(* IEC 61131-3 sources: plc-hackathon-2026/deliver/ME_v2_src, 24 files *)

(* ---- typeTeamAgg.st ---- *)
TYPE typeTeamAgg :
// Team energy [kWh] and cost [EUR] aggregate for one day, one month or the year.
// Names follow spec tables 12 (energies) and 4.3 (cost components). LREAL accumulators.
STRUCT
	E_fne : LREAL;                      // PV production after curtailment (FNE_P_act)
	E_fec : LREAL;                      // fixed consumption (FEC_P_fix remembered from k-1)
	E_bess_chg : LREAL;                 // battery charging, bus side
	E_bess_dch : LREAL;                 // battery discharging, bus side
	E_ev : LREAL;                       // all EV chargers, bus side
	E_ev_ch : ARRAY[0..3] OF LREAL;     // per EV charger, bus side
	E_import : LREAL;                   // grid import
	E_export : LREAL;                   // grid export
	P_peak : LREAL;                     // [kW] max 15-min import (monthly value; also kept per day for info)
	C_purchase : LREAL;                 // energy purchase = import * c_en
	C_revenue : LREAL;                  // export revenue = export * 0.9 * c_en
	C_grid : LREAL;                     // grid fee on import (VT/NT)
	C_peak : LREAL;                     // peak power cost (month/year only; 0 for days)
	C_total : LREAL;                    // purchase - revenue + grid (+ peak for month/year)
END_STRUCT
END_TYPE

(* ---- typeTeamAlarm.st ---- *)
TYPE typeTeamAlarm :
// One alarm/message history entry, stamped with SIMULATED time (no PLC clock).
STRUCT
	k : DINT;                           // simulation step when raised
	sStamp : STRING(20);                // simulated date/time "DD.MM.YYYY HH:MM"
	iCode : INT;                        // see Team_HMI alarm code list
	sText : STRING(80);                 // human readable message
END_STRUCT
END_TYPE

(* ---- Team_Cfg.st ---- *)
// Team_Cfg: team tuning constants (physics parameters are always read from SimParam).
VAR_GLOBAL CONSTANT
	N_STEPS : DINT := 35040;            // steps in the simulated year
	GRID_MARGIN_IMP : REAL := 1.0;      // [kW] safety margin below EGC_MAX_IMPORT for the predicted grid power
	GRID_MARGIN_EXP : REAL := 1.0;      // [kW] safety margin below EGC_MAX_EXPORT
	P_EPS : REAL := 0.001;              // [kW] below this a BESS setpoint is treated as zero
	// ---- forecast (FB_Forecast) ----
	FC_ALPHA_FEC : REAL := 0.5;         // EMA weight of the newest day for the load profile
	FC_ALPHA_PV : REAL := 0.3;          // EMA weight of the newest day for the PV profile
	FC_ALPHA_SIG : REAL := 0.3;         // EMA weight for the FEC deviation (sigma)
	FC_KSIG_TT : REAL := 1.0;           // two-tariff: pessimistic load = expected + FC_KSIG_TT * sigma
	FC_KSIG_DA : REAL := 0.0;           // day-ahead: same (arbitrage is worth more than the reserve)
	FC_CORR_W : INT := 4;               // intraday correction window [steps], 0 = off (max 16)
	FC_CORR_TAU : REAL := 16.0;         // fade-out of the intraday correction [steps]
	FC_CORR_FEC : BOOL := TRUE;         // apply intraday correction to FEC
	FC_CORR_PV : BOOL := TRUE;          // apply intraday correction to PV
	// ---- planner (FB_Planner) ----
	PLAN_H : INT := 96;                 // planning horizon [steps] (24 h)
	PLAN_DA_PUBLISHED : BOOL := TRUE;   // TRUE: day-ahead horizon limited to published prices (13:00 rule)
	PLAN_PEN : REAL := 20.0;            // [EUR/kW per step] penalty for planned import above the cap
	PLAN_TVF : REAL := 0.9;             // terminal value of stored energy = mean import price * PLAN_TVF
	PLAN_PVF : REAL := 0.6;             // PV share trusted when computing the peak cap
	PLAN_HI_TT : BOOL := TRUE;          // two-tariff: DP peak penalty uses the pessimistic net load
	PLAN_HI_DA : BOOL := FALSE;         // day-ahead: DP peak penalty uses the expected net load
	PLAN_TSPLIT : BOOL := FALSE;        // TRUE: free import level from the expected forecast (see FB_Planner)
	PLAN_CAPM : REAL := 1.02;           // safety factor on the computed peak cap
END_VAR

(* ---- Team_HMI.st ---- *)
// Team_HMI: everything the HMI needs that is not directly in SimIO/SimParam/SimCtrl.
// Written by FB_HmiUpdate (called from Team_Main). Only iSelDay / iSelMonth are written by the HMI.
// All times are SIMULATED time (derived from simOut.t_sim), never the PLC clock.
VAR_GLOBAL
	// ---- status / header (show on every screen) ----
	sDateTime : STRING(20);             // "DD.MM.YYYY HH:MM" start of current interval k
	k : DINT;                           // current step
	rProgressPct : REAL;                // 0..100 % of the year
	xTariffHigh : BOOL;                 // TRUE = VT (high tariff) in current interval
	sTariff : STRING(2);                // 'VT' / 'NT'
	sPriceMode : STRING(20);            // 'Dvotarifni (HEP)' / 'Dan-unaprijed'
	rPrice : REAL;                      // [EUR/kWh] energy price of the current interval
	rGridFee : REAL;                    // [EUR/kWh] grid fee of the current interval
	// ---- power flows: requested (simCmd, interval k) vs actual (*_act, interval k-1) [kW] ----
	rFneAvail : REAL;                   // available PV in interval k (before curtailment)
	rFneExpected : REAL;                // PV expected after our curtailment, interval k
	xCurtActive : BOOL;                 // curtailment enabled in interval k
	rCurtValue : REAL;                  // curtailment limit [kW]
	rFneAct : REAL;                     // actual PV, interval k-1
	rFec : REAL;                        // fixed consumption, interval k
	rFecPrev : REAL;                    // fixed consumption, interval k-1
	rBessReq : REAL;                    // requested battery power, + = discharge, - = charge
	rBessChgReq : REAL;                 // requested charge [kW] (0 if not charging)
	rBessDchReq : REAL;                 // requested discharge [kW]
	rBessAct : REAL;                    // actual battery power interval k-1, + = discharge
	rBessChgAct : REAL;
	rBessDchAct : REAL;
	aEvReq : ARRAY[0..3] OF REAL;       // requested EV power, interval k
	aEvAct : ARRAY[0..3] OF REAL;       // actual EV power, interval k-1
	rEvReqSum : REAL;
	rEvActSum : REAL;
	rGridPred : REAL;                   // predicted grid power interval k, + = import, - = export
	rImportAct : REAL;                  // measured import interval k-1
	rExportAct : REAL;                  // measured export interval k-1
	rGridPredErr : REAL;                // |prediction(k-1) - measurement(k-1)| [kW]
	rGridPredErrMax : REAL;             // max of the above since reset
	// ---- battery ----
	rSoc : REAL;                        // [%]
	rSocMin : REAL;                     // [%] safety limits (SimParam)
	rSocMax : REAL;
	sBessDir : STRING(12);              // 'PUNJENJE' / 'PRAZNJENJE' / 'MIROVANJE'
	// ---- EV chargers ----
	aEvConnected : ARRAY[0..3] OF BOOL;
	aEvDeparture : ARRAY[0..3] OF STRING(20);   // planned departure "DD.MM.YYYY HH:MM" ('' if not connected)
	aEvRemaining : ARRAY[0..3] OF REAL;         // [kWh] energy still required
	aEvDelivered : ARRAY[0..3] OF REAL;         // [kWh] delivered this session
	aEvStepsLeft : ARRAY[0..3] OF DINT;         // 15-min intervals until departure
	// ---- peak power ----
	rPeakMonth : REAL;                  // [kW] monthly import peak so far (current month)
	rPeakTarget : REAL;                 // [kW] import cap the controller currently aims for
	// ---- energy/cost tables: selection written by the HMI ----
	iSelDay : INT := 0;                 // 0..364 -> stSelDay
	iSelMonth : INT := 1;               // 1..12  -> stSelMonth, aSelMonthDays
	stSelDay : typeTeamAgg;
	stSelMonth : typeTeamAgg;
	aSelMonthDays : ARRAY[1..31] OF typeTeamAgg;   // days of the selected month (unused days = 0)
	iSelMonthDays : INT;                // number of days in the selected month
	// ---- 24 h trends: index 95 = newest interval (k-1), 0 = oldest ----
	aTrFne : ARRAY[0..95] OF REAL;      // PV actual [kW]
	aTrFec : ARRAY[0..95] OF REAL;      // fixed consumption [kW]
	aTrGrid : ARRAY[0..95] OF REAL;     // grid, + import / - export [kW]
	aTrBess : ARRAY[0..95] OF REAL;     // battery, + discharge / - charge [kW]
	aTrEv : ARRAY[0..95] OF REAL;       // EV total [kW]
	aTrSoc : ARRAY[0..95] OF REAL;      // SoC [%]
	aTrPrice : ARRAY[0..95] OF REAL;    // energy price [EUR/kWh]
	// ---- alarms ----
	xAlmImport : BOOL;                  // EGC_overload_import (previous step)
	xAlmExport : BOOL;                  // EGC_overload_export
	xAlmTripped : BOOL;                 // plant disconnected
	xAlmFinished : BOOL;                // year finished (message)
	xAlmEvUnmet : BOOL;                 // an EV left with undelivered energy (latched until reset)
	xAlmGuardEv : BOOL;                 // guard reduced EV charging to hold import limit (this step)
	xAlmGuardCurt : BOOL;               // guard curtailed PV to hold export limit (this step)
	xAlmGuardFail : BOOL;               // predicted import above limit even after all measures
	aAlarmHist : ARRAY[0..49] OF typeTeamAlarm;   // newest at index 0
	nAlarms : DINT;                     // number of messages since reset
	sLastAlarm : STRING(80);
	// ---- diagnostics ----
	nCalls : DINT;                      // Team_Main calls since PLC start
	nSteps : DINT;                      // new steps processed since reset
	nGuardEv : DINT;                    // steps with EV shedding
	nGuardCurt : DINT;                  // steps with export curtailment by the guard
	nGuardFail : DINT;                  // steps where the guard could not hold the import limit
	nBothEnables : DINT;                // must stay 0
	rEvUnmetSum : REAL;                 // [kWh] energy not delivered at departures (own estimate)
END_VAR

(* ---- Team_Log.st ---- *)
// Team_Log: daily and monthly energy/cost tables (spec 4.2/4.3). Index = simulated day / month of interval k-1.
VAR_GLOBAL
	aDay : ARRAY[0..364] OF typeTeamAgg;    // day_of_year 0..364 (C_peak = 0, C_total = purchase - revenue + grid)
	aMonth : ARRAY[1..12] OF typeTeamAgg;   // month 1..12 incl. peak power P_peak and C_peak
	stYear : typeTeamAgg;                   // yearly totals (copied to Team_Results)
END_VAR

(* ---- Team_Prices.st ---- *)
// Team_Prices: price lists (cjenici, spec 3.9/4.1) generated by tools/gen_prices.py from the organizer CSVs.
// Energy price only; grid fee and peak price come from SimParam. Not a simulator profile (FNE/FEC/EV are never embedded).
VAR_GLOBAL CONSTANT
	// Elektra two-tariff energy price [EUR/kWh] per calendar quarter (1 = Jan-Mar ... 4 = Oct-Dec)
	TT_NT : ARRAY[1..4] OF REAL := [0.09, 0.1051, 0.0934, 0.0949];
	TT_VT : ARRAY[1..4] OF REAL := [0.1531, 0.1786, 0.1588, 0.1613];
END_VAR
VAR_GLOBAL
	// Day-ahead energy price [EUR/kWh] per 15-min interval k = 0..35039 (ENTSO-E HR 2025, may be negative)
	aDA : ARRAY[0..35039] OF REAL := [
		4(0.1353348), 4(0.143694), 4(0.1349352), 4(0.1010124), 4(0.0687852), 4(0.1011852), 4(0.0974808), 4(0.0902556), 4(0.0399492), 4(0.0485892), 4(0.04158), 4(0.0430056),
		4(0.04347), 4(0.059886), 4(0.0664632), 4(0.0900288), 4(0.1161648), 4(0.1328832), 4(0.1382724), 4(0.1446984), 4(0.1406268), 4(0.1307124), 4(0.1310364), 4(0.0904176),
		4(0.0689904), 4(0.0865296), 4(0.0846936), 4(0.053136), 4(0.0614844), 4(0.0834732), 4(0.1200204), 4(0.1431324), 4(0.1405836), 4(0.1433268), 4(0.1391148), 4(0.1337364),
		4(0.1330668), 4(0.126144), 4(0.135), 4(0.1405188), 4(0.1650456), 4(0.1762452), 4(0.1695492), 4(0.1646028), 4(0.1414152), 4(0.134622), 4(0.1270188), 4(0.1095228),
		4(0.111996), 4(0.1023732), 4(0.0968436), 4(0.0945216), 4(0.0923832), 4(0.0993816), 4(0.1185516), 4(0.1469556), 4(0.1492452), 4(0.1461564), 4(0.1350216), 4(0.1219968),
		4(0.1201716), 4(0.118206), 4(0.124956), 4(0.1402596), 4(0.1587276), 4(0.1571508), 4(0.1572696), 4(0.1564488), 4(0.1478196), 4(0.1314684), 4(0.1361988), 4(0.1318572),
		4(0.1189296), 4(0.1130112), 4(0.1087344), 4(0.1065204), 4(0.1077732), 4(0.113454), 4(0.12096), 4(0.1352808), 4(0.1386612), 4(0.14121), 4(0.1407672), 4(0.1385532),
		4(0.1404324), 4(0.140238), 4(0.147312), 4(0.15309), 4(0.1819368), 4(0.1857924), 4(0.1848096), 4(0.1831572), 4(0.1590624), 4(0.151524), 4(0.1455192), 4(0.1259604),
		4(0.1211004), 4(0.107838), 4(0.1033668), 4(0.1013364), 4(0.1006992), 4(0.0971892), 4(0.0989064), 4(0.1068012), 4(0.105408), 4(0.1070172), 4(0.103194), 4(0.1084104),
		4(0.1057752), 4(0.1129248), 4(0.122094), 4(0.1337364), 4(0.1717308), 4(0.165024), 4(0.1562328), 4(0.1627236), 4(0.1535328), 4(0.1449144), 4(0.1105056), 4(0.0771984),
		4(0.1130004), 4(0.0960336), 4(0.0743256), 4(0.0708804), 4(0.070794), 4(0.0962172), 4(0.1229364), 4(0.1331748), 4(0.1334664), 4(0.1152576), 4(0.097956), 4(0.0780624),
		4(0.0841212), 4(0.10476), 4(0.1249668), 4(0.1229904), 4(0.1472904), 4(0.1600344), 4(0.1528524), 4(0.1521828), 4(0.1456272), 4(0.122364), 4(0.1168128), 4(0.0853416),
		4(0.0343116), 4(0.056538), 4(0.0510192), 4(0.0135), 4(0.0662688), 4(0.0844668), 4(0.1362636), 4(0.16443), 4(0.148014), 4(0.1423224), 4(0.1318248), 4(0.131274),
		4(0.1322676), 4(0.1404432), 4(0.1504656), 4(0.1588572), 4(0.1668384), 4(0.166806), 4(0.1628424), 4(0.1643328), 4(0.1532088), 4(0.1370196), 4(0.125064), 4(0.1204416),
		4(0.0901584), 4(0.0813672), 4(0.0789048), 4(0.0747036), 4(0.0923076), 4(0.11178), 4(0.1367388), 4(0.1635336), 4(0.1611252), 4(0.1341576), 4(0.1174068), 4(0.1103436),
		4(0.1120824), 4(0.1245996), 4(0.1353132), 4(0.1550556), 4(0.1646784), 4(0.165456), 4(0.1622916), 4(0.1614384), 4(0.1484352), 4(0.1356372), 4(0.1255716), 4(0.114588),
		4(0.1147284), 4(0.114588), 4(0.1119096), 4(0.1104408), 4(0.1152468), 4(0.1184868), 4(0.1342656), 4(0.1542132), 4(0.1678104), 4(0.1601208), 4(0.1514916), 4(0.1435644),
		4(0.1331532), 4(0.1284012), 4(0.1325484), 4(0.1425708), 4(0.1583496), 4(0.1566756), 4(0.16065), 4(0.1521612), 4(0.1421172), 4(0.1240056), 4(0.11151), 4(0.0968328),
		4(0.0941976), 4(0.0868104), 4(0.0826092), 4(0.0808164), 4(0.0767664), 4(0.1046088), 4(0.1354968), 4(0.165024), 4(0.1680264), 4(0.1522368), 4(0.1334556), 4(0.1226772),
		4(0.1160244), 4(0.1134108), 4(0.1188108), 4(0.1389852), 4(0.1609308), 4(0.1583604), 4(0.1590084), 4(0.1569024), 4(0.1457568), 4(0.1323108), 4(0.129492), 4(0.1226016),
		4(0.1179468), 4(0.1079676), 4(0.1042632), 4(0.1000296), 4(0.099144), 4(0.1006236), 4(0.1021788), 4(0.1209168), 4(0.12312), 4(0.1200744), 4(0.113454), 4(0.1078488),
		4(0.1046088), 4(0.100602), 4(0.1068768), 4(0.113994), 4(0.1448928), 4(0.1509732), 4(0.1472256), 4(0.148284), 4(0.1366848), 4(0.1265328), 4(0.11799), 4(0.1143612),
		4(0.1075896), 4(0.0961416), 4(0.0964548), 4(0.092178), 4(0.0918), 4(0.0919188), 4(0.0946836), 4(0.10989), 4(0.1258092), 4(0.1296756), 4(0.1271916), 4(0.1140588),
		4(0.1112292), 4(0.1075788), 4(0.1139616), 4(0.1299564), 4(0.1461024), 4(0.1542564), 4(0.1583928), 4(0.1557468), 4(0.1468152), 4(0.1380348), 4(0.1312956), 4(0.124092),
		4(0.1213812), 4(0.1134756), 4(0.1128168), 4(0.1083996), 4(0.108), 4(0.1190052), 4(0.1512108), 4(0.1927476), 4(0.2371032), 4(0.1868184), 4(0.15201), 4(0.1311444),
		4(0.1245456), 4(0.1297512), 4(0.1363284), 4(0.1529928), 4(0.1704564), 4(0.1678212), 4(0.16902), 4(0.1670976), 4(0.1538244), 4(0.1375164), 4(0.1288008), 4(0.1167588),
		4(0.1186812), 4(0.115344), 4(0.1107), 4(0.1092312), 4(0.1125036), 4(0.1180332), 4(0.1495908), 4(0.1742688), 4(0.2001672), 4(0.16416), 4(0.141156), 4(0.1340712),
		4(0.1289304), 4(0.1293084), 4(0.1439532), 4(0.1770552), 4(0.1979964), 4(0.2446632), 4(0.239652), 4(0.211572), 4(0.187164), 4(0.172746), 4(0.1610172), 4(0.1348812),
		4(0.127656), 4(0.1213488), 4(0.1200528), 4(0.1174932), 4(0.1255068), 4(0.1390392), 4(0.1600992), 4(0.2120148), 4(0.3359124), 4(0.338904), 4(0.3266568), 4(0.325566),
		4(0.31023), 4(0.306774), 4(0.3062448), 4(0.3319596), 4(0.326268), 4(0.368226), 4(0.320328), 4(0.265248), 4(0.1937088), 4(0.1670328), 4(0.1554768), 4(0.133812),
		4(0.136296), 4(0.131868), 4(0.1281636), 4(0.1259928), 4(0.1292652), 4(0.1392012), 4(0.1701216), 4(0.2121984), 4(0.2210544), 4(0.189), 4(0.164052), 4(0.1518912),
		4(0.1456488), 4(0.1492344), 4(0.1566), 4(0.1827144), 4(0.19683), 4(0.2082348), 4(0.1990656), 4(0.1943676), 4(0.172368), 4(0.1623996), 4(0.1519992), 4(0.1398276),
		4(0.1364364), 4(0.1331208), 4(0.1297836), 4(0.1277532), 4(0.1277964), 4(0.1346328), 4(0.152064), 4(0.1890108), 4(0.2247804), 4(0.1893672), 4(0.1700352), 4(0.1518696),
		4(0.1365552), 4(0.1339524), 4(0.1444284), 4(0.1637172), 4(0.1839888), 4(0.1930284), 4(0.1943136), 4(0.1881576), 4(0.1705428), 4(0.1566), 4(0.1511676), 4(0.1383588),
		4(0.1363392), 4(0.1309284), 4(0.1311336), 4(0.128412), 4(0.1263816), 4(0.1294164), 4(0.1325592), 4(0.1465776), 4(0.157626), 4(0.155628), 4(0.1445796), 4(0.1315224),
		4(0.1283796), 4(0.1242108), 4(0.129168), 4(0.149094), 4(0.1772712), 4(0.1826928), 4(0.1809756), 4(0.181278), 4(0.1686096), 4(0.1548936), 4(0.147312), 4(0.1397088),
		4(0.1403028), 4(0.1350108), 4(0.1336068), 4(0.1309392), 4(0.1297944), 4(0.1296), 4(0.1314252), 4(0.1340172), 4(0.1335636), 4(0.136188), 4(0.1366092), 4(0.1341252),
		4(0.12123), 4(0.1161108), 4(0.1261548), 4(0.1377324), 4(0.1627344), 4(0.1759428), 4(0.180522), 4(0.1794096), 4(0.1741608), 4(0.1651644), 4(0.145044), 4(0.133866),
		4(0.1322784), 4(0.1294056), 4(0.1259388), 4(0.1235628), 4(0.124686), 4(0.1404216), 4(0.1766232), 4(0.3070548), 4(0.4670028), 4(0.3149496), 4(0.2551932), 4(0.2076084),
		4(0.193266), 4(0.1851012), 4(0.2071332), 4(0.2981016), 4(0.446472), 4(0.6208812), 4(0.5111424), 4(0.3192156), 4(0.2376), 4(0.1836), 4(0.1718928), 4(0.1540944),
		4(0.1477764), 4(0.1417932), 4(0.134622), 4(0.1350972), 4(0.1429056), 4(0.16416), 4(0.207414), 4(0.3141612), 4(0.4177224), 4(0.2861676), 4(0.2540484), 4(0.2179224),
		4(0.2129004), 4(0.1951344), 4(0.2188512), 4(0.3057588), 4(0.245214), 4(0.3387744), 4(0.2779704), 4(0.2207844), 4(0.190728), 4(0.1687392), 4(0.153684), 4(0.144234),
		4(0.141588), 4(0.1360152), 4(0.1345896), 4(0.1350972), 4(0.1372464), 4(0.1506816), 4(0.20925), 4(0.3410964), 4(0.2672136), 4(0.2153628), 4(0.1933848), 4(0.1867752),
		4(0.1782), 4(0.1836), 4(0.1943136), 4(0.2137752), 4(0.2703888), 4(0.276102), 4(0.2261952), 4(0.222642), 4(0.2220156), 4(0.1710072), 4(0.1589436), 4(0.145854),
		4(0.1353888), 4(0.1299564), 4(0.119394), 4(0.1175796), 4(0.1227096), 4(0.1344708), 4(0.1809864), 4(0.2092608), 4(0.1881684), 4(0.1808568), 4(0.1625292), 4(0.1594728),
		4(0.1543104), 4(0.1588032), 4(0.1690416), 4(0.1919376), 4(0.2108916), 4(0.2148012), 4(0.2028672), 4(0.1957824), 4(0.2018628), 4(0.1633608), 4(0.1606176), 4(0.136188),
		4(0.127656), 4(0.1162512), 4(0.1107), 4(0.1093392), 4(0.1170288), 4(0.1424304), 4(0.17469), 4(0.1909872), 4(0.1764828), 4(0.1599048), 4(0.1535652), 4(0.1422576),
		4(0.1392444), 4(0.13662), 4(0.1417716), 4(0.161892), 4(0.1961064), 4(0.1983744), 4(0.1922616), 4(0.1883412), 4(0.1774872), 4(0.1666008), 4(0.1547208), 4(0.1429488),
		4(0.1203336), 4(0.1117476), 4(0.0980856), 4(0.094878), 4(0.0971136), 4(0.1055808), 4(0.1218564), 4(0.1337904), 4(0.1181628), 4(0.1153224), 4(0.1033776), 4(0.0975888),
		4(0.09396), 4(0.0924372), 4(0.1067256), 4(0.1288872), 4(0.1661148), 4(0.1701108), 4(0.1716444), 4(0.1709208), 4(0.162864), 4(0.155574), 4(0.1481004), 4(0.135),
		4(0.1419552), 4(0.1297404), 4(0.1272888), 4(0.1204524), 4(0.12096), 4(0.1231524), 4(0.1255176), 4(0.1334664), 4(0.1427112), 4(0.1400004), 4(0.1207656), 4(0.112752),
		4(0.1054188), 4(0.1028808), 4(0.1209168), 4(0.13095), 4(0.1467288), 4(0.1559088), 4(0.1424628), 4(0.1443312), 4(0.1348812), 4(0.1245888), 4(0.104004), 4(0.08397),
		4(0.0654696), 4(0.0605124), 4(0.0433404), 4(0.032022), 4(0.0490536), 4(0.118098), 4(0.1559088), 4(0.187002), 4(0.1719684), 4(0.1409616), 4(0.1084428), 4(0.1040148),
		4(0.0946944), 4(0.1125792), 4(0.1399464), 4(0.1582416), 4(0.1937628), 4(0.1899936), 4(0.1928124), 4(0.1906308), 4(0.170856), 4(0.1461024), 4(0.130626), 4(0.106056),
		4(0.106758), 4(0.0855684), 4(0.0941112), 4(0.0877068), 4(0.0877392), 4(0.122688), 4(0.1498608), 4(0.1502712), 4(0.1519992), 4(0.1354212), 4(0.141318), 4(0.1357344),
		4(0.1322892), 4(0.1372788), 4(0.1420632), 4(0.135162), 4(0.1540296), 4(0.1559304), 4(0.1593864), 4(0.1502928), 4(0.1499256), 4(0.1251612), 4(0.1250208), 4(0.1051704),
		4(0.105462), 4(0.097362), 4(0.0910332), 4(0.0914328), 4(0.0972), 4(0.1214676), 4(0.154656), 4(0.1773468), 4(0.1579068), 4(0.1480896), 4(0.1204308), 4(0.1014444),
		4(0.093204), 4(0.0935496), 4(0.1055484), 4(0.1400328), 4(0.1792692), 4(0.1827792), 4(0.1721088), 4(0.173502), 4(0.1609524), 4(0.1491912), 4(0.1330236), 4(0.1119204),
		4(0.110268), 4(0.1095228), 4(0.1069524), 4(0.1100844), 4(0.1098036), 4(0.1232496), 4(0.1569348), 4(0.1669788), 4(0.173124), 4(0.1639764), 4(0.1429704), 4(0.13311),
		4(0.1219428), 4(0.122364), 4(0.1403892), 4(0.1655748), 4(0.1736748), 4(0.1896696), 4(0.1858032), 4(0.1741824), 4(0.1635228), 4(0.145908), 4(0.1370952), 4(0.129816),
		4(0.1296), 4(0.1269), 4(0.1232064), 4(0.1236384), 4(0.1267164), 4(0.1316088), 4(0.1604556), 4(0.1728), 4(0.176796), 4(0.1672056), 4(0.140508), 4(0.136296),
		4(0.1296648), 4(0.1308852), 4(0.1296432), 4(0.1655964), 4(0.1810512), 4(0.1930716), 4(0.1992384), 4(0.1933092), 4(0.1756728), 4(0.164916), 4(0.1607472), 4(0.144126),
		4(0.1494828), 4(0.1409724), 4(0.135108), 4(0.1288332), 4(0.1295568), 4(0.1312308), 4(0.1374948), 4(0.1563192), 4(0.1657368), 4(0.1538352), 4(0.138672), 4(0.1296864),
		4(0.1191132), 4(0.111672), 4(0.122796), 4(0.1411344), 4(0.1683072), 4(0.1792368), 4(0.180036), 4(0.1760184), 4(0.169128), 4(0.1568592), 4(0.1530684), 4(0.1422792),
		4(0.1439208), 4(0.1370628), 4(0.1328292), 4(0.1303128), 4(0.1321272), 4(0.1332828), 4(0.1383372), 4(0.146772), 4(0.148284), 4(0.148716), 4(0.1404432), 4(0.1396764),
		4(0.1320192), 4(0.1208304), 4(0.1263168), 4(0.140562), 4(0.168156), 4(0.1802088), 4(0.185544), 4(0.187866), 4(0.17874), 4(0.1682316), 4(0.1603152), 4(0.1438992),
		4(0.1399032), 4(0.1367604), 4(0.1346976), 4(0.1296432), 4(0.1330992), 4(0.1379916), 4(0.1719144), 4(0.2245104), 4(0.2626884), 4(0.1922832), 4(0.161946), 4(0.1363176),
		4(0.1266516), 4(0.1249776), 4(0.1344276), 4(0.1597968), 4(0.1793664), 4(0.226962), 4(0.2167884), 4(0.217188), 4(0.1811592), 4(0.16524), 4(0.1557252), 4(0.1466748),
		4(0.142992), 4(0.1355832), 4(0.1330344), 4(0.1339092), 4(0.13311), 4(0.1378404), 4(0.1674432), 4(0.2056644), 4(0.2289492), 4(0.1763748), 4(0.1474524), 4(0.1369656),
		4(0.127602), 4(0.1222452), 4(0.1296972), 4(0.1542456), 4(0.181332), 4(0.189324), 4(0.189), 4(0.1863648), 4(0.1727352), 4(0.1464804), 4(0.1424412), 4(0.1347624),
		4(0.1260036), 4(0.1207548), 4(0.1198584), 4(0.1186056), 4(0.1248912), 4(0.1323648), 4(0.1636524), 4(0.1825092), 4(0.1952748), 4(0.1720764), 4(0.145476), 4(0.133704),
		4(0.127926), 4(0.1297512), 4(0.139158), 4(0.1556496), 4(0.1719252), 4(0.19116), 4(0.205092), 4(0.2048004), 4(0.1836), 4(0.1678536), 4(0.155196), 4(0.144774),
		4(0.1443636), 4(0.1403892), 4(0.13608), 4(0.135), 4(0.1350108), 4(0.1447524), 4(0.165996), 4(0.1944972), 4(0.2356128), 4(0.1930932), 4(0.1686204), 4(0.1617408),
		4(0.1561032), 4(0.1526148), 4(0.1520208), 4(0.1622808), 4(0.181656), 4(0.188244), 4(0.1913544), 4(0.1864512), 4(0.1768068), 4(0.159624), 4(0.1512108), 4(0.131706),
		4(0.136134), 4(0.121716), 4(0.1175256), 4(0.1134), 4(0.1185192), 4(0.1280772), 4(0.1678104), 4(0.1848744), 4(0.1782324), 4(0.1625076), 4(0.1456812), 4(0.1280556),
		4(0.1243512), 4(0.1240164), 4(0.12744), 4(0.1442556), 4(0.1857924), 4(0.1894644), 4(0.1884924), 4(0.1860624), 4(0.1818072), 4(0.1557576), 4(0.1285632), 4(0.1209816),
		4(0.09828), 4(0.0950184), 4(0.0937872), 4(0.09612), 4(0.0968652), 4(0.0982692), 4(0.1052028), 4(0.1174068), 4(0.1222128), 4(0.109134), 4(0.1035072), 4(0.0960336),
		4(0.0954828), 4(0.097686), 4(0.1025244), 4(0.12744), 4(0.16173), 4(0.1752948), 4(0.1733832), 4(0.1713852), 4(0.1661472), 4(0.16092), 4(0.1542564), 4(0.1449792),
		4(0.1458), 4(0.136404), 4(0.1319004), 4(0.128844), 4(0.1261656), 8(0.12636), 4(0.1441044), 4(0.1477116), 4(0.1321812), 4(0.1230876), 4(0.1191456), 4(0.1106028),
		4(0.1090368), 4(0.118692), 4(0.130032), 4(0.1627992), 4(0.1736856), 4(0.1889784), 4(0.1888164), 4(0.1786968), 4(0.1560816), 4(0.15444), 4(0.139482), 4(0.1297944),
		4(0.1247292), 4(0.1217916), 4(0.1173096), 4(0.1168992), 4(0.126576), 4(0.1724004), 4(0.1935684), 4(0.1958688), 4(0.1762344), 4(0.1672488), 4(0.1512108), 4(0.136512),
		4(0.132732), 4(0.142398), 4(0.179712), 4(0.2052972), 4(0.218322), 4(0.2210112), 4(0.2083752), 4(0.2056644), 4(0.1809), 4(0.1751544), 4(0.1435428), 4(0.1483812),
		4(0.1365768), 4(0.1335204), 4(0.1290384), 4(0.1365876), 4(0.1763856), 4(0.1951884), 4(0.2572236), 4(0.1924884), 4(0.15687), 4(0.13068), 4(0.1269432), 4(0.1278612),
		4(0.1289304), 4(0.1395684), 4(0.1727136), 4(0.200016), 4(0.2052), 4(0.2388312), 4(0.2170044), 4(0.1934064), 4(0.1859868), 4(0.1727892), 4(0.1431432), 4(0.1397952),
		4(0.1380996), 4(0.1369656), 4(0.1367172), 4(0.1390392), 4(0.1469772), 4(0.1866024), 4(0.1955232), 4(0.1944), 4(0.1889136), 4(0.1791612), 4(0.171234), 4(0.16119),
		4(0.1638144), 4(0.1802196), 4(0.1956852), 4(0.2190564), 4(0.3030804), 4(0.2873556), 4(0.240462), 4(0.2384316), 4(0.1923156), 4(0.1861812), 4(0.1728), 4(0.1722708),
		4(0.161298), 4(0.158868), 4(0.1538136), 4(0.1591596), 4(0.1767852), 4(0.2259684), 4(0.421524), 4(0.3348108), 4(0.2808108), 4(0.2247588), 4(0.2027268), 4(0.2015604),
		4(0.2252664), 4(0.2457648), 4(0.2673), 4(0.2891484), 4(0.2678184), 4(0.2236788), 4(0.2122416), 4(0.1927152), 4(0.1759536), 4(0.1653696), 4(0.1503036), 4(0.1514376),
		4(0.1460916), 4(0.141048), 4(0.1412748), 4(0.141858), 4(0.1520748), 4(0.1772712), 4(0.2337336), 4(0.2835216), 4(0.229284), 4(0.1935144), 4(0.1778976), 4(0.1623564),
		4(0.1625508), 4(0.1714824), 4(0.1871316), 4(0.2142396), 4(0.3135456), 4(0.3104244), 4(0.2420388), 4(0.198234), 4(0.1766232), 4(0.16524), 4(0.1512324), 4(0.1472688),
		4(0.1418796), 4(0.1303884), 4(0.1291356), 4(0.1295784), 4(0.1315872), 4(0.146718), 4(0.1623888), 4(0.1616328), 4(0.148068), 4(0.1345572), 4(0.1278288), 4(0.1213812),
		4(0.1188108), 4(0.126252), 4(0.1413936), 4(0.1687716), 4(0.1905552), 4(0.1925856), 4(0.1880064), 4(0.1818504), 4(0.165348), 4(0.1515672), 4(0.1441692), 4(0.1448388),
		4(0.139212), 4(0.1334556), 4(0.129492), 4(0.1291356), 4(0.1305612), 4(0.133758), 4(0.1448712), 4(0.153846), 4(0.152334), 4(0.1427652), 4(0.141696), 4(0.1389636),
		4(0.1375812), 4(0.14094), 4(0.1524744), 4(0.174852), 4(0.1890324), 4(0.191322), 4(0.1876932), 4(0.1830708), 4(0.1726272), 4(0.1613412), 4(0.1420308), 4(0.1431216),
		4(0.1307448), 4(0.1299672), 4(0.1365876), 4(0.1406052), 4(0.1550124), 4(0.1884924), 4(0.2253096), 4(0.2265732), 4(0.185004), 4(0.1508436), 4(0.1288764), 4(0.1232928),
		4(0.1176012), 4(0.13176), 4(0.1601748), 4(0.1869372), 4(0.238572), 4(0.2883816), 4(0.2338956), 4(0.1934928), 4(0.1759212), 4(0.169074), 4(0.15444), 4(0.146664),
		4(0.1429488), 4(0.1358748), 4(0.1331316), 4(0.1377216), 4(0.163998), 4(0.2263032), 4(0.3576096), 4(0.209304), 4(0.1750356), 4(0.154386), 4(0.1445148), 4(0.142398),
		4(0.1559736), 4(0.1631448), 4(0.1770876), 4(0.3453516), 4(0.2810268), 4(0.2770092), 4(0.2601612), 4(0.1939248), 4(0.1817316), 4(0.1740852), 4(0.1480032), 4(0.14121),
		4(0.1392768), 4(0.1372896), 4(0.136458), 4(0.1398168), 4(0.155088), 4(0.1828872), 4(0.218592), 4(0.190404), 4(0.165456), 4(0.123606), 4(0.1240056), 4(0.1162728),
		4(0.1160568), 4(0.126954), 4(0.1515888), 4(0.190944), 4(0.249534), 4(0.2520504), 4(0.2164968), 4(0.1938492), 4(0.1805868), 4(0.1764936), 4(0.1671192), 4(0.1350972),
		4(0.1303452), 4(0.1251936), 4(0.1203984), 4(0.1305396), 4(0.1563948), 4(0.2001456), 4(0.263412), 4(0.19062), 4(0.1302804), 4(0.1142748), 4(0.0986364), 4(0.1005588),
		4(0.1060236), 4(0.1154952), 4(0.153846), 4(0.1964844), 4(0.2781972), 4(0.3032856), 4(0.2709936), 4(0.187596), 4(0.176904), 4(0.1739556), 4(0.1439748), 4(0.1269432),
		4(0.1223964), 4(0.1204956), 4(0.1224288), 4(0.1231308), 4(0.1458), 4(0.1756512), 4(0.188244), 4(0.1582416), 4(0.1398276), 4(0.1123524), 4(0.0950508), 4(0.0867564),
		4(0.0860436), 4(0.107892), 4(0.1171476), 4(0.1718604), 4(0.2034612), 4(0.2067012), 4(0.2070792), 4(0.1797876), 4(0.1654884), 4(0.145422), 4(0.1260468), 4(0.13203),
		4(0.1259496), 4(0.1227312), 4(0.1168668), 4(0.1191024), 4(0.1260468), 4(0.151794), 4(0.1414152), 4(0.1065204), 4(0.0763344), 4(0.0634392), 4(0.0612036), 4(0.0569916),
		4(0.0606852), 4(0.0737316), 4(0.128358), 4(0.1802304), 4(0.2145528), 4(0.1995408), 4(0.2117664), 4(0.1919808), 4(0.1703268), 4(0.1657152), 4(0.1615464), 4(0.1378512),
		4(0.138294), 4(0.1283796), 4(0.1277748), 4(0.128736), 4(0.1349352), 4(0.1454112), 4(0.1423332), 4(0.1270296), 4(0.1109592), 4(0.0945432), 4(0.0962172), 4(0.0814752),
		4(0.080838), 4(0.1136808), 4(0.1515996), 4(0.20547), 4(0.2142504), 4(0.2108916), 4(0.2121984), 4(0.1816344), 4(0.1752408), 4(0.1579716), 4(0.1437696), 4(0.1412748),
		4(0.1266408), 4(0.1217808), 4(0.1202796), 4(0.12393), 4(0.1646784), 4(0.2244888), 4(0.2619324), 4(0.1898856), 4(0.17928), 4(0.1571292), 4(0.1439964), 4(0.1381104),
		4(0.1377216), 4(0.1576908), 4(0.2053944), 4(0.2542212), 4(0.3007044), 4(0.3385584), 4(0.314172), 4(0.2235384), 4(0.1914516), 4(0.1759428), 4(0.1442664), 4(0.154332),
		4(0.139428), 4(0.1344168), 4(0.1337688), 4(0.1378404), 4(0.1590192), 4(0.2322324), 4(0.2833596), 4(0.1877148), 4(0.1683828), 4(0.1544076), 4(0.139374), 4(0.1379268),
		4(0.140346), 4(0.1505088), 4(0.1666008), 4(0.2288196), 4(0.3069468), 4(0.3333636), 4(0.2880468), 4(0.2162916), 4(0.1727892), 4(0.1578528), 4(0.1416744), 4(0.1348488),
		4(0.1326132), 4(0.1286388), 4(0.1282284), 4(0.1286172), 4(0.1369332), 4(0.1886328), 4(0.2148444), 4(0.1917864), 4(0.1698516), 4(0.1571292), 4(0.1430892), 4(0.13122),
		4(0.1323864), 4(0.1405836), 4(0.1608552), 4(0.1918404), 4(0.2159892), 4(0.2162052), 4(0.1993896), 4(0.1851768), 4(0.1579716), 4(0.1453248), 4(0.129816), 4(0.1205928),
		4(0.1121148), 4(0.1109268), 8(0.1096308), 4(0.1193508), 4(0.158328), 4(0.1742148), 4(0.1794096), 4(0.1623456), 4(0.1463184), 4(0.1380024), 4(0.130626), 4(0.1261872),
		4(0.1297512), 4(0.1470096), 4(0.181764), 4(0.1843668), 4(0.1918836), 4(0.1853712), 4(0.1789992), 4(0.1529928), 4(0.1429056), 4(0.1239732), 4(0.1306044), 4(0.1193832),
		4(0.1181304), 4(0.1156464), 4(0.1216944), 4(0.13392), 4(0.1674648), 4(0.1978236), 4(0.1741608), 4(0.1593324), 4(0.1399248), 4(0.1272024), 4(0.1191888), 4(0.1188972),
		4(0.1216944), 4(0.1370952), 4(0.1721628), 4(0.2049408), 4(0.2110428), 4(0.2149308), 4(0.1967652), 4(0.1700352), 4(0.1497528), 4(0.134946), 4(0.1395468), 4(0.130464),
		4(0.1266948), 4(0.1222884), 4(0.1193616), 4(0.1248264), 4(0.1381212), 4(0.1493208), 4(0.1511892), 4(0.1508868), 4(0.138024), 4(0.12393), 4(0.1121904), 4(0.1080648),
		4(0.1125252), 4(0.1363068), 4(0.1677024), 4(0.21735), 4(0.2160972), 4(0.2048868), 4(0.173556), 4(0.1505412), 4(0.1351188), 4(0.1295136), 4(0.1363176), 4(0.1292436),
		4(0.1137132), 4(0.113724), 4(0.1215432), 4(0.1246428), 4(0.1444932), 4(0.1420956), 4(0.120906), 4(0.09612), 4(0.073764), 4(0.05292), 4(0.0297), 4(0.019008),
		4(0.0572184), 4(0.0780732), 4(0.1435644), 4(0.1693332), 4(0.176526), 4(0.1771632), 4(0.1706292), 4(0.1626372), 4(0.1358316), 4(0.1227204), 4(0.1238328), 4(0.1172664),
		4(0.115668), 4(0.1113588), 4(0.1151604), 4(0.1288332), 4(0.1513188), 4(0.17604), 4(0.1595484), 4(0.1176444), 4(0.0878364), 4(0.084618), 4(0.091476), 4(0.0626184),
		4(0.0921672), 4(0.1216296), 4(0.152766), 4(0.1925964), 4(0.2588436), 4(0.2024784), 4(0.1784916), 4(0.1745604), 4(0.1605204), 4(0.1555308), 4(0.1387368), 4(0.1302264),
		4(0.1188756), 4(0.1167696), 4(0.1265112), 4(0.1686852), 4(0.1939896), 4(0.1906956), 4(0.153306), 4(0.1248804), 4(0.103302), 4(0.1115964), 4(0.039798), 4(0.0315252),
		4(0.0721656), 4(0.1109484), 4(0.1677996), 4(0.2093148), 4(0.2734452), 4(0.215298), 4(0.1860192), 4(0.1675188), 4(0.1552824), 4(0.1442556), 4(0.1448064), 4(0.1312524),
		4(0.1238328), 4(0.118854), 4(0.1313712), 4(0.1473228), 4(0.18387), 4(0.163944), 4(0.1172124), 4(0.0805248), 4(0.0244836), 4(0.0119124), 4(0.0075924), 4(0.0011232),
		4(0.0041688), 4(0.0786888), 4(0.134892), 4(0.1743768), 4(0.228744), 4(0.1930392), 4(0.1734264), 4(0.1610604), 4(0.1397736), 4(0.1315116), 4(0.1128816), 4(0.1133676),
		4(0.1125792), 4(0.1146852), 4(0.1219968), 4(0.1468692), 4(0.1857276), 4(0.1662336), 4(0.11718), 4(0.086076), 4(0.0622944), 4(0.0057564), 4(0.0016632), 4(0.0007776),
		4(0.0142128), 4(0.0805788), 4(0.1324512), 4(0.2071116), 4(0.237006), 4(0.2223612), 4(0.1900692), 4(0.1577772), 4(0.1492776), 4(0.1302912), 4(0.1153116), 4(0.1140264),
		4(0.10854), 4(0.1099656), 4(0.114048), 4(0.1347624), 4(0.164322), 4(0.1642896), 4(0.1339956), 4(0.0899316), 4(0.071064), 4(0.0343548), 4(0.0138132), 4(0.0086508),
		4(0.0415476), 4(0.1037232), 4(0.1464804), 4(0.1729836), 4(0.2413584), 4(0.208764), 4(0.175068), 4(0.151524), 4(0.140994), 4(0.1352808), 4(0.1441908), 4(0.13662),
		4(0.1405512), 4(0.137808), 4(0.1404756), 4(0.1484568), 4(0.146016), 4(0.1347948), 4(0.1058832), 4(0.0783432), 4(0.019494), 4(0.00243), 4(0.000864), 4(4.32E-05),
		4(7.56E-05), 4(0.0650916), 4(0.1236708), 4(0.1769364), 4(0.2254716), 4(0.2034612), 4(0.166914), 4(0.154116), 4(0.1454112), 4(0.1249884), 4(0.1188108), 4(0.115452),
		4(0.1132056), 4(0.1155276), 4(0.1188864), 4(0.121716), 4(0.1188324), 4(0.106218), 4(0.0736344), 4(0.0316116), 4(0.010908), 4(0.0016416), 4(0.000702), 4(-0.0003456),
		4(0.0007884), 4(0.0187812), 4(0.1079352), 4(0.149796), 4(0.1598832), 4(0.158166), 4(0.148824), 4(0.1400328), 4(0.125334), 4(0.119502), 4(0.10692), 4(0.105948),
		4(0.1073304), 4(0.1075032), 4(0.107838), 4(0.1214136), 4(0.1614492), 4(0.1707372), 4(0.144612), 4(0.1070604), 4(0.0843588), 4(0.0798876), 4(0.0821016), 4(0.0835056),
		4(0.0917568), 4(0.1085508), 4(0.1429704), 4(0.1568592), 4(0.1869804), 4(0.171828), 4(0.1521828), 4(0.1384992), 4(0.1163376), 4(0.1065528), 4(0.114426), 4(0.1117476),
		4(0.1086804), 4(0.1099332), 4(0.1132272), 4(0.1220832), 4(0.1521828), 4(0.1583064), 4(0.1551744), 4(0.1403568), 4(0.1103544), 4(0.1058724), 4(0.1052568), 4(0.1080432),
		4(0.1128168), 4(0.1251504), 4(0.1503792), 4(0.1712016), 4(0.205632), 4(0.1912248), 4(0.1594512), 4(0.1449036), 4(0.1326996), 4(0.1161864), 4(0.1102356), 4(0.1087776),
		4(0.1059912), 4(0.1063044), 4(0.1118664), 4(0.122418), 4(0.1487052), 4(0.1657152), 4(0.1566972), 4(0.135), 4(0.110376), 4(0.1075248), 4(0.1059048), 4(0.1074924),
		4(0.1098576), 4(0.1288764), 4(0.1465776), 4(0.1611252), 4(0.205578), 4(0.1930068), 4(0.1576692), 4(0.142776), 4(0.1296), 4(0.1187028), 4(0.1152576), 4(0.0640764),
		4(0.0236844), 4(0.0324216), 4(0.0692064), 4(0.1137564), 4(0.1436292), 4(0.1567836), 4(0.141912), 4(0.1055592), 4(0.1039932), 4(0.0934092), 4(0.0904392), 4(0.0753192),
		4(0.094176), 4(0.11664), 4(0.1324296), 4(0.1532628), 4(0.179334), 4(0.1873476), 4(0.16092), 4(0.1465452), 4(0.1107216), 4(0.1079028), 4(0.1178172), 4(0.11448),
		4(0.114372), 4(0.1121364), 4(0.113724), 4(0.1232928), 4(0.1544832), 4(0.164646), 4(0.1372248), 4(0.1197936), 4(0.098928), 4(0.0945216), 4(0.0987228), 4(0.098604),
		4(0.1005372), 4(0.1195128), 4(0.1374084), 4(0.1529388), 4(0.1640088), 4(0.160002), 4(0.1404108), 4(0.1203012), 4(0.12312), 4(0.1135836), 4(0.121122), 4(0.1113912),
		4(0.10368), 4(0.097092), 4(0.093852), 4(0.097794), 4(0.1047708), 4(0.1073736), 4(0.0978804), 4(0.0824688), 4(0.0540432), 4(0.016038), 4(0.0560736), 4(0.05184),
		4(0.0588708), 4(0.0791316), 4(0.0940032), 4(0.1425492), 4(0.15444), 4(0.1435968), 4(0.1311768), 4(0.11718), 4(0.1134216), 4(0.10287), 4(0.0972108), 4(0.0926532),
		4(0.0859896), 4(0.0844344), 4(0.084888), 4(0.0869508), 4(0.0919512), 4(0.0886356), 4(0.084186), 4(0.0742608), 4(0.0340956), 4(0.0137268), 4(0.0090072), 4(0.0057564),
		4(0.0104112), 4(0.03348), 4(0.0786024), 4(0.1285416), 4(0.1432188), 4(0.1512), 4(0.1364364), 4(0.1175796), 4(0.1102248), 4(0.088614), 4(0.0892296), 4(0.0895212),
		4(0.0872208), 4(0.0873828), 4(0.092718), 4(0.111564), 4(0.1459944), 4(0.1650996), 4(0.1475496), 4(0.1150524), 4(0.0911736), 4(0.0838188), 4(0.0725976), 4(0.0486756),
		4(0.0543132), 4(0.0770472), 4(0.1122876), 4(0.1642572), 4(0.1824984), 4(0.1836), 4(0.15282), 4(0.1292544), 4(0.1171152), 4(0.10098), 4(0.099576), 4(0.0971892),
		4(0.1000404), 4(0.096876), 4(0.103248), 4(0.1221804), 4(0.1527228), 4(0.1476144), 4(0.0788184), 4(0.0556524), 4(0.033966), 4(0.0033156), 4(0.0044496), 4(0.0034992),
		4(0.0080676), 4(0.0745524), 4(0.1153116), 4(0.1616328), 4(0.18495), 4(0.178416), 4(0.1556388), 4(0.1349568), 4(0.1285092), 4(0.1130112), 4(0.1197396), 4(0.1151928),
		4(0.113292), 4(0.1126548), 4(0.1180764), 4(0.138024), 4(0.1770012), 4(0.1575828), 4(0.1099116), 4(0.0314172), 4(0.0230472), 4(0.0017064), 4(0.0002052), 4(0.001404),
		4(0.0042444), 4(0.07425), 4(0.1289088), 4(0.1772928), 4(0.2667708), 4(0.2296512), 4(0.1785348), 4(0.1571184), 4(0.1424952), 4(0.1250316), 4(0.1358532), 4(0.119772),
		4(0.1138968), 4(0.1154304), 4(0.1230444), 4(0.141642), 4(0.1664928), 4(0.1559628), 4(0.1072116), 4(0.087264), 4(0.0393336), 4(0.0036936), 4(0.0004644), 4(0.000702),
		4(0.0190728), 4(0.0910548), 4(0.1377324), 4(0.1914516), 4(0.2737044), 4(0.2508084), 4(0.1867536), 4(0.1605096), 4(0.1471608), 4(0.137484), 4(0.1430244), 4(0.132408),
		4(0.1289088), 4(0.1239192), 4(0.128898), 4(0.1521288), 4(0.1841832), 4(0.1653588), 4(0.1232388), 4(0.0808056), 4(0.0430488), 4(0.0079056), 4(0.00189), 4(0.0002376),
		4(0.0067608), 4(0.0624348), 4(0.1274616), 4(0.1607364), 4(0.2246508), 4(0.1900584), 4(0.1624212), 4(0.1486404), 4(0.132354), 4(0.1172556), 4(0.106812), 4(0.0965088),
		4(0.1034424), 4(0.1046304), 4(0.1058292), 4(0.1103976), 4(0.0961416), 4(0.076086), 4(0.0631044), 4(0.0527472), 4(0.023598), 4(0.0159948), 4(0.046926), 4(0.0540972),
		4(0.0613224), 4(0.0924372), 4(0.1254852), 4(0.1314252), 4(0.1388988), 4(0.1359504), 4(0.1250316), 4(0.0847152), 4(0.081108), 4(0.06696), 4(0.0401004), 4(0.03915),
		4(0.0478116), 4(0.0467424), 4(0.0470232), 4(0.0467316), 4(0.0483192), 4(0.041256), 4(0.0276156), 4(0.0231984), 4(0.0148824), 4(0.010368), 4(0.0145692), 4(0.0054108),
		4(0.0123768), 4(0.0467208), 4(0.097092), 4(0.1409076), 4(0.1566756), 4(0.1554228), 4(0.151632), 4(0.1417932), 4(0.1374084), 4(0.1233792), 4(0.1183032), 4(0.11637),
		4(0.1103112), 4(0.107298), 4(0.1109052), 4(0.1302696), 4(0.1545156), 4(0.1774008), 4(0.1754136), 4(0.1472364), 4(0.1205388), 4(0.1193184), 4(0.113616), 4(0.1166832),
		4(0.1260144), 4(0.1354752), 4(0.1469664), 4(0.1676052), 4(0.225018), 4(0.2084832), 4(0.1749708), 4(0.150984), 4(0.1370196), 4(0.1251072), 4(0.10989), 4(0.1109808),
		4(0.1094148), 4(0.1137564), 4(0.113076), 4(0.1185732), 4(0.1511568), 4(0.1553904), 4(0.1502604), 4(0.12474), 4(0.11718), 4(0.1110024), 4(0.1050516), 4(0.1064772),
		4(0.1191672), 4(0.1322028), 4(0.1511568), 4(0.15525), 4(0.1925208), 4(0.1871856), 4(0.160488), 4(0.1487268), 4(0.1365984), 4(0.110214), 4(0.1091016), 4(0.106596),
		4(0.1064016), 4(0.1079244), 4(0.1107216), 4(0.1205388), 4(0.1464264), 4(0.1543536), 4(0.1490616), 4(0.1211652), 4(0.1083348), 4(0.1047708), 4(0.1027296), 4(0.091908),
		4(0.1026864), 4(0.110538), 4(0.127116), 4(0.154818), 4(0.1812996), 4(0.1863648), 4(0.1700028), 4(0.142668), 4(0.1342008), 4(0.1196856), 4(0.1138104), 4(0.1077084),
		4(0.1057968), 4(0.1071468), 4(0.1059372), 4(0.1139292), 4(0.1418364), 4(0.15228), 4(0.13338), 4(0.0971136), 4(0.0874692), 4(0.0493992), 4(0.04212), 4(0.0297),
		4(0.0637956), 4(0.0911844), 4(0.1082484), 4(0.1454544), 4(0.1713312), 4(0.1830816), 4(0.1533384), 4(0.1351404), 4(0.12285), 4(0.109512), 4(0.099144), 4(0.08586),
		4(0.0853416), 4(0.0862488), 4(0.086778), 4(0.1185948), 4(0.141156), 4(0.131976), 4(0.1102464), 4(0.0834624), 4(0.073872), 4(0.0550908), 4(0.0735588), 4(0.081054),
		4(0.0810432), 4(0.112914), 4(0.1191132), 4(0.1475928), 4(0.1800792), 4(0.1791612), 4(0.1642248), 4(0.139266), 4(0.1315224), 4(0.1212516), 4(0.1260792), 4(0.1137672),
		4(0.1047384), 4(0.1047708), 4(0.1076652), 4(0.1040364), 4(0.0920052), 4(0.1079244), 4(0.102654), 4(0.0875772), 4(0.0980748), 4(0.101952), 4(0.0973728), 4(0.0860328),
		4(0.0907416), 4(0.09612), 4(0.1204956), 4(0.13689), 4(0.1678644), 4(0.1719684), 4(0.1418472), 4(0.1155708), 4(0.0931284), 4(0.0756324), 4(0.0499284), 4(0.0171504),
		4(0.0054972), 4(0.001296), 4(9.72E-05), 4(0.0011016), 4(0.0011772), 4(0.001728), 4(0.000108), 4(-0.0008856), 4(-0.0044712), 4(-0.016794), 4(-0.024732), 4(-0.0234252),
		4(-0.01161), 4(-0.0038664), 4(-0.002214), 4(0.0343872), 4(0.095202), 4(0.0986472), 4(0.09558), 4(0.0917568), 4(0.054864), 4(0.0783216), 4(0.07101), 4(0.0717876),
		4(0.0763452), 4(0.0797256), 4(0.1066068), 4(0.1601424), 4(0.204714), 4(0.1906092), 4(0.1490832), 4(0.1241892), 4(0.1147284), 4(0.1007532), 4(0.0931068), 4(0.0853848),
		4(0.0827388), 4(0.0965304), 4(0.121014), 4(0.1552932), 4(0.2376432), 4(0.208602), 4(0.1483272), 4(0.1257552), 4(0.1110024), 4(0.1108188), 4(0.104544), 4(0.1025028),
		4(0.1041228), 4(0.1015848), 4(0.1119852), 4(0.1436616), 4(0.1899504), 4(0.1721196), 4(0.119016), 4(0.0971784), 4(0.0837324), 4(0.0729216), 4(0.0497988), 4(0.0529308),
		4(0.063774), 4(0.0988956), 4(0.1104732), 4(0.150822), 4(0.1844424), 4(0.1531656), 4(0.1248264), 4(0.10611), 4(0.087804), 8(0.0763884), 4(0.0763236), 4(0.0782244),
		4(0.0793692), 4(0.094122), 4(0.1310364), 4(0.1680912), 4(0.1364364), 4(0.0936684), 4(0.0721872), 4(0.0539784), 4(0.0527688), 4(0.0516456), 4(0.0528228), 4(0.0762696),
		4(0.0892836), 4(0.1145448), 4(0.1249668), 4(0.163296), 4(0.1449576), 4(0.1180116), 4(0.0979236), 4(0.082134), 4(0.0786024), 4(0.082242), 4(0.0783216), 4(0.0791316),
		4(0.085266), 4(0.1108404), 4(0.1525068), 4(0.1803168), 4(0.143964), 4(0.0854388), 4(0.0449388), 4(0.0023436), 4(-5.4E-05), 4(-0.0026676), 4(7.56E-05), 4(0.0056268),
		4(0.0464508), 4(0.0988416), 4(0.15768), 4(0.2069928), 4(0.1957824), 4(0.155196), 4(0.1250748), 4(0.115398), 4(0.120636), 4(0.1153656), 4(0.1161432), 4(0.1162404),
		4(0.1199124), 4(0.1269432), 4(0.1723032), 4(0.2012256), 4(0.1536516), 4(0.1045656), 4(0.0711828), 4(0.0084456), 4(0.0), 4(-0.000864), 4(-0.000702), 4(0.0011124),
		4(0.0440208), 4(0.1187568), 4(0.144018), 4(0.1943892), 4(0.1816884), 4(0.1463508), 4(0.1414044), 4(0.120312), 4(0.1343952), 4(0.121824), 4(0.117882), 4(0.1172556),
		4(0.1168344), 4(0.1170072), 4(0.1300752), 4(0.1264248), 4(0.1114776), 4(0.0626724), 4(0.0007128), 4(-0.0008424), 4(-0.0193104), 4(-0.0406296), 4(-0.0391392), 4(-0.027378),
		4(0.0044712), 4(0.0357912), 4(0.0894132), 4(0.1547208), 4(0.1366092), 4(0.1053432), 4(0.0853092), 4(0.07425), 4(0.076086), 4(0.0674892), 4(0.06993), 4(0.0769716),
		4(0.0790452), 4(0.0877068), 4(0.086724), 4(0.088398), 4(0.0452952), 4(0.000108), 4(-0.0017064), 4(-0.0238572), 4(-0.053676), 4(-0.078732), 4(-0.0623376), 4(-0.0312228),
		4(-0.0057672), 4(0.0648432), 4(0.147474), 4(0.1614384), 4(0.1543968), 4(0.1360368), 4(0.1243404), 4(0.1108836), 4(0.0975888), 4(0.0961956), 4(0.0922104), 4(0.0947268),
		4(0.0965844), 4(0.1113912), 4(0.1432188), 4(0.1895832), 4(0.1559088), 4(0.1177956), 4(0.091692), 4(0.069714), 4(0.044496), 4(0.0462132), 4(0.0648108), 4(0.0874584),
		4(0.1036692), 4(0.1245888), 4(0.1679184), 4(0.1964952), 4(0.199206), 4(0.1556388), 4(0.1374732), 4(0.1198044), 4(0.1027512), 4(0.0974592), 4(0.0986472), 4(0.1008504),
		4(0.1032156), 4(0.1205712), 4(0.1641816), 4(0.193914), 4(0.1477116), 4(0.0986256), 4(0.0863892), 4(0.0829656), 4(0.0634176), 4(0.058482), 4(0.0728784), 4(0.0916488),
		4(0.1005912), 4(0.110322), 4(0.173988), 4(0.2445012), 4(0.2341332), 4(0.1611684), 4(0.134622), 4(0.119988), 4(0.1241676), 4(0.1159272), 4(0.1125792), 4(0.1121364),
		4(0.1148688), 4(0.1344708), 4(0.1790208), 4(0.1892376), 4(0.1422036), 4(0.1101384), 4(0.0935496), 4(0.0719064), 4(0.0168264), 4(0.0208332), 4(0.0560736), 4(0.080298),
		4(0.1092204), 4(0.118692), 4(0.1336284), 4(0.2242944), 4(0.2358504), 4(0.1809), 4(0.1442664), 4(0.1234116), 4(0.1139616), 4(0.1056348), 4(0.1038852), 4(0.103032),
		4(0.108972), 4(0.1207224), 4(0.1610712), 4(0.1946376), 4(0.1502064), 4(0.113184), 4(0.0890028), 4(0.0739584), 4(0.0424116), 4(0.0027648), 4(9.72E-05), 4(0.0023652),
		4(0.0735912), 4(0.0892836), 4(0.1238868), 4(0.1767744), 4(0.18414), 4(0.1397844), 4(0.1205496), 4(0.093258), 4(0.0891756), 4(0.085266), 4(0.0749844), 4(0.0763452),
		4(0.0837648), 4(0.0936144), 4(0.1195776), 4(0.1210788), 4(0.0954072), 4(0.0687636), 4(0.0160056), 4(0.0003456), 4(-0.0001944), 4(-0.0003996), 4(-0.0012204), 4(-1.08E-05),
		4(0.0644436), 4(0.1005372), 4(0.1495152), 4(0.2005128), 4(0.2052108), 4(0.1707912), 4(0.1496556), 4(0.1200096), 4(0.1212516), 4(0.1176876), 4(0.1135836), 4(0.111672),
		4(0.1126116), 4(0.1131084), 4(0.1209168), 4(0.1166508), 4(0.107244), 4(0.0751788), 4(0.0218052), 4(0.0), 4(-0.0082512), 4(-0.0096336), 4(-0.0296352), 4(-0.0058104),
		4(0.0024084), 4(0.0930852), 4(0.1310688), 4(0.1958904), 4(0.1957068), 4(0.1428516), 4(0.1317492), 4(0.1090692), 4(0.1047492), 4(0.0844236), 4(0.06723), 4(0.0808596),
		4(0.068904), 4(0.07047), 4(0.0669492), 4(0.02997), 4(0.0145044), 4(0.0091044), 4(0.0), 4(-2.16E-05), 4(-0.0039528), 4(-0.0203472), 4(-0.0274104), 4(-0.0107244),
		4(-1.08E-05), 4(0.067554), 4(0.1166076), 4(0.1562004), 4(0.1356588), 4(0.148338), 4(0.115992), 4(0.1072872), 4(0.1001376), 4(0.094446), 4(0.0936252), 4(0.0940464),
		4(0.0972324), 4(0.1147392), 4(0.134136), 4(0.1655532), 4(0.1559304), 4(0.1219968), 4(0.1114668), 4(0.1099224), 4(0.1146636), 4(0.0954828), 4(0.0881172), 4(0.0972108),
		4(0.1171152), 4(0.1199016), 4(0.1491372), 4(0.1905984), 4(0.1769904), 4(0.1226016), 4(0.1017792), 4(0.0915732), 4(0.0911844), 4(0.0888516), 4(0.082134), 4(0.0800496),
		4(0.0826848), 4(0.1007748), 4(0.1189296), 4(0.1303128), 4(0.1203444), 4(0.1157328), 4(0.1088316), 4(0.1033992), 4(0.110484), 4(0.1044684), 4(0.1045116), 4(0.1028592),
		4(0.113508), 4(0.1146852), 4(0.12258), 4(0.1606068), 4(0.166266), 4(0.1270404), 4(0.1207116), 4(0.1108404), 4(0.0989604), 4(0.0937116), 4(0.0941868), 4(0.0989712),
		4(0.1060128), 4(0.1160028), 4(0.1389204), 4(0.1464372), 4(0.1187352), 4(0.0677916), 4(0.0260604), 4(0.0118152), 4(0.006804), 4(0.0032724), 4(0.0025704), 4(0.0147204),
		4(0.0669168), 4(0.1053324), 4(0.1277748), 4(0.1716444), 4(0.175284), 4(0.1328184), 4(0.1192644), 4(0.1064772), 4(0.099576), 4(0.0939276), 4(0.0925668), 4(0.091908),
		4(0.093906), 4(0.101358), 4(0.1204632), 4(0.1335636), 4(0.1250856), 4(0.0778032), 4(0.0428112), 4(0.0188352), 4(0.0135324), 4(0.0105624), 4(0.0170424), 4(0.0813132),
		4(0.0984852), 4(0.1112832), 4(0.1260576), 4(0.1449144), 4(0.1362852), 4(0.122904), 4(0.106812), 4(0.1047492), 4(0.0972648), 4(0.0883116), 4(0.0846504), 4(0.0844128),
		4(0.0861948), 4(0.0853416), 4(0.0876312), 4(0.0921024), 4(0.0929556), 4(0.0878256), 4(0.092124), 4(0.0933336), 4(0.085482), 4(0.0714852), 4(0.069174), 4(0.073278),
		4(0.0888084), 4(0.104436), 4(0.1191024), 4(0.1419336), 4(0.1508112), 4(0.1315656), 4(0.122418), 4(0.1136808), 4(0.1031832), 4(0.0919836), 4(0.0969948), 4(0.0951048),
		4(0.0976968), 4(0.1049112), 4(0.1099656), 4(0.1059696), 4(0.09045), 4(0.0593676), 4(0.0165456), 4(0.0049032), 4(0.0), 4(-0.0026244), 4(-0.0063288), 4(-0.0007668),
		4(0.000216), 4(0.0784836), 4(0.1226556), 4(0.1489104), 4(0.181116), 4(0.1473984), 4(0.1261332), 4(0.1095876), 4(0.1113372), 4(0.1074492), 4(0.1029132), 4(0.1074924),
		4(0.1061208), 4(0.1018764), 4(0.1026432), 4(0.0850716), 4(0.0643032), 4(0.0005616), 4(-0.00108), 4(-0.0438264), 4(-0.1085184), 4(-0.1069632), 4(-0.0672084), 4(-0.0093204),
		4(0.0), 4(0.0681696), 4(0.1159164), 4(0.120852), 4(0.148608), 4(0.1387368), 4(0.1311444), 4(0.1202796), 4(0.115452), 4(0.1081512), 4(0.1023084), 4(0.1019736),
		4(0.1065636), 4(0.1056132), 4(0.1011636), 4(0.0946836), 4(0.0807948), 4(0.0301536), 4(-0.0018468), 4(-0.0013392), 4(-0.0304992), 4(-0.0383616), 4(-0.0051408), 4(0.0100548),
		4(0.0472284), 4(0.0835056), 4(0.1080324), 4(0.1305504), 4(0.1498932), 4(0.142668), 4(0.1325916), 4(0.1150308), 4(0.10503), 4(0.0969948), 4(0.095688), 4(0.092934),
		4(0.0926748), 4(0.1090368), 4(0.13473), 4(0.1637928), 4(0.1512756), 4(0.1119744), 4(0.0972108), 4(0.0858816), 4(0.0816156), 4(0.0716472), 4(0.0775332), 4(0.08559),
		4(0.0961524), 4(0.1151388), 4(0.166536), 4(0.25704), 4(0.2649024), 4(0.1657044), 4(0.134838), 4(0.1278936), 4(0.120042), 4(0.1111428), 4(0.1089396), 4(0.1093176),
		4(0.1144908), 4(0.1238868), 4(0.148446), 4(0.1554012), 4(0.1232496), 4(0.1085616), 4(0.092178), 4(0.0950508), 4(0.0863352), 4(0.0863136), 4(0.0951156), 4(0.1047924),
		4(0.1126332), 4(0.1224504), 4(0.1525176), 4(0.2163024), 4(0.233982), 4(0.1381968), 4(0.1173312), 4(0.1114992), 4(0.1053972), 4(0.0984636), 4(0.096984), 4(0.0951588),
		4(0.0964548), 4(0.104112), 4(0.12069), 4(0.129762), 4(0.1272348), 4(0.1106352), 4(0.1011204), 4(0.0885924), 4(0.08532), 4(0.081108), 4(0.0845316), 4(0.0884736),
		4(0.094878), 4(0.108486), 4(0.1284228), 4(0.140292), 4(0.170208), 4(0.1236384), 4(0.1150524), 4(0.100548), 4(0.1026432), 4(0.0913464), 4(0.0899424), 4(0.0921132),
		4(0.0935712), 4(0.1056348), 4(0.1142208), 4(0.1224612), 4(0.1139616), 4(0.089154), 4(0.0855684), 4(0.0797256), 4(0.0720036), 4(0.0555984), 4(0.0483516), 4(0.0726408),
		4(0.0891432), 4(0.0930528), 4(0.1091232), 4(0.1262304), 4(0.132894), 4(0.1184004), 4(0.1083996), 4(0.0994572), 4(0.1152684), 4(0.1028052), 4(0.1022544), 4(0.100332),
		4(0.0995868), 4(0.1011312), 4(0.1030644), 4(0.0941976), 4(0.0744228), 4(0.037206), 4(0.002754), 4(-1.08E-05), 4(-0.0003564), 4(-0.0021708), 4(-0.004806), 4(-0.0011556),
		4(0.0), 4(0.0334692), 4(0.086184), 4(0.1063584), 4(0.1207116), 4(0.102708), 4(0.0932472), 4(0.0797904), 4(0.075438), 4(0.0660312), 4(0.0624348), 4(0.0630396),
		4(0.0702432), 4(0.071982), 4(0.0714744), 4(0.0671436), 4(0.0379296), 4(4.32E-05), 4(-0.00324), 4(-0.0293004), 4(-0.0782676), 4(-0.1019088), 4(-0.0983664), 4(-0.048546),
		4(-0.0055836), 4(0.019818), 4(0.1018872), 4(0.1191996), 4(0.133866), 4(0.1172664), 4(0.10692), 4(0.101574), 4(0.1014768), 4(0.0955044), 4(0.0905364), 4(0.0940788),
		4(0.0999756), 4(0.1090908), 4(0.1507896), 4(0.1415772), 4(0.1030644), 4(0.0727596), 4(0.0104004), 4(-1.08E-05), 4(-0.0036072), 4(-0.006372), 4(-0.0066744), 4(-0.0016632),
		4(0.0024624), 4(0.0800388), 4(0.1211112), 4(0.1627776), 4(0.2053512), 4(0.13932), 4(0.1145448), 4(0.104922), 4(0.1003212), 4(0.096012), 4(0.0908172), 4(0.0884952),
		4(0.0898992), 4(0.1005372), 4(0.1155708), 4(0.1219212), 4(0.1014876), 4(0.0683964), 4(0.00405), 4(0.0), 4(-0.0008208), 4(-0.002052), 4(-0.0012096), 4(1.08E-05),
		4(0.0165672), 4(0.0854604), 4(0.109998), 4(0.1488564), 4(0.1870992), 4(0.1397088), 4(0.1188756), 4(0.1069848), 4(0.1026), 4(0.097308), 4(0.0969516), 4(0.0975132),
		4(0.10152), 4(0.1054404), 4(0.1240812), 4(0.1299672), 4(0.1004832), 4(0.0732132), 4(0.0076464), 4(0.0), 4(-0.00108), 4(-0.0067068), 4(-0.00324), 4(-2.16E-05),
		4(0.0225612), 4(0.0873072), 4(0.108972), 4(0.1333692), 4(0.1820232), 4(0.1380564), 4(0.1175148), 4(0.1079136), 4(0.1085184), 4(0.1022976), 4(0.100602), 4(0.100872),
		4(0.10098), 4(0.0932904), 4(0.0875772), 4(0.0758484), 4(0.0585252), 4(0.0), 4(-0.00324), 4(-0.043308), 4(-0.0840024), 4(-0.1321488), 4(-0.1249128), 4(-0.0539892),
		4(-0.0055836), 4(0.0390636), 4(0.1058724), 4(0.1395468), 4(0.1763748), 4(0.1295892), 4(0.1079352), 4(0.0932904), 4(0.0951588), 4(0.0777924), 4(0.0668196), 4(0.0670896),
		4(0.0719172), 4(0.0837972), 4(0.0954072), 4(0.0823392), 4(0.0659988), 4(0.0239544), 4(0.000918), 4(-1.08E-05), 4(-0.000864), 4(-0.00324), 4(-0.00432), 4(-8.64E-05),
		4(0.000324), 4(0.076356), 4(0.111726), 4(0.1352592), 4(0.1588464), 4(0.1337688), 4(0.118206), 4(0.1072008), 4(0.1083132), 4(0.1037448), 4(0.1019304), 4(0.0991224),
		4(0.0958284), 4(0.095742), 4(0.0939168), 4(0.088344), 4(0.072252), 4(0.0146124), 4(1.08E-05), 4(-1.08E-05), 4(-0.0012528), 4(-0.0032832), 4(-0.0029052), 4(-3.24E-05),
		4(0.0), 4(0.0320976), 4(0.0815724), 4(0.092772), 4(0.1169964), 4(0.1018224), 4(0.0896076), 4(0.080082), 4(0.0669924), 4(0.049896), 4(0.0354996), 4(0.0224964),
		4(0.0220212), 4(0.0168264), 4(0.0147096), 4(0.0084564), 4(0.0031644), 4(0.0), 8(-1.08E-05), 4(-2.16E-05), 4(-0.00216), 4(-0.0054108), 4(-0.0017172), 4(-1.08E-05),
		4(0.0115668), 4(0.0917568), 4(0.1081512), 4(0.117396), 4(0.112752), 4(0.107298), 4(0.0980316), 4(0.073062), 4(0.0782352), 4(0.0683316), 4(0.0703944), 4(0.0736344),
		4(0.0959688), 4(0.1133892), 4(0.1383912), 4(0.121554), 4(0.1057968), 4(0.0998136), 4(0.0791748), 4(0.0630828), 4(0.06129), 4(0.0630504), 4(0.0752544), 4(0.1072224),
		4(0.1063584), 4(0.1234548), 4(0.1529928), 4(0.2298996), 4(0.1341252), 4(0.114426), 4(0.1076328), 4(0.0901044), 4(0.083376), 4(0.0793152), 4(0.0782136), 4(0.0890352),
		4(0.1010232), 4(0.117504), 4(0.1349244), 4(0.121986), 4(0.106488), 4(0.0984636), 4(0.0834084), 4(0.0767772), 4(0.0748656), 4(0.082188), 4(0.09693), 4(0.10422),
		4(0.1187352), 4(0.1399032), 4(0.1995624), 4(0.1647864), 4(0.1384452), 4(0.1172664), 4(0.108108), 4(0.1052676), 4(0.0991224), 4(0.0969624), 4(0.0992304), 4(0.0996192),
		4(0.1077732), 4(0.1334124), 4(0.151308), 4(0.130464), 4(0.1252908), 4(0.1233036), 4(0.1053108), 4(0.0926424), 4(0.095472), 4(0.0964872), 4(0.1048356), 4(0.109242),
		4(0.11286), 4(0.124686), 4(0.1476684), 4(0.1641168), 4(0.1295892), 4(0.120636), 4(0.108486), 4(0.108594), 4(0.103842), 4(0.1037232), 4(0.1064232), 4(0.103356),
		4(0.1196856), 4(0.135378), 4(0.1460484), 4(0.1295892), 4(0.1150524), 4(0.1010556), 4(0.0880416), 4(0.0741312), 4(0.0734832), 4(0.080946), 4(0.0917028), 4(0.1069632),
		4(0.1270404), 4(0.1392876), 4(0.1683828), 4(0.2076624), 4(0.1483164), 4(0.1402164), 4(0.1265652), 4(0.1089288), 4(0.108918), 4(0.1056888), 4(0.1071036), 4(0.10746),
		4(0.1157328), 4(0.137268), 4(0.1338876), 4(0.0993276), 4(0.09261), 4(0.0594648), 4(0.0046332), 4(0.0041148), 4(0.0001836), 4(2.16E-05), 4(0.0539676), 4(0.0891108),
		4(0.1053324), 4(0.1233792), 4(0.1494936), 4(0.1941408), 4(0.1425492), 4(0.1244808), 4(0.1113912), 4(0.1144584), 4(0.1150632), 4(0.1104948), 4(0.1041984), 4(0.1083996),
		4(0.1083348), 4(0.1052352), 4(0.0992196), 4(0.0747576), 4(0.0101952), 4(0.0001188), 4(-0.0266004), 4(-0.064206), 4(-0.109242), 4(-0.1218996), 4(-0.0501552), 4(-0.0003672),
		4(0.048924), 4(0.115236), 4(0.1368576), 4(0.2568348), 4(0.1327212), 4(0.1220832), 4(0.1079136), 4(0.1080648), 4(0.1071144), 4(0.1053216), 4(0.1077192), 4(0.1077732),
		4(0.1077624), 4(0.0990792), 4(0.0740232), 4(0.0053568), 4(-0.000108), 4(-0.0128304), 4(-0.031752), 4(-0.053622), 4(-0.1621728), 4(-0.1631232), 4(-0.1230984), 4(-0.0197532),
		4(0.0024084), 4(0.1368144), 4(0.1777356), 4(0.2075004), 4(0.1311444), 4(0.1164564), 4(0.0999108), 4(0.0973836), 4(0.0920268), 4(0.0915192), 4(0.0922104), 4(0.0959904),
		4(0.1181736), 4(0.183114), 4(0.18117), 4(0.1382508), 4(0.1005912), 4(0.0831924), 4(0.0682452), 4(0.08856), 4(0.0952776), 4(0.1076976), 4(0.089262), 4(0.100386),
		4(0.1452492), 4(0.1892592), 4(0.2874204), 4(0.398142), 4(0.1982556), 4(0.1593756), 4(0.1203984), 4(0.1186812), 4(0.1068012), 4(0.1048248), 4(0.1049328), 4(0.1081728),
		4(0.1320624), 4(0.148176), 4(0.1388016), 4(0.1085832), 4(0.0890784), 4(0.040014), 4(0.01296), 4(0.0476172), 4(0.0699948), 4(0.0722196), 4(0.0861624), 4(0.1033236),
		4(0.102492), 4(0.1289088), 4(0.206118), 4(0.3784752), 4(0.1723788), 4(0.133326), 4(0.1205496), 4(0.1241244), 4(0.1132056), 4(0.112914), 4(0.11232), 4(0.1106676),
		4(0.11826), 4(0.1400868), 4(0.131814), 4(0.1078812), 4(0.0788292), 4(0.0158652), 4(0.0215028), 4(0.0409536), 4(0.042174), 4(0.0464184), 4(0.053028), 4(0.080568),
		4(0.108), 4(0.1353888), 4(0.2057724), 4(0.3596508), 4(0.149526), 4(0.1296864), 4(0.1213272), 4(0.1189188), 4(0.1101924), 4(0.1071144), 4(0.109026), 4(0.1114668),
		4(0.1188216), 4(0.1345248), 4(0.1406052), 4(0.1073304), 4(0.074952), 4(0.0139752), 4(0.0087156), 4(0.0107244), 4(0.0185112), 4(0.0243), 4(0.0544644), 4(0.0997812),
		4(0.1133352), 4(0.127548), 4(0.1606176), 4(0.1883736), 4(0.1441152), 4(0.1249776), 4(0.1201068), 4(0.1119852), 4(0.0981396), 4(0.0953856), 4(0.0943596), 4(0.0985392),
		4(0.1052676), 4(0.1185624), 4(0.125874), 4(0.11988), 4(0.1070604), 4(0.0822744), 4(0.0500256), 4(0.0670464), 4(0.0664308), 4(0.0704916), 4(0.0389556), 4(0.0719712),
		4(0.0899964), 4(0.1389744), 4(0.1404972), 4(0.1750788), 4(0.1504548), 4(0.1267164), 4(0.1187244), 4(0.1025028), 4(0.1025676), 4(0.0971136), 4(0.0976104), 4(0.0991008),
		4(0.1047384), 4(0.1007856), 4(0.0982584), 4(0.0659556), 4(0.0012312), 4(3.24E-05), 4(0.0022896), 4(-0.0045684), 4(-0.0105624), 4(-0.0120852), 4(-0.004212), 4(0.0168696),
		4(0.103248), 4(0.1315008), 4(0.1367496), 4(0.2086992), 4(0.168588), 4(0.1741176), 4(0.149526), 4(0.1169748), 4(0.111294), 4(0.108216), 4(0.10692), 4(0.1079784),
		4(0.1076112), 4(0.1000404), 4(0.09558), 4(0.0674784), 4(0.0087372), 4(0.0), 4(-0.000216), 4(-0.00216), 4(-0.0079596), 4(-0.0162), 4(-0.0096876), 4(-0.0001944),
		4(0.0266004), 4(0.1076976), 4(0.1350864), 4(0.1609092), 4(0.1439424), 4(0.1304532), 4(0.1149876), 4(0.1225692), 4(0.1158084), 4(0.108216), 4(0.1047708), 4(0.1207008),
		4(0.1344384), 4(0.1598184), 4(0.1454976), 4(0.134082), 4(0.1046628), 4(0.0786996), 4(0.0315252), 4(0.0137916), 4(0.0054), 4(0.00864), 4(0.031644), 4(0.0960444),
		4(0.1199988), 4(0.1412748), 4(0.1701648), 4(0.2475684), 4(0.165942), 4(0.153036), 4(0.133164), 4(0.1355076), 4(0.1200204), 4(0.1187892), 4(0.125226), 4(0.1433052),
		4(0.1516968), 4(0.1575072), 4(0.1465776), 4(0.1102248), 4(0.1443636), 4(0.0680832), 4(0.01728), 4(0.0474336), 4(0.0505008), 4(0.0750492), 4(0.1015524), 4(0.1183032),
		4(0.125226), 4(0.1600668), 4(0.2360664), 4(0.3586572), 4(0.2145528), 4(0.1586304), 4(0.1271052), 4(0.126846), 4(0.1122768), 4(0.10854), 4(0.108), 4(0.1068984),
		4(0.11259), 4(0.135864), 4(0.14904), 8(0.1380024), 4(0.1104948), 4(0.1079136), 4(0.1441044), 4(0.0809352), 4(0.0972864), 4(0.08856), 4(0.10638), 4(0.164808),
		4(0.1511136), 4(0.1728), 4(0.244026), 4(0.1728), 4(0.127386), 4(0.1714716), 4(0.1155492), 4(0.1046412), 4(0.099252), 4(0.1009584), 4(0.100494), 4(0.107784),
		4(0.1307772), 4(0.1335528), 4(0.1153332), 4(0.0972648), 4(0.0782136), 4(0.0742284), 4(0.0745416), 4(0.0848016), 4(0.0877176), 4(0.1006236), 4(0.1068768), 4(0.1139616),
		4(0.1231416), 4(0.1410264), 4(0.2009556), 4(0.1498176), 4(0.1325592), 4(0.1225476), 4(0.1203012), 4(0.1095876), 4(0.1022436), 4(0.1019952), 4(0.1123956), 4(0.1309932),
		4(0.1546668), 4(0.1647864), 4(0.14688), 4(0.1138968), 4(0.1063476), 4(0.0952236), 4(0.0704808), 4(0.0646488), 4(0.0784728), 4(0.0910872), 4(0.10611), 4(0.1036152),
		4(0.1372248), 4(0.1579608), 4(0.2321676), 4(0.1640844), 4(0.1405836), 4(0.1221264), 4(0.1219212), 4(0.1096848), 4(0.102546), 4(0.0975564), 4(0.0960444), 4(0.09612),
		4(0.09963), 4(0.0857736), 4(0.0697572), 4(0.0132408), 4(0.0001188), 4(0.0020412), 4(0.0028512), 4(0.0034668), 4(0.0050436), 4(0.0023328), 4(0.0112752), 4(0.061884),
		4(0.1006236), 4(0.131598), 4(0.1714932), 4(0.143316), 4(0.1268136), 4(0.1065204), 4(0.0853956), 4(0.055566), 4(0.0240732), 4(0.0094068), 4(0.0050652), 4(0.0044928),
		4(0.001404), 4(0.0014364), 4(0.0006048), 4(0.0006156), 4(-2.16E-05), 4(-0.0010908), 4(0.0), 4(-0.000108), 4(-0.0054432), 4(-0.0015552), 4(0.0001728), 4(0.0081972),
		4(0.0522072), 4(0.1140372), 4(0.1248048), 4(0.1272996), 4(0.1148148), 4(0.1052568), 4(0.1039284), 4(0.0939384), 4(0.0904176), 4(0.0894132), 4(0.0949104), 4(0.1055052),
		4(0.1440396), 4(0.1637388), 4(0.1495368), 4(0.1128168), 4(0.0786132), 4(0.0399708), 4(0.0249804), 4(0.0192564), 4(0.0132084), 4(0.0109296), 4(0.0421308), 4(0.1064772),
		4(0.1375056), 4(0.1655856), 4(0.2446308), 4(0.1834272), 4(0.1646568), 4(0.125064), 4(0.112266), 4(0.0988308), 4(0.0900828), 4(0.0875016), 4(0.091152), 4(0.0979236),
		4(0.1111968), 4(0.0986148), 4(0.0764532), 4(0.0566352), 4(0.0049356), 4(0.0037908), 4(0.0001944), 4(0.0019872), 4(0.0054), 4(0.0240948), 4(0.0672516), 4(0.101304),
		4(0.125766), 4(0.1537272), 4(0.2341008), 4(0.1538784), 4(0.125172), 4(0.1048248), 4(0.0974484), 4(0.0846288), 4(0.0822312), 4(0.0766584), 4(0.0804708), 4(0.0921564),
		4(0.1108836), 4(0.111996), 4(0.107892), 4(0.1027944), 4(0.0878904), 4(0.083808), 4(0.075654), 4(0.0714528), 4(0.0676836), 4(0.065826), 4(0.086562), 4(0.1224504),
		4(0.1397196), 4(0.1499148), 4(0.1804572), 4(0.1550016), 4(0.1392552), 4(0.128466), 4(0.1038852), 4(0.0990792), 4(0.0972756), 4(0.0968544), 4(0.0965628), 4(0.0972648),
		4(0.1080324), 4(0.0871992), 4(0.088236), 4(0.065232), 4(0.018792), 4(0.001458), 4(-5.4E-05), 4(0.0184464), 4(0.01674), 4(0.0305748), 4(0.0394632), 4(0.0908496),
		4(0.0944568), 4(0.1191996), 4(0.1864188), 4(0.1461024), 4(0.1067256), 4(0.0862488), 4(0.0728892), 4(0.0557496), 4(0.0441288), 4(0.036666), 4(0.0403812), 4(0.0619704),
		4(0.0924588), 4(0.0738504), 4(0.0572508), 4(0.0314604), 4(0.001836), 4(0.0002052), 4(0.0040392), 4(0.0006912), 4(0.0002484), 4(0.0001296), 4(0.000162), 4(0.0238248),
		4(0.0842832), 4(0.1412532), 4(0.1762776), 4(0.1549584), 4(0.1406052), 4(0.1169856), 4(0.11556), 4(0.1095876), 4(0.1095012), 4(0.1109592), 4(0.112158), 4(0.1099332),
		4(0.096876), 4(0.0852444), 4(0.0590544), 4(0.00108), 4(-2.16E-05), 4(-0.00108), 4(-0.0033156), 4(-0.0142236), 4(-0.00837), 4(-0.00324), 4(-4.32E-05), 4(0.0477468),
		4(0.0958176), 4(0.141696), 4(0.2635524), 4(0.1943244), 4(0.1402812), 4(0.1119204), 4(0.1022652), 4(0.0918756), 4(0.0811512), 4(0.0760104), 4(0.0733212), 4(0.0671976),
		4(0.0372708), 4(0.01404), 4(0.002592), 4(-1.08E-05), 4(-0.000648), 4(-0.0022788), 4(-0.0059184), 4(-0.0139644), 4(-0.0220428), 4(-0.0168588), 4(-0.00648), 4(0.0103896),
		4(0.0524988), 4(0.1278072), 4(0.1284984), 4(0.1213596), 4(0.1189944), 4(0.1043388), 4(0.0950508), 4(0.0870048), 4(0.0853524), 4(0.0898452), 4(0.0964656), 4(0.1171584),
		4(0.1232496), 4(0.1143072), 4(0.1108188), 4(0.0956772), 4(0.0651564), 4(0.0358668), 4(0.0216), 4(0.0138024), 4(0.01188), 4(0.02133), 4(0.0661176), 4(0.1079568),
		4(0.1765908), 4(0.3469392), 4(0.4860864), 4(0.26784), 4(0.1620108), 4(0.1377432), 4(0.1282284), 4(0.1261008), 4(0.1164672), 4(0.1145556), 4(0.1159704), 4(0.1350216),
		4(0.1554444), 4(0.137538), 4(0.0964656), 4(0.062802), 4(0.006156), 4(0.0056592), 4(0.0068904), 4(0.0050652), 4(0.0030132), 4(0.010098), 4(0.044658), 4(0.0909468),
		4(0.1353456), 4(0.1728324), 4(0.256392), 4(0.1592244), 4(0.1248588), 4(0.126306), 4(0.1097388), 4(0.09288), 4(0.0863676), 4(0.0856224), 4(0.0912492), 4(0.1063908),
		4(0.1080216), 4(0.120366), 4(0.1102572), 4(0.0616032), 4(0.019764), 4(0.0150876), 4(0.0100656), 4(0.0104652), 4(0.0204768), 4(0.0584928), 4(0.11124), 4(0.1388988),
		4(0.182358), 4(0.235872), 4(0.3683772), 4(0.2498796), 4(0.1628424), 4(0.1323864), 4(0.141534), 4(0.124794), 4(0.113724), 4(0.1114776), 4(0.1157868), 4(0.1220724),
		4(0.1202364), 4(0.1400976), 4(0.1223748), 4(0.0857844), 4(0.0725976), 4(0.0539244), 4(0.0222696), 4(0.0136944), 4(0.0097308), 4(0.0267516), 4(0.091962), 4(0.1187028),
		4(0.1723896), 4(0.2221668), 4(0.3450708), 4(0.141912), 4(0.12339), 4(0.119394), 4(0.1108836), 4(0.1109916), 4(0.1019844), 4(0.099252), 4(0.0910764), 4(0.104922),
		4(0.1252152), 4(0.1134), 4(0.0784296), 4(0.0095904), 4(4.32E-05), 4(0.0035208), 4(0.0230364), 4(0.0484488), 4(0.043362), 4(0.0673812), 4(0.1042308), 4(0.1218456),
		4(0.1533492), 4(0.1487052), 4(0.2392416), 4(0.1461996), 4(0.13554), 4(0.1167156), 4(0.1227744), 4(0.1135512), 4(0.1086696), 4(0.1050192), 4(0.0993384), 4(0.0978264),
		4(0.0852444), 4(0.0829872), 4(0.0763884), 4(0.0613116), 4(0.031536), 4(0.0101952), 4(0.0012852), 4(-1.08E-05), 8(-2.16E-05), 4(0.0051084), 4(0.0542808), 4(0.1124064),
		4(0.220914), 4(0.1984716), 4(0.1426248), 4(0.1268676), 4(0.1132596), 4(0.105192), 4(0.0964656), 4(0.0910764), 4(0.0871668), 4(0.0844668), 4(0.0704808), 4(0.0487296),
		4(0.0044496), 4(0.0), 4(-0.00054), 4(-0.00216), 4(-0.003888), 4(-0.0186732), 4(-0.0281772), 4(-0.0354132), 4(-0.0223452), 4(0.007182), 4(0.094122), 4(0.1315116),
		4(0.1775628), 4(0.2268324), 4(0.1461024), 4(0.1164024), 4(0.0955692), 4(0.0949968), 4(0.0844344), 4(0.057294), 4(0.0558144), 4(0.059508), 4(0.07074), 4(0.1152576),
		4(0.1198692), 4(0.0993816), 4(0.0310608), 4(0.0198072), 4(0.0327024), 4(0.032778), 4(0.0394524), 4(0.0001728), 4(0.0155196), 4(0.0060696), 4(0.1347192), 4(0.1499472),
		4(0.1755108), 4(0.264762), 4(0.185814), 4(0.1346004), 4(0.1173852), 4(0.0981612), 4(0.0895968), 4(0.0771876), 4(0.0673596), 4(0.061506), 4(0.0814428), 4(0.0904932),
		4(0.092556), 4(0.0938628), 4(0.0725544), 4(0.0251964), 4(0.0030456), 4(0.002916), 4(0.0042876), 4(0.0351864), 4(0.0820152), 4(0.111078), 4(0.1142208), 4(0.1436292),
		4(0.236682), 4(0.2784888), 4(0.1508976), 4(0.1117476), 4(0.1179252), 4(0.0867456), 4(0.0793476), 4(0.0732564), 4(0.0795744), 4(0.079434), 4(0.10476), 4(0.1211544),
		4(0.1116828), 4(0.086832), 4(0.0623484), 4(0.020898), 4(0.0018684), 4(0.0072144), 4(0.0162864), 4(0.0223992), 4(0.0470772), 4(0.1081836), 4(0.1273428), 4(0.1238004),
		4(0.1679508), 4(0.2366928), 4(0.1964196), 4(0.1338552), 4(0.114696), 4(0.1250316), 4(0.096714), 4(0.0909792), 4(0.0917676), 4(0.0962496), 4(0.105678), 4(0.1190268),
		4(0.1024488), 4(0.0828792), 4(0.0399924), 4(1.08E-05), 4(0.0067068), 4(0.0241488), 4(0.0286416), 4(0.0509436), 4(0.05751), 4(0.0763236), 4(0.1107108), 4(0.1377756),
		4(0.194562), 4(0.2354076), 4(0.1548612), 4(0.1331532), 4(0.119394), 4(0.1273752), 4(0.1156788), 4(0.1081512), 4(0.104112), 4(0.101466), 4(0.1098468), 4(0.1141776),
		4(0.0954396), 4(0.0818856), 4(0.0436536), 4(0.006642), 4(0.0026244), 4(0.0062316), 4(0.0070956), 4(0.0139212), 4(0.0508464), 4(0.082674), 4(0.1157976), 4(0.0856224),
		4(0.1397736), 4(0.1737072), 4(0.14742), 4(0.129708), 4(0.1228176), 4(0.1137348), 4(0.0952992), 4(0.0897264), 4(0.0863136), 4(0.076896), 4(0.0692496), 4(0.0551772),
		4(0.0243864), 4(0.0093744), 4(0.0), 4(-0.0018792), 4(-0.0094608), 4(-0.0035964), 4(-0.007074), 4(-0.023436), 4(-0.0066204), 4(-9.72E-05), 4(0.0122904), 4(0.1031184),
		4(0.1500768), 4(0.1819152), 4(0.1509516), 4(0.143262), 4(0.1263708), 4(0.0990792), 4(0.0934848), 4(0.0919296), 4(0.093906), 4(0.096768), 4(0.0973404), 4(0.0855144),
		4(0.0631476), 4(0.011124), 4(0.0008208), 4(0.0), 4(-2.16E-05), 4(-0.0012744), 4(-0.0060264), 4(-0.0054), 4(-0.00216), 4(0.0), 4(0.0708264), 4(0.1212408),
		4(0.1461132), 4(0.1623132), 4(0.150606), 4(0.1439424), 4(0.1298484), 4(0.112482), 4(0.0996192), 4(0.0937872), 4(0.0932688), 4(0.0895968), 4(0.118638), 4(0.1185516),
		4(0.1324404), 4(0.111618), 4(0.087426), 4(0.0643032), 4(0.0597996), 4(0.0489996), 4(0.0471204), 4(0.0472716), 4(0.0797364), 4(0.1164132), 4(0.12339), 4(0.1369548),
		4(0.1420308), 4(0.2038392), 4(0.2098332), 4(0.1419444), 4(0.1309608), 4(0.1126008), 4(0.103464), 4(0.1013472), 4(0.1011096), 4(0.1019304), 4(0.1105704), 4(0.1262628),
		4(0.113832), 4(0.1038312), 4(0.0719172), 4(0.0064152), 4(0.0144828), 4(0.019224), 4(0.0210384), 4(0.034128), 4(0.0487728), 4(0.0869076), 4(0.1121256), 4(0.1290276),
		4(0.1652076), 4(0.2544156), 4(0.25002), 4(0.146988), 4(0.1266516), 4(0.1217916), 4(0.114696), 4(0.1093716), 4(0.1025244), 4(0.1039284), 4(0.1101168), 4(0.1198368),
		4(0.1233036), 4(0.1179684), 4(0.0779004), 4(0.0237708), 4(0.0012636), 4(0.004698), 4(0.0074628), 4(0.0149688), 4(0.0956556), 4(0.1121472), 4(0.1222668), 4(0.1513296),
		4(0.1998756), 4(0.2920428), 4(0.1903176), 4(0.1462968), 4(0.1251072), 4(0.1233144), 4(0.1181412), 4(0.111024), 4(0.1086048), 4(0.1050192), 4(0.1081512), 4(0.105408),
		4(0.0920376), 4(0.0803088), 4(0.0111888), 4(0.001728), 4(0.0064908), 4(0.0041688), 4(0.0290196), 4(0.034722), 4(0.0723168), 4(0.0699192), 4(0.1370628), 4(0.1520316),
		4(0.15984), 4(0.1751004), 4(0.1606608), 4(0.1512972), 4(0.1363068), 4(0.1316196), 4(0.117234), 4(0.118638), 4(0.116046), 4(0.1123308), 4(0.1180332), 4(0.1292112),
		4(0.1247184), 4(0.1100736), 4(0.0665928), 4(0.01674), 4(0.0040068), 4(0.0014472), 4(0.0025704), 4(0.0004968), 4(0.0084888), 4(0.07857), 4(0.1214892), 4(0.1335852),
		4(0.1467396), 4(0.2140452), 4(0.1911816), 4(0.148014), 4(0.1310904), 4(0.1293516), 4(0.1193184), 4(0.116802), 4(0.115668), 4(0.1170612), 4(0.1123848), 4(0.1087344),
		4(0.0979992), 4(0.0820044), 4(0.025272), 4(0.000216), 4(-5.4E-05), 4(9.72E-05), 4(-0.0121608), 4(-0.0070632), 4(-6.48E-05), 4(0.000216), 4(0.0830628), 4(0.1289628),
		4(0.1418148), 4(0.1637928), 4(0.1766556), 4(0.1519128), 4(0.1360584), 4(0.11799), 4(0.1090044), 4(0.1035828), 4(0.1008072), 4(0.098496), 4(0.0948348), 4(0.0805464),
		4(0.0285552), 4(0.0), 4(-9.72E-05), 4(-0.0119988), 4(-0.0366984), 4(-0.0538812), 4(-0.0822096), 4(-0.068418), 4(-0.03105), 4(-0.0011556), 4(0.028026), 4(0.1011096),
		4(0.1409292), 4(0.1519992), 4(0.1468584), 4(0.1372896), 4(0.1097604), 4(0.0923292), 4(0.0985932), 4(0.08721), 4(0.0870912), 4(0.1015416), 4(0.122742), 4(0.1363176),
		4(0.1230552), 4(0.0982044), 4(0.0436968), 4(0.0270756), 4(0.0405972), 4(0.0665928), 4(0.0669276), 4(0.0775872), 4(0.1097172), 4(0.14148), 4(0.15012), 4(0.2063232),
		4(0.2017872), 4(0.17307), 4(0.1608336), 4(0.133272), 4(0.1248696), 4(0.1080756), 4(0.1046628), 4(0.1011096), 4(0.0991656), 4(0.0924588), 4(0.1161756), 4(0.1274508),
		4(0.1290276), 4(0.100278), 4(0.0648108), 4(0.0324432), 4(0.0243432), 4(0.0190512), 4(0.0177336), 4(0.0194508), 4(0.0532116), 4(0.08721), 4(0.1349352), 4(0.155628),
		4(0.191376), 4(0.1916568), 4(0.184464), 4(0.1894968), 4(0.154332), 4(0.133164), 4(0.1138212), 4(0.1153872), 4(0.1079892), 4(0.1228284), 4(0.1260036), 4(0.1202256),
		4(0.1207548), 4(0.1074924), 4(0.0803736), 4(0.0287064), 4(0.0168156), 4(0.0170856), 4(0.0137376), 4(0.0324756), 4(0.0447876), 4(0.1053), 4(0.1256904), 4(0.1491048),
		4(0.2041848), 4(0.2267568), 4(0.2653668), 4(0.1892376), 4(0.1403244), 4(0.129546), 4(0.1185408), 4(0.1140372), 4(0.113238), 4(0.1132056), 4(0.121284), 4(0.1272456),
		4(0.1306476), 4(0.1153332), 4(0.1050732), 4(0.0949968), 4(0.087372), 4(0.0764208), 4(0.0724464), 4(0.0726192), 4(0.1070064), 4(0.1196532), 4(0.1327968), 4(0.1564812),
		4(0.2280852), 4(0.231768), 4(0.1820448), 4(0.1643328), 4(0.1386288), 4(0.127926), 4(0.1314576), 4(0.1225908), 4(0.1213596), 4(0.1183896), 4(0.1196532), 4(0.1212192),
		4(0.122256), 4(0.116316), 4(0.098766), 4(0.0856008), 4(0.072846), 4(0.059346), 4(0.0697896), 4(0.0748548), 4(0.0992412), 4(0.1045116), 4(0.1250748), 4(0.1391904),
		4(0.1592784), 4(0.1797444), 4(0.1571508), 4(0.1402704), 4(0.1227636), 4(0.107622), 4(0.097524), 4(0.0896076), 4(0.0851256), 4(0.0768636), 4(0.083106), 4(0.0826524),
		4(0.0644976), 4(0.030024), 4(0.0025272), 4(1.08E-05), 4(0.000162), 4(0.0002484), 4(-1.08E-05), 4(0.007776), 4(5.4E-05), 4(0.0324864), 4(0.1048464), 4(0.1136808),
		4(0.1214784), 4(0.1394928), 4(0.138888), 4(0.1296108), 4(0.11178), 4(0.1026756), 4(0.0965736), 4(0.0968328), 4(0.0937656), 4(0.0920052), 4(0.092124), 4(0.0932472),
		4(0.0725868), 4(0.0477144), 4(0.0023976), 4(0.0), 4(-0.0001296), 4(-0.004752), 4(-0.0142884), 4(-0.007236), 4(-0.0008424), 4(0.00162), 4(0.0497124), 4(0.0990252),
		4(0.1103112), 4(0.1209384), 4(0.1275156), 4(0.1228284), 4(0.10908), 4(0.1066284), 4(0.0961524), 4(0.0918324), 4(0.0908604), 4(0.0929664), 4(0.1032264), 4(0.1212948),
		4(0.1202472), 4(0.1114884), 4(0.1036908), 4(0.0807732), 4(0.0590436), 4(0.0407052), 4(0.0968868), 4(0.1061748), 4(0.11691), 4(0.1244592), 4(0.1278504), 4(0.1276776),
		4(0.1932552), 4(0.2946888), 4(0.2458188), 4(0.16956), 4(0.132462), 4(0.1201824), 4(0.109458), 4(0.096228), 4(0.0955476), 4(0.0972108), 4(0.1119096), 4(0.1241676),
		4(0.1273104), 4(0.1150416), 4(0.1123092), 4(0.098874), 4(0.0896292), 4(0.0532872), 4(0.0516132), 4(0.0717444), 4(0.084564), 4(0.098064), 4(0.1242108), 4(0.164214),
		4(0.3122388), 4(0.4338144), 4(0.388584), 4(0.2623536), 4(0.1559952), 4(0.1288332), 4(0.1110024), 4(0.0999432), 4(0.0994464), 4(0.0976212), 4(0.1071144), 4(0.1231308),
		4(0.1185516), 4(0.1128816), 4(0.0977184), 4(0.0837648), 4(0.0732888), 4(0.050328), 4(0.0368496), 4(0.057996), 4(0.0777708), 4(0.0928368), 4(0.1289304), 4(0.198234),
		4(0.4699296), 4(0.4789368), 4(0.21816), 4(0.148122), 4(0.122148), 4(0.1028808), 4(0.0955908), 4(0.08532), 4(0.0852444), 4(0.0873504), 4(0.0986472), 4(0.1117044),
		4(0.1153872), 4(0.113292), 4(0.097686), 4(0.0810648), 4(0.061938), 4(0.0455328), 4(0.0431892), 4(0.0624672), 4(0.0844776), 4(0.1244808), 4(0.1308096), 4(0.1752084),
		4(0.2456892), 4(0.3086964), 4(0.1867212), 4(0.1485432), 4(0.1245564), 4(0.138186), 4(0.1172556), 4(0.1213056), 4(0.1042956), 4(0.1119096), 4(0.123336), 4(0.1305288),
		4(0.124578), 4(0.108), 4(0.098442), 4(0.0756108), 4(0.1065096), 4(0.1281528), 4(0.1286388), 4(0.1359828), 4(0.1321704), 4(0.179982), 4(0.1339956), 4(0.16038),
		4(0.1565028), 4(0.1752732), 4(0.1635012), 4(0.1387584), 4(0.1272348), 4(0.1133676), 4(0.1060452), 4(0.102924), 4(0.0987984), 4(0.0963684), 4(0.092124), 4(0.0866376),
		4(0.0490752), 4(0.0192888), 4(0.0036072), 4(0.0), 4(-8.64E-05), 4(-0.0011772), 4(0.0134352), 4(-0.0001944), 4(0.01593), 4(0.1086156), 4(0.1355724), 4(0.1884384),
		4(0.2259144), 4(0.2191968), 4(0.194346), 4(0.1416744), 4(0.1329588), 4(0.1122444), 4(0.105408), 4(0.0995544), 4(0.0977076), 4(0.0972756), 4(0.094446), 4(0.079866),
		4(0.0787212), 4(0.0717768), 4(0.0364176), 4(0.021546), 4(0.016308), 4(0.0138996), 4(0.008532), 4(0.0115236), 4(0.0597672), 4(0.0795636), 4(0.1052568), 4(0.1294488),
		4(0.1887192), 4(0.2116368), 4(0.1651104), 4(0.1423548), 4(0.1216728), 4(0.1251072), 4(0.1106568), 4(0.1060992), 4(0.1022112), 4(0.1041984), 4(0.115398), 4(0.1387908),
		4(0.1447308), 4(0.1512864), 4(0.1352376), 4(0.1192968), 4(0.1111644), 4(0.0945324), 4(0.0956124), 4(0.09369), 4(0.0995652), 4(0.12123), 4(0.128574), 4(0.1542132),
		4(0.1693008), 4(0.18414), 4(0.1525824), 4(0.1401192), 4(0.1097064), 4(0.1121904), 4(0.0989388), 4(0.09423), 4(0.092934), 4(0.0933768), 4(0.09693), 4(0.1155384),
		4(0.1243836), 4(0.1200204), 4(0.0915084), 4(0.092826), 4(0.0928044), 4(0.0939708), 4(0.0866592), 4(0.0844344), 4(0.0944352), 4(0.1188432), 4(0.1055268), 4(0.1377324),
		4(0.1460916), 4(0.1474524), 4(0.1412208), 4(0.1289844), 4(0.1089504), 4(0.1065312), 4(0.0933984), 4(0.0898668), 4(0.0884088), 4(0.0888084), 4(0.1027512), 4(0.1169964),
		4(0.1215108), 4(0.1180332), 4(0.1012284), 4(0.083376), 4(0.0748872), 4(0.0638064), 4(0.04563), 4(0.0364284), 4(0.0563652), 4(0.0715716), 4(0.0873504), 4(0.1155816),
		4(0.1312416), 4(0.1470204), 4(0.1511892), 4(0.133056), 4(0.1130112), 4(0.1089828), 4(0.1033884), 4(0.096228), 4(0.0925344), 4(0.094284), 4(0.1059912), 4(0.1124928),
		4(0.1032264), 4(0.1032048), 4(0.0900288), 4(0.0736344), 4(0.064908), 4(0.0485352), 8(0.0414828), 4(0.0599076), 4(0.0819072), 4(0.0999), 4(0.11745), 4(0.1283688),
		4(0.1516104), 4(0.1534032), 4(0.1318248), 4(0.1157976), 4(0.1107864), 4(0.1042092), 4(0.0983448), 4(0.0939816), 4(0.0947268), 4(0.1011852), 4(0.1112616), 4(0.109944),
		4(0.1046736), 4(0.0960012), 4(0.0843588), 4(0.0724896), 4(0.0641736), 4(0.042822), 4(0.0346032), 4(0.077652), 4(0.1113696), 4(0.134028), 4(0.159894), 4(0.167292),
		4(0.1526472), 4(0.13824), 4(0.1301184), 4(0.1221372), 4(0.1221696), 4(0.1123092), 4(0.110484), 4(0.1019844), 4(0.0973404), 4(0.0948888), 4(0.0898668), 4(0.0926316),
		4(0.0873936), 4(0.0626076), 4(0.0196452), 4(0.00324), 4(0.0002376), 8(0.0), 4(0.0002376), 4(0.0390312), 4(0.1000836), 4(0.1085832), 4(0.115506), 4(0.1379808),
		4(0.1350756), 4(0.1348812), 4(0.1282392), 4(0.1221156), 4(0.1147932), 4(0.112374), 4(0.1097604), 4(0.1064124), 4(0.1026216), 4(0.097308), 4(0.0930636), 4(0.0784512),
		4(0.0241596), 4(0.0046224), 4(5.4E-05), 16(0.0), 4(0.0023436), 4(0.0706428), 4(0.1156032), 4(0.12042), 4(0.1377432), 4(0.1392444), 4(0.1370952), 4(0.1259496),
		4(0.1212948), 4(0.1081188), 4(0.100278), 4(0.0963144), 4(0.0985284), 4(0.1117044), 4(0.1222776), 4(0.1216296), 4(0.1069092), 4(0.0902016), 4(0.0821448), 4(0.0802116),
		4(0.079218), 4(0.0714852), 4(0.0639576), 4(0.0804708), 4(0.120906), 4(0.129384), 4(0.1402596), 4(0.1705644), 4(0.2698272), 4(0.2057832), 4(0.1403028), 4(0.128034),
		4(0.1134), 4(0.1056564), 4(0.096444), 4(0.0920484), 4(0.0905256), 4(0.0976536), 4(0.1151604), 4(0.11934), 4(0.1141452), 4(0.0955476), 4(0.0771336), 4(0.0666144),
		4(0.0662364), 4(0.0532764), 4(0.0603612), 4(0.093204), 4(0.119556), 4(0.1280124), 4(0.1289952), 4(0.169776), 4(0.1799928), 4(0.1607256), 4(0.1293732), 4(0.115344),
		4(0.1033776), 4(0.0960768), 4(0.0887868), 4(0.0847044), 4(0.0849312), 4(0.0909144), 4(0.1100844), 4(0.1174068), 4(0.1167264), 4(0.1069848), 4(0.0921564), 4(0.0912924),
		4(0.092772), 4(0.0919188), 4(0.0991764), 4(0.1137888), 4(0.117558), 4(0.1215324), 4(0.1491048), 4(0.1629288), 4(0.1708128), 4(0.1590732), 4(0.1402164), 4(0.1337256),
		4(0.1199448), 4(0.108594), 4(0.0995544), 4(0.0976104), 4(0.0983124), 4(0.102762), 4(0.127008), 4(0.1325484), 4(0.1143936), 4(0.100548), 4(0.0918), 4(0.0832356),
		4(0.0757836), 4(0.06777), 4(0.0670788), 4(0.0744012), 4(0.115884), 4(0.1212192), 4(0.1259604), 4(0.1470312), 4(0.1611036), 4(0.1453032), 4(0.1350756), 4(0.1233144),
		4(0.1162404), 4(0.1071036), 4(0.1037988), 4(0.1025352), 4(0.1034856), 4(0.113346), 4(0.1238328), 4(0.1238652), 4(0.118044), 4(0.1041984), 4(0.0887868), 4(0.0885384),
		4(0.0864), 4(0.0788616), 4(0.076896), 4(0.0784944), 4(0.1206792), 4(0.1259928), 4(0.1369656), 4(0.1487808), 4(0.167238), 4(0.1630476), 4(0.1398816), 4(0.1346112),
		4(0.1253448), 4(0.1143612), 4(0.1140804), 4(0.1131948), 4(0.1085076), 4(0.1195128), 4(0.0999216), 4(0.0894132), 4(0.08181), 4(0.0543996), 4(0.0108), 4(0.000702),
		4(0.0), 4(-1.08E-05), 4(0.0), 4(0.011556), 4(0.083268), 4(0.1204308), 4(0.152766), 4(0.1486836), 4(0.1716012), 4(0.1554984), 4(0.1422252), 4(0.139104),
		4(0.1324512), 4(0.1087452), 4(0.1015524), 4(0.1168884), 4(0.1063044), 4(0.1143936), 4(0.102762), 4(0.0783), 4(0.0729), 4(0.0387288), 4(0.007992), 4(0.0020196),
		4(0.0), 4(-1.08E-05), 4(0.0), 4(0.008856), 4(0.0770904), 4(0.1126224), 4(0.1337688), 4(0.1530252), 4(0.1504224), 4(0.1490724), 4(0.1397196), 4(0.1353024),
		4(0.1188756), 4(0.0903852), 4(0.0857304), 4(0.084996), 4(0.1062936), 4(0.116694), 4(0.129114), 4(0.128466), 4(0.1157328), 4(0.100062), 4(0.0910872), 4(0.0889272),
		4(0.0922104), 4(0.093582), 4(0.0813132), 4(0.083484), 4(0.1195776), 4(0.123012), 4(0.1785456), 4(0.2618892), 4(0.1650672), 4(0.1500228), 4(0.1317492), 4(0.123336),
		4(0.1198476), 4(0.111888), 4(0.1070928), 4(0.1060776), 4(0.1067688), 4(0.1103868), 4(0.121014), 4(0.118854), 4(0.108108), 4(0.1104516), 4(0.0917028), 4(0.0775008),
		4(0.0584064), 4(0.0771336), 4(0.0931176), 4(0.1044576), 4(0.115884), 4(0.1167048), 4(0.1890108), 4(0.2402892), 4(0.1754892), 4(0.1508436), 4(0.1356264), 4(0.1235196),
		4(0.1188864), 4(0.118962), 4(0.1160244), 4(0.11286), 4(0.1170936), 4(0.1198908), 4(0.123552), 4(0.1251396), 4(0.10422), 4(0.0911412), 4(0.092394), 4(0.1002996),
		4(0.1063584), 4(0.1061424), 4(0.1061856), 4(0.08883), 4(0.1239192), 4(0.1787616), 4(0.2854656), 4(0.398628), 4(0.4804272), 4(0.1721088), 4(0.1566324), 4(0.13878),
		4(0.1209708), 4(0.1177308), 4(0.113346), 4(0.112212), 4(0.1119528), 4(0.1116936), 4(0.119124), 4(0.1251504), 4(0.1225152), 4(0.1044036), 4(0.0979668), 4(0.0928476),
		4(0.0901044), 4(0.1005696), 4(0.1140372), 4(0.1066932), 4(0.1181844), 4(0.125766), 4(0.2029968), 4(0.3079404), 4(0.2915676), 4(0.2006208), 4(0.1465668), 4(0.12204),
		4(0.1231092), 4(0.1187892), 4(0.115398), 4(0.1139832), 4(0.1163052), 4(0.1242648), 4(0.129438), 4(0.124146), 4(0.1254744), 4(0.1117584), 4(0.112806), 4(0.1030644),
		4(0.1017252), 4(0.1113588), 4(0.1166184), 4(0.1194372), 4(0.140724), 4(0.1522584), 4(0.3404592), 4(0.510408), 4(0.5089608), 4(0.2201256), 4(0.151308), 4(0.1296756),
		4(0.1241568), 4(0.1185084), 4(0.1193508), 4(0.116154), 4(0.11556), 4(0.1164564), 4(0.1171044), 4(0.1135944), 4(0.0973944), 4(0.096444), 4(0.0903096), 4(0.0855468),
		4(0.0751356), 4(0.0724896), 4(0.0754812), 4(0.0893484), 4(0.1319868), 4(0.1819368), 4(0.1296324), 4(0.1445256), 4(0.165132), 4(0.1652076), 4(0.131166), 4(0.1181304),
		4(0.1073088), 4(0.1025244), 4(0.0995436), 4(0.0939276), 4(0.0988632), 4(0.0997812), 4(0.0945), 4(0.0898452), 4(0.0815832), 4(0.0830952), 4(0.0853848), 4(0.0782352),
		4(0.0503928), 4(0.0162432), 4(0.009558), 4(0.0216756), 4(0.0634284), 4(0.0904176), 4(0.1181304), 4(0.1282284), 4(0.1380564), 4(0.1473768), 4(0.1389744), 4(0.1187892),
		4(0.1032048), 4(0.090288), 4(0.0862056), 4(0.0877284), 4(0.0891108), 4(0.09369), 4(0.1125792), 4(0.1263816), 4(0.1265112), 4(0.1220076), 4(0.1134864), 4(0.105462),
		4(0.096606), 4(0.0935928), 4(0.0874152), 4(0.0934956), 4(0.106758), 4(0.1110672), 4(0.1481436), 4(0.1478628), 4(0.1523232), 4(0.1424304), 4(0.1201284), 4(0.1055052),
		4(0.1123308), 4(0.1009692), 4(0.0942408), 4(0.0937548), 4(0.096768), 4(0.1102464), 4(0.1139184), 4(0.1168452), 4(0.1014984), 4(0.0914004), 4(0.077652), 4(0.0622944),
		4(0.0343548), 4(0.0290736), 4(0.0639468), 4(0.0737748), 4(0.0968976), 4(0.106758), 4(0.1316952), 4(0.1355076), 4(0.1717524), 4(0.1509408), 4(0.1256688), 4(0.1129896),
		4(0.1054944), 4(0.101088), 4(0.0940896), 4(0.0945756), 4(0.0971568), 4(0.1081944), 4(0.1146204), 4(0.1203336), 4(0.0942408), 4(0.0735804), 4(0.0575424), 4(0.0437076),
		4(0.0267732), 4(0.0191052), 4(0.011556), 4(0.0307476), 4(0.086454), 4(0.1083456), 4(0.147744), 4(0.2216052), 4(0.1869264), 4(0.1528416), 4(0.126414), 4(0.1158192),
		4(0.1119312), 4(0.1084428), 4(0.083808), 4(0.0798552), 4(0.084456), 4(0.1081944), 4(0.1160028), 4(0.109944), 4(0.1012932), 4(0.088344), 4(0.0800496), 4(0.079704),
		4(0.0688932), 4(0.0549288), 4(0.0422064), 4(0.0672408), 4(0.0867024), 4(0.1121256), 4(0.1342548), 4(0.1381212), 4(0.1514484), 4(0.1485972), 4(0.1384668), 4(0.110916),
		4(0.1135404), 4(0.1060776), 4(0.0983124), 4(0.0939924), 4(0.0995436), 4(0.1082808), 4(0.11367), 4(0.1179036), 4(0.11394), 4(0.0974052), 4(0.0724572), 4(0.0712368),
		4(0.073116), 4(0.0709884), 4(0.056214), 4(0.0570132), 4(0.0814752), 4(0.0968868), 4(0.1303668), 4(0.144666), 4(0.165672), 4(0.1641816), 4(0.1395144), 4(0.1199556),
		4(0.122526), 4(0.1066392), 4(0.103032), 4(0.096822), 4(0.09585), 4(0.09558), 4(0.0940572), 4(0.089046), 4(0.0775224), 4(0.0549288), 4(0.0320544), 4(0.0061344),
		4(0.003186), 12(0.0), 4(0.0061776), 4(0.0699948), 4(0.1038852), 4(0.1246104), 4(0.1494612), 4(0.1344276), 4(0.1197288), 4(0.1017684), 4(0.095526), 4(0.083862),
		4(0.0759456), 4(0.0758808), 4(0.0736128), 4(0.06723), 4(0.0518076), 4(0.0283716), 4(0.0066528), 4(0.0), 4(-0.0010908), 4(-0.002268), 4(-0.00324), 4(-0.010692),
		4(-0.0108864), 4(-0.0053784), 4(-0.0009612), 4(0.0394956), 4(0.0933336), 4(0.1022976), 4(0.1315332), 4(0.1193832), 4(0.1134864), 4(0.0918972), 4(0.0896184), 4(0.0756756),
		4(0.0755676), 4(0.0747576), 4(0.0777924), 4(0.0994896), 4(0.1007964), 4(0.1092528), 4(0.1029132), 4(0.0925344), 4(0.072036), 4(0.053244), 4(0.0158112), 4(0.004374),
		4(0.0007128), 4(0.0428328), 4(0.0724248), 4(0.1031508), 4(0.128088), 4(0.1614816), 4(0.1781676), 4(0.1270404), 4(0.1074816), 4(0.0851796), 4(0.061452), 4(0.0173016),
		4(0.0335556), 4(0.0270432), 4(0.0647676), 4(0.0875988), 4(0.1043928), 4(0.1010232), 4(0.0789588), 4(0.0040932), 4(0.0), 4(-0.0019656), 4(-0.0053676), 4(0.0193104),
		4(-0.01296), 4(0.0035208), 4(0.0650376), 4(0.1025028), 4(0.1197072), 4(0.158976), 4(0.1924884), 4(0.1321704), 4(0.1163592), 4(0.0919944), 4(0.08235), 4(0.064584),
		4(0.0724356), 4(0.0751032), 4(0.0722196), 4(0.0885708), 4(0.1032264), 4(0.105138), 4(0.09072), 4(0.0300564), 4(2.16E-05), 4(0.0023436), 4(0.0112536), 4(0.0130032),
		4(0.0072576), 4(0.0324432), 4(0.0902232), 4(0.0826092), 4(0.110862), 4(0.14283), 4(0.1920996), 4(0.1685556), 4(0.1188), 4(0.1092312), 4(0.1051596), 4(0.1038312),
		4(0.0972972), 4(0.0937008), 4(0.0947052), 4(0.0947484), 4(0.1088856), 4(0.1022544), 4(0.0511704), 4(0.0184032), 4(-0.0021276), 4(0.0), 4(-0.0001836), 4(-0.0034992),
		8(2.16E-05), 4(0.0560196), 4(0.0812052), 4(0.119826), 4(0.1540512), 4(0.19008), 4(0.1396332), 4(0.1188), 4(0.1093824), 4(0.101466), 4(0.097254), 4(0.092988),
		4(0.0895428), 4(0.087534), 4(0.098604), 4(0.105732), 4(0.10341), 4(0.0797364), 4(0.0515268), 4(0.008964), 4(0.0071172), 4(0.0), 4(-1.08E-05), 8(0.0),
		4(0.0113292), 4(0.1089072), 4(0.1307232), 4(0.2210112), 4(0.2701836), 4(0.1662768), 4(0.1353348), 4(0.117126), 4(0.1107756), 4(0.1098576), 4(0.1093176), 4(0.106056),
		4(0.1058724), 4(0.1059696), 4(0.1053864), 4(0.0925344), 4(0.0733644), 4(0.0165672), 4(-2.16E-05), 4(-0.00108), 4(-0.0112428), 4(-0.0178308), 4(-0.0161028), 4(-0.0029376),
		4(0.0001404), 4(0.1256688), 4(0.1277856), 4(0.147744), 4(0.1759428), 4(0.1368576), 4(0.121932), 4(0.1026), 4(0.0914004), 4(0.089478), 4(0.0891324), 4(0.0834624),
		4(0.086292), 4(0.089424), 4(0.087588), 4(0.075006), 4(0.0285768), 4(-1.08E-05), 4(-0.0037908), 4(-0.016848), 4(-0.040986), 4(-0.065124), 4(-0.053622), 4(-0.0213408),
		4(-0.000216), 4(0.0612792), 4(0.0978912), 4(0.1306692), 4(0.1625292), 4(0.1290276), 4(0.1151172), 4(0.1057968), 4(0.1071684), 4(0.098442), 4(0.0938196), 4(0.091152),
		4(0.0998136), 4(0.11178), 4(0.1383372), 4(0.1235952), 4(0.088992), 4(0.0359748), 4(0.003942), 4(0.0027432), 12(0.0), 4(0.00972), 4(0.0638496), 4(0.1064124),
		4(0.1511892), 4(0.2255148), 4(0.2634228), 4(0.151578), 4(0.1175796), 4(0.10368), 4(0.10044), 4(0.0968436), 4(0.0922428), 4(0.0915516), 4(0.0927288), 4(0.1013688),
		4(0.1112076), 4(0.1062072), 4(0.1012068), 4(0.06966), 4(0.016686), 4(0.0142344), 4(0.0090504), 4(0.00324), 4(0.005562), 4(0.037854), 4(0.0789264), 4(0.1226988),
		4(0.1589544), 4(0.2915352), 4(0.3295404), 4(0.1598076), 4(0.1236708), 4(0.106056), 4(0.1043928), 4(0.0972), 4(0.0938412), 4(0.0914868), 4(0.0940356), 4(0.0992844),
		4(0.1173312), 4(0.1118016), 4(0.0965628), 4(0.0675972), 4(-0.0010476), 4(0.0051948), 4(0.0072792), 4(0.0105516), 4(0.044496), 4(0.076572), 4(0.091044), 4(0.1043712),
		4(0.1423548), 4(0.2827332), 4(0.3024756), 4(0.1629936), 4(0.1330668), 4(0.1147716), 4(0.105948), 4(0.09936), 4(0.095526), 4(0.0944892), 4(0.0948996), 4(0.1036908),
		4(0.114372), 4(0.1140804), 4(0.102222), 4(0.091692), 4(0.0690768), 4(0.0608688), 4(0.0477468), 4(0.0395712), 4(0.059292), 4(0.0749844), 4(0.0853092), 4(0.1082484),
		4(0.1595268), 4(0.2783052), 4(0.302832), 4(0.1678968), 4(0.131436), 4(0.114426), 4(0.1070496), 4(0.1056888), 4(0.0997812), 4(0.0950724), 4(0.09747), 4(0.1012932),
		4(0.1066392), 4(0.1069632), 4(0.1008936), 4(0.076302), 4(0.0271944), 4(0.00324), 4(8.64E-05), 8(0.0), 4(0.0018684), 4(0.0396684), 4(0.0890028), 4(0.112968),
		4(0.1316412), 4(0.1474308), 4(0.1201176), 4(0.114156), 4(0.1033668), 4(0.101574), 4(0.0963468), 4(0.0948024), 4(0.0887652), 4(0.086832), 4(0.0897912), 4(0.0926424),
		4(0.0928044), 4(0.0834084), 4(0.0707292), 4(0.0261468), 4(0.004104), 4(0.0001836), 8(-1.08E-05), 4(0.0), 4(0.0336312), 4(0.0784512), 4(0.1110888), 4(0.1409832),
		4(0.1503576), 4(0.1296864), 4(0.1070172), 4(0.0968328), 4(0.0962496), 4(0.0894672), 4(0.0898884), 4(0.088344), 4(0.0886572), 4(0.0896832), 4(0.0897588), 4(0.0794124),
		4(0.0700272), 4(0.0251208), 4(0.0085104), 4(0.000486), 4(7.56E-05), 4(-0.0006912), 4(-0.0008532), 4(0.000702), 4(0.0162972), 4(0.070848), 4(0.102168), 4(0.1183464),
		4(0.1214784), 4(0.1188432), 4(0.1131624), 4(0.1099656), 4(0.0972864), 4(0.0915408), 4(0.0894888), 4(0.087264), 4(0.0926532), 4(0.1038636), 4(0.1221048), 4(0.1274508),
		4(0.1095984), 4(0.0944784), 4(0.0745632), 4(0.0496044), 4(0.0216432), 4(0.0153684), 4(0.0198072), 4(0.0589248), 4(0.078408), 4(0.1063152), 4(0.1248372), 4(0.1927476),
		4(0.2221668), 4(0.1348596), 4(0.115074), 4(0.10692), 4(0.1082484), 4(0.1004724), 4(0.0934956), 4(0.0911412), 4(0.094662), 4(0.107838), 4(0.11718), 4(0.116748),
		4(0.105894), 4(0.0956556), 4(0.0752112), 4(0.0466884), 4(0.0322704), 4(0.0410184), 4(0.0458892), 4(0.062154), 4(0.0813456), 4(0.1165104), 4(0.1353024), 4(0.1965816),
		4(0.1798848), 4(0.12447), 4(0.112752), 4(0.1057968), 4(0.1039068), 4(0.09855), 4(0.0925776), 4(0.0904824), 4(0.0944244), 4(0.1039284), 4(0.1170288), 4(0.1152144),
		4(0.1107756), 4(0.0854712), 4(0.0685584), 4(0.0496908), 4(0.0509112), 4(0.0378), 4(0.0441936), 4(0.0734832), 4(0.0816264), 4(0.108918), 4(0.1242432), 4(0.1416852),
		4(0.141588), 4(0.1269756), 4(0.1184868), 4(0.10854), 4(0.1003428), 4(0.0889596), 4(0.0889812), 4(0.0913248), 4(0.0920376), 4(0.1071468), 4(0.1159488), 4(0.116586),
		4(0.1103868), 4(0.1104948), 4(0.0993924), 4(0.0908712), 4(0.081594), 4(0.0765936), 4(0.0845424), 4(0.0920916), 4(0.1040688), 4(0.1174392), 4(0.1227852), 4(0.139212),
		4(0.1449468), 4(0.1272888), 4(0.1077516), 4(0.0973404), 4(0.0931824), 4(0.084294), 4(0.080514), 4(0.0785376), 4(0.0771336), 4(0.0883224), 4(0.1097928), 4(0.1111752),
		4(0.0999864), 4(0.0854604), 4(0.0674352), 4(0.0444852), 4(0.0181548), 4(0.0063828), 4(0.002376), 4(0.0068796), 4(0.0500148), 4(0.0769608), 4(0.0993816), 4(0.1111752),
		4(0.1211436), 4(0.1157868), 4(0.1110996), 4(0.1019196), 4(0.1029564), 4(0.0964656), 4(0.0937764), 4(0.09099), 4(0.0910008), 4(0.0914868), 4(0.0932148), 4(0.0936576),
		4(0.0893916), 4(0.0561708), 4(0.0136512), 4(0.003618), 4(0.0014904), 4(0.0001296), 4(0.0004752), 4(0.0038016), 4(0.0161028), 4(0.0949212), 4(0.11961), 4(0.1299672),
		4(0.1430676), 4(0.1295676), 4(0.1200528), 4(0.1143612), 4(0.10854), 4(0.1027188), 4(0.101088), 4(0.0984528), 4(0.0972756), 4(0.0975348), 4(0.0972), 4(0.0913896),
		4(0.0492804), 4(0.0023112), 4(-1.08E-05), 4(-7.56E-05), 4(-0.0021384), 4(-0.008046), 4(-0.007992), 4(-0.000108), 4(0.0), 4(0.0745524), 4(0.111132), 4(0.1190052),
		4(0.1265544), 4(0.1234656), 4(0.1161), 4(0.1085616), 4(0.1029024), 4(0.0939924), 4(0.0890676), 4(0.0857736), 4(0.0867456), 4(0.107298), 4(0.12069), 4(0.1304856),
		4(0.116316), 4(0.0993276), 4(0.0734616), 4(0.0378216), 4(0.0108), 4(0.0064044), 4(0.0073224), 4(0.027216), 4(0.0745092), 4(0.0971784), 4(0.1213812), 4(0.1643868),
		4(0.2321028), 4(0.1470636), 4(0.1242432), 4(0.113562), 4(0.112644), 4(0.1100736), 4(0.1075032), 4(0.1061424), 4(0.1086696), 4(0.1091124), 4(0.1281636), 4(0.12933),
		4(0.1141884), 4(0.0972), 4(0.0625104), 4(0.050706), 4(0.0335988), 4(0.0283824), 4(0.041094), 4(0.0801792), 4(0.0985392), 4(0.1215756), 4(0.1410696), 4(0.1973484),
		4(0.1938816), 4(0.1351944), 4(0.1184976), 4(0.1075464), 4(0.1070928), 4(0.09747), 4(0.0937332), 4(0.0956988), 4(0.0993708), 4(0.1079136), 4(0.1183896), 4(0.1245996),
		4(0.1227312), 4(0.1097604), 4(0.0743688), 4(0.0643356), 4(0.0582552), 4(0.0422172), 4(0.0506736), 4(0.0843372), 4(0.0943704), 4(0.116424), 4(0.1400436), 4(0.2202228),
		4(0.2212164), 4(0.136296), 4(0.1227204), 4(0.1118556), 4(0.104922), 4(0.0995112), 4(0.0951588), 4(0.095796), 4(0.1001052), 4(0.1042956), 4(0.1260036), 4(0.1299456),
		4(0.1062612), 4(0.029592), 4(0.0138672), 4(0.0003348), 4(0.0001404), 4(0.0001188), 4(0.0174528), 4(0.041256), 4(0.0967572), 4(0.1228392), 4(0.1542024), 4(0.17901),
		4(0.1546992), 4(0.1292976), 4(0.1138644), 4(0.098226), 4(0.0921564), 4(0.0942408), 4(0.093906), 4(0.0953208), 4(0.0980748), 4(0.107244), 4(0.1150092), 4(0.1181088),
		4(0.1187568), 4(0.1012824), 4(0.0864108), 4(0.0636984), 4(0.0523152), 4(0.0518508), 4(0.06426), 4(0.0898452), 4(0.1021896), 4(0.1253232), 4(0.1316736), 4(0.1583172),
		4(0.1521504), 4(0.1255824), 4(0.1086804), 4(0.0977076), 4(0.1025028), 4(0.0968328), 4(0.0924264), 4(0.0880308), 4(0.0945756), 4(0.1008936), 4(0.0983664), 4(0.100008),
		4(0.0945648), 4(0.08991), 4(0.041742), 4(0.0056484), 12(0.0), 4(0.0103356), 4(0.06912), 4(0.1111428), 4(0.1403244), 4(0.1409292), 4(0.1352808), 4(0.120528),
		4(0.1060776), 4(0.0908604), 4(0.0856764), 4(0.0759348), 4(0.0680832), 4(0.0641412), 4(0.0608688), 4(0.0760752), 4(0.0766476), 4(0.0724464), 4(0.0240948), 4(0.0058212),
		4(1.08E-05), 4(-1.08E-05), 4(-0.000108), 4(-0.0010584), 4(-0.000648), 4(0.0), 4(0.030024), 4(0.0945432), 4(0.1216944), 4(0.1385316), 4(0.1365552), 4(0.1198692),
		4(0.1080108), 4(0.09585), 4(0.0969516), 4(0.0968112), 4(0.0954072), 4(0.0943488), 4(0.0963144), 4(0.1070496), 4(0.1234008), 4(0.128142), 4(0.1157544), 4(0.1080432),
		4(0.0664956), 4(0.0680292), 4(0.0436752), 4(0.0244944), 4(0.041256), 4(0.0772308), 4(0.0893484), 4(0.1196316), 4(0.1857816), 4(0.2346516), 4(0.212058), 4(0.136728),
		4(0.1164672), 4(0.1057212), 4(0.0926316), 4(0.0898236), 4(0.0930096), 4(0.0931068), 4(0.0956664), 4(0.1035288), 4(0.1270404), 4(0.1475064), 4(0.1280124), 4(0.0709884),
		4(0.0660312), 4(0.062964), 4(0.066798), 4(0.0583308), 4(0.0742932), 4(0.079974), 4(0.1011096), 4(0.1198476), 4(0.178308), 4(0.2984796), 4(0.2524068), 4(0.1359072),
		4(0.1167048), 4(0.1117692), 4(0.1128816), 4(0.0878148), 4(0.0844236), 4(0.0785268), 4(0.0828684), 4(0.0997812), 4(0.1169856), 4(0.1197612), 4(0.1093716), 4(0.0844128),
		4(0.0385668), 4(0.0088884), 4(0.0064908), 4(0.0067608), 4(0.012582), 4(0.080136), 4(0.1025676), 4(0.129438), 4(0.1508436), 4(0.1916244), 4(0.1670868), 4(0.1346652),
		4(0.1231308), 4(0.1146096), 4(0.1114992), 4(0.1050732), 4(0.1006668), 4(0.09288), 4(0.087102), 4(0.1057536), 4(0.125334), 4(0.1277748), 4(0.1141668), 4(0.0795636),
		4(0.0416664), 4(0.0062532), 4(0.003456), 4(0.0034128), 4(0.0332316), 4(0.0673596), 4(0.0984312), 4(0.127278), 4(0.1856952), 4(0.3272724), 4(0.2477304), 4(0.1391688),
		4(0.121014), 4(0.1136052), 4(0.1053864), 4(0.0918216), 4(0.0890136), 8(0.087588), 4(0.1003644), 4(0.1224828), 4(0.1366524), 4(0.1304424), 4(0.1102464), 4(0.0993816),
		4(0.097416), 4(0.0900504), 4(0.082728), 4(0.0814104), 4(0.0889812), 4(0.1041768), 4(0.1378512), 4(0.1486188), 4(0.1789128), 4(0.1654668), 4(0.1353564), 4(0.1314684),
		4(0.1117476), 4(0.1114668), 4(0.1121472), 4(0.1123308), 4(0.1119636), 4(0.1110024), 4(0.1117908), 4(0.100494), 4(0.0984312), 4(0.108162), 4(0.09099), 4(0.0130788),
		4(0.0), 4(-2.16E-05), 4(-0.0009288), 4(-0.0010692), 4(-1.08E-05), 4(0.0502416), 4(0.113994), 4(0.1474416), 4(0.1770012), 4(0.1669356), 4(0.1444716), 4(0.1326672),
		4(0.0921456), 4(0.0880632), 4(0.0820908), 4(0.0779868), 4(0.0805032), 4(0.0799632), 4(0.0797256), 4(0.078192), 4(0.0539892), 4(0.0), 4(-9.72E-05), 4(-0.00432),
		4(-0.0216972), 4(-0.0432216), 4(-0.057672), 4(-0.0437616), 4(-0.0214056), 4(-0.0013176), 4(0.0628344), 4(0.1138752), 4(0.155412), 4(0.1439532), 4(0.1284336), 4(0.1154304),
		4(0.101034), 4(0.0932148), 4(0.0950832), 4(0.0944892), 4(0.0954504), 4(0.0971676), 4(0.1091448), 4(0.1326996), 4(0.152874), 4(0.1329696), 4(0.1096416), 4(0.09261),
		4(0.0804168), 4(0.0693144), 4(0.0674784), 4(0.0777924), 4(0.0887004), 4(0.112428), 4(0.1440828), 4(0.220644), 4(0.4345812), 4(0.324864), 4(0.1563516), 4(0.1446228),
		4(0.1303344), 4(0.1172556), 4(0.1099872), 4(0.109728), 4(0.10962), 4(0.109674), 4(0.1178388), 4(0.1933632), 4(0.2904876), 4(0.1942488), 4(0.130086), 4(0.1123956),
		4(0.10449), 4(0.0924588), 4(0.0926532), 4(0.0978048), 4(0.1064448), 4(0.118476), 4(0.1529172), 4(0.2284632), 4(0.4141368), 4(0.2348568), 4(0.1481004), 4(0.1352484),
		4(0.1256364), 4(0.1052892), 4(0.0994032), 4(0.0979128), 4(0.0980424), 4(0.0970704), 4(0.1056024), 4(0.1359828), 4(0.2188404), 4(0.1539), 4(0.1290384), 4(0.125712),
		4(0.1230768), 4(0.1085184), 4(0.1033776), 4(0.11043), 4(0.1105056), 4(0.126468), 4(0.1398816), 4(0.1782432), 4(0.2774736), 4(0.1759644), 4(0.1263384), 4(0.1052028),
		4(0.0919728), 4(0.0889164), 4(0.0832464), 4(0.0747468), 4(0.0768636), 4(0.0815292), 4(0.1068768), 4(0.135432), 4(0.146124), 4(0.1241352), 4(0.11853), 4(0.0859248),
		4(0.088668), 4(0.0951804), 4(0.0963576), 4(0.0906876), 4(0.1092528), 4(0.1655532), 4(0.161352), 4(0.1674648), 4(0.2125224), 4(0.1584576), 4(0.1357452), 4(0.128142),
		4(0.1159164), 4(0.08721), 4(0.0774792), 4(0.0737208), 4(0.0738612), 4(0.076464), 4(0.1169208), 4(0.1486944), 4(0.1574748), 4(0.139698), 4(0.1020816), 4(0.0672192),
		4(0.0574668), 4(0.047304), 4(0.0592164), 4(0.0684396), 4(0.0917784), 4(0.1134), 4(0.1579392), 4(0.1558548), 4(0.2587356), 4(0.1702728), 4(0.1234872), 4(0.1149768),
		4(0.1011096), 4(0.096012), 4(0.080298), 4(0.072252), 4(0.074034), 4(0.0797472), 4(0.08343), 4(0.0946296), 4(0.0837432), 4(0.0709776), 4(0.0609444), 4(0.0148608),
		4(0.0025596), 12(0.0), 4(1.08E-05), 4(0.0906228), 4(0.1221156), 4(0.130572), 4(0.1434996), 4(0.1292112), 4(0.1107), 4(0.1089072), 4(0.0983988), 4(0.0882792),
		4(0.0777168), 4(0.0787212), 4(0.0838944), 4(0.090018), 4(0.0977508), 4(0.0976428), 4(0.1017792), 4(0.096876), 4(0.0805788), 4(0.0567108), 4(0.01809), 4(0.0064044),
		4(0.0), 4(-1.08E-05), 4(0.0), 4(0.0218484), 4(0.09477), 4(0.1365012), 4(0.1884924), 4(0.1353348), 4(0.0953532), 4(0.0811836), 4(0.034344), 4(0.0627372),
		4(0.0462888), 4(0.051678), 4(0.0491184), 4(0.0495288), 4(0.0818532), 4(0.1369224), 4(0.153846), 4(0.1176336), 4(0.068094), 4(0.0139752), 4(0.0094608), 4(0.0073548),
		4(0.0079596), 4(0.0097416), 4(0.0347652), 4(0.100494), 4(0.1305612), 4(0.1646028), 4(0.2120364), 4(0.1541376), 4(0.1421928), 4(0.1278396), 4(0.1211652), 4(0.1188),
		4(0.1095552), 4(0.0971892), 4(0.0976968), 4(0.0990792), 4(0.1087992), 4(0.1271916), 4(0.1418364), 4(0.1350108), 4(0.0979668), 4(0.1011852), 4(0.0575208), 4(0.088074),
		4(0.07857), 4(0.060588), 4(0.099576), 4(0.1183572), 4(0.1818828), 4(0.1750572), 4(0.2438856), 4(0.1561032), 4(0.1332504), 4(0.1225908), 4(0.0931716), 4(0.0876096),
		4(0.0686448), 4(0.05508), 4(0.0507816), 4(0.0610956), 4(0.0904392), 4(0.1231416), 4(0.1347192), 4(0.1216296), 4(0.1008936), 4(0.073818), 4(0.0471528), 4(0.0137268),
		4(0.0096768), 4(0.0134784), 4(0.0524124), 4(0.09369), 4(0.1133892), 4(0.1575504), 4(0.2139372), 4(0.1597536), 4(0.114804), 4(0.10638), 4(0.080514), 4(0.062748),
		4(0.0543888), 4(0.0425304), 4(0.043038), 4(0.0548208), 4(0.0846072), 4(0.1183032), 4(0.1257876), 4(0.100386), 4(0.0878364), 4(0.0657396), 4(0.005886), 4(0.0001944),
		8(0.0), 4(0.0005184), 4(0.0727812), 4(0.1296648), 4(0.158274), 4(0.2404404), 4(0.1616112), 4(0.1188), 4(0.1122552), 4(0.095256), 4(0.0800172), 4(0.0774684),
		4(0.0767124), 4(0.076248), 4(0.0762048), 4(0.0984204), 4(0.1245888), 4(0.1485324), 4(0.118476), 4(0.089802), 4(0.0535464), 4(0.0134352), 4(0.0010692), 8(0.0),
		4(0.0129276), 4(0.086292), 4(0.1228284), 4(0.2646648), 4(0.4275612), 4(0.1723896), 4(0.1162404), 4(0.1088856), 4(0.0867132), 4(0.1031508), 4(0.0917568), 4(0.0873288),
		4(0.08721), 4(0.0871344), 4(0.0936792), 4(0.102762), 4(0.1012608), 4(0.0878688), 4(0.0269028), 4(-6.48E-05), 4(-0.0009936), 4(-0.0082512), 4(-0.0099144), 4(-0.0044388),
		4(0.000216), 4(0.035316), 4(0.1202148), 4(0.1439532), 4(0.1590408), 4(0.1135296), 4(0.091098), 4(0.0837972), 4(0.0549828), 4(0.0308124), 4(0.0162972), 4(0.0076788),
		4(0.00675), 4(0.0060156), 4(0.0162216), 4(0.0047628), 4(0.0056484), 4(0.0036396), 4(0.000162), 4(0.0002808), 4(-0.0107244), 4(-0.0153684), 4(-0.0153144), 4(-0.003294),
		4(-5.4E-05), 4(0.0102276), 4(0.1020168), 4(0.1085724), 4(0.1221048), 4(0.122526), 4(0.1062612), 4(0.1080432), 4(0.0909792), 4(0.0825984), 4(0.078786), 4(0.0760968),
		4(0.0744444), 4(0.0742932), 4(0.0893808), 4(0.1210032), 4(0.1334664), 4(0.1137996), 4(0.0994896), 4(0.070254), 4(0.0389232), 4(0.052812), 4(0.0392148), 4(0.0638172),
		4(0.0730836), 4(0.0939168), 4(0.1230552), 4(0.1426464), 4(0.2384208), 4(0.146934), 4(0.1176444), 4(0.1114452), 4(0.0988524), 4(0.0848556), 4(0.0842832), 4(0.0831168),
		4(0.08289), 4(0.0864432), 4(0.1043496), 4(0.1272888), 4(0.1743984), 4(0.1552824), 4(0.1128708), 4(0.0788076), 4(0.0907848), 4(0.0831924), 4(0.080676), 4(0.0836676),
		4(0.1017036), 4(0.1199016), 4(0.147096), 4(0.2131812), 4(0.3071952), 4(0.1736964), 4(0.124254), 4(0.117558), 4(0.10125), 4(0.0936252), 4(0.083754), 4(0.0831384),
		4(0.0755568), 4(0.0933012), 4(0.1062828), 4(0.1361556), 4(0.1363824), 4(0.1237248), 4(0.1157868), 4(0.118692), 4(0.1044792), 4(0.0871236), 4(0.0786024), 4(0.0952776),
		4(0.1093932), 4(0.1175148), 4(0.139698), 4(0.1697328), 4(0.2123172), 4(0.1445796), 4(0.1106892), 4(0.0973728), 4(0.0833652), 4(0.0777816), 4(0.076626), 4(0.0708804),
		4(0.06912), 4(0.0704484), 4(0.0855684), 4(0.1162404), 4(0.1383048), 4(0.1346976), 4(0.1101168), 4(0.1086372), 4(0.108972), 4(0.1170612), 4(0.094338), 4(0.095472),
		4(0.1007748), 4(0.112536), 4(0.1278612), 4(0.1292328), 4(0.1483272), 4(0.1333908), 4(0.1194804), 4(0.1092204), 4(0.0875772), 4(0.0847584), 4(0.0812808), 4(0.0790344),
		4(0.0791532), 4(0.081594), 4(0.0895644), 4(0.1201392), 4(0.130626), 4(0.135756), 4(0.1283256), 4(0.1155708), 4(0.1126116), 4(0.110214), 4(0.1050624), 4(0.1039176),
		4(0.1070604), 4(0.111456), 4(0.1222776), 4(0.131976), 4(0.142506), 4(0.1291788), 4(0.1147068), 4(0.104652), 4(0.097092), 4(0.0918864), 4(0.0918648), 4(0.091854),
		4(0.091962), 4(0.0957852), 4(0.1001052), 4(0.0948024), 4(0.1089936), 4(0.1145664), 4(0.1060236), 4(0.1005588), 4(0.0880848), 4(0.0704592), 4(0.0411804), 4(0.056052),
		4(0.0906984), 4(0.108108), 4(0.116964), 4(0.1370628), 4(0.1540728), 4(0.1331964), 4(0.1216836), 4(0.1145556), 4(0.1095336), 4(0.1089504), 4(0.106596), 4(0.0993492),
		4(0.099468), 4(0.0983664), 4(0.099144), 4(0.101574), 4(0.107082), 4(0.1004724), 4(0.0990144), 4(0.0934092), 4(0.0413208), 4(0.0184788), 4(0.0092124), 4(0.01404),
		4(0.0682128), 4(0.1161432), 4(0.140724), 4(0.1449468), 4(0.1676916), 4(0.1495368), 4(0.1350216), 4(0.1247616), 4(0.1067796), 4(0.1024812), 4(0.1003752), 4(0.0995868),
		4(0.1000728), 4(0.0999756), 4(0.1110348), 4(0.1501524), 4(0.2378484), 4(0.170154), 4(0.1240596), 4(0.0999324), 4(0.0954072), 4(0.0886464), 4(0.0872316), 4(0.0953532),
		4(0.0993276), 4(0.1150416), 4(0.1596996), 4(0.336852), 4(0.4232628), 4(0.181818), 4(0.1384884), 4(0.1234764), 4(0.112536), 4(0.1080972), 4(0.10179), 4(0.10368),
		4(0.1070604), 4(0.1053108), 4(0.1181196), 4(0.1588572), 4(0.2841588), 4(0.2259684), 4(0.1509408), 4(0.1291896), 4(0.1101168), 4(0.1014012), 4(0.100656), 4(0.1039176),
		4(0.111186), 4(0.169668), 4(0.2632932), 4(0.3780648), 4(0.3876876), 4(0.1838376), 4(0.1418148), 4(0.1209276), 4(0.1133244), 0.1176984, 0.1049004, 0.1022004,
		0.1020168, 0.0994572, 0.098496, 0.0972864, 0.0966492, 0.1020168, 0.1018656, 0.1025136, 0.102708, 2(0.1000296), 0.1016172, 0.104544,
		0.0976752, 0.0990036, 0.0951048, 0.1050408, 0.09747, 0.1049328, 0.1107864, 0.1254096, 0.1078596, 0.1275264, 0.1438884, 0.160542,
		0.1744524, 0.1942812, 0.1903932, 0.1838268, 0.2056968, 0.1525716, 0.1267488, 0.10287, 0.1481868, 0.1134108, 0.101034, 0.087642,
		0.1117476, 0.103032, 0.0897372, 0.0739368, 0.1107864, 0.1032588, 0.0964224, 0.0984096, 0.1004724, 0.0957204, 0.095256, 0.0957204,
		0.0962928, 0.099846, 0.1029672, 0.1054944, 0.0981936, 0.1029888, 0.1093608, 0.1115856, 0.1092204, 0.1101924, 0.1172988, 0.1233252,
		0.1030644, 0.1108404, 0.1180116, 0.141588, 0.0972108, 0.128628, 0.1557252, 0.2078136, 0.1522476, 0.2071764, 0.286524, 0.3740796,
		0.3946968, 0.3669516, 0.3216564, 0.2560356, 0.2248668, 0.1646892, 0.1406484, 0.118098, 0.1419012, 0.13122, 0.111402, 0.1049976,
		0.119016, 0.1114992, 0.103194, 0.0972432, 0.1028376, 0.1007532, 0.0987336, 0.0940248, 0.107838, 0.1001808, 0.0955152, 0.0980532,
		0.1042416, 0.1008612, 0.0935388, 0.0902556, 0.0940896, 0.0946836, 0.0973296, 0.1021788, 0.1022652, 2(0.1022004), 0.102114, 0.1012068,
		0.1042092, 0.104436, 0.1044684, 0.096444, 0.0999972, 0.1069848, 0.1239948, 0.1036692, 0.1272564, 0.143046, 0.17955, 0.1791936,
		0.207252, 0.200556, 0.1771092, 0.1978668, 0.1599156, 0.1201176, 0.0903528, 0.1381752, 0.1273644, 0.108162, 0.0947052, 0.1228284,
		0.1167804, 0.1018548, 0.0940356, 0.1076328, 0.0988092, 0.0917568, 0.087912, 0.0979884, 0.0909144, 0.0873288, 0.0871668, 0.0857088,
		0.0867456, 0.0921996, 0.0960768, 0.0901692, 0.099036, 0.0997164, 0.1002132, 0.089856, 0.0997704, 0.1118232, 0.124362, 0.1047492,
		0.1313172, 0.1454436, 0.1568592, 0.1152036, 0.129654, 0.1487376, 0.1744308, 0.1295136, 0.1557252, 0.1912032, 0.2399112, 0.2334312,
		0.2184084, 0.1760724, 0.1458972, 0.1684584, 0.1434996, 0.1309068, 0.1161432, 0.1353564, 0.1268676, 0.1066716, 0.0984312, 0.1247184,
		0.1180008, 0.106704, 0.0996516, 0.1130112, 0.1004508, 0.0868428, 0.0863568, 0.0998892, 0.0899532, 0.0836028, 0.0741744, 0.0889272,
		0.0825012, 0.0749628, 0.0645192, 0.0826848, 0.0809136, 0.0779544, 0.0773172, 0.069984, 0.0884088, 0.0915192, 0.0865404, 0.0818208,
		0.082458, 0.0914544, 0.0942732, 0.0842724, 0.088884, 0.1003968, 0.1227852, 0.1029132, 0.1215972, 0.1445256, 0.160542, 0.1543536,
		0.1549692, 0.1495044, 0.140562, 0.1559412, 0.1398384, 0.1335636, 0.1174716, 0.1315548, 0.1192536, 0.1061316, 0.094068, 0.1159272,
		0.105678, 0.0879552, 0.0579636, 0.058806, 0.0549288, 0.0512676, 0.0431676, 0.0487728, 0.0444096, 0.0401868, 0.0350676, 0.0293652,
		0.0250776, 0.0278964, 0.0329616, 0.0209844, 0.030402, 0.0673704, 0.0730836, 0.0356076, 0.0785268, 0.0981396, 0.1111104, 0.0897804,
		0.095742, 0.1120824, 0.1355508, 0.0998028, 0.113832, 0.1480356, 0.1649916, 0.1248156, 0.1364688, 0.1570428, 0.16551, 0.1535652,
		0.153792, 0.1444284, 0.1402596, 0.1580148, 0.1400328, 0.1317168, 0.1256688, 0.138996, 0.133218, 0.1250856, 0.1080324, 0.1381212,
		0.1300644, 0.1134108, 0.1031616, 0.1231632, 0.1115964, 0.0996192, 0.0915516, 0.1191672, 0.1138104, 0.1026972, 0.0926208, 0.1060992,
		0.1004076, 0.0922968, 0.0871344, 0.0970812, 0.09288, 0.0907848, 0.090342, 0.089046, 0.089694, 0.0903744, 0.0909792, 0.0925236,
		0.092664, 0.0946512, 0.0992844, 0.096714, 0.1025568, 0.109026, 0.1239192, 0.1080972, 0.1201392, 0.1225044, 0.1286064, 0.1474632,
		0.1445472, 0.1453572, 0.1209276, 0.1454976, 0.1221912, 0.1184004, 0.1068444, 0.1182384, 0.1087776, 0.0995328, 0.062964, 0.1067904,
		0.0810216, 0.0158328, 0.0022572, 0.00243, 0.0010368, 0.0003348, 0.0001404, 0.0007452, 0.0001836, 7.56E-05, 8.64E-05, 0.002106,
		0.002052, 0.0019656, 0.0031428, 0.0056808, 0.0111564, 0.023706, 0.058806, 0.0173556, 0.0504144, 0.0758808, 0.11475, 0.0453276,
		0.089802, 0.1099764, 0.1335744, 0.09099, 0.1438128, 0.1691496, 0.173124, 0.1792152, 0.20061, 0.2262492, 0.24354, 0.164808,
		0.1630692, 0.1615572, 0.1581336, 0.2051352, 0.1921536, 0.175122, 0.1358532, 0.1642896, 0.1350972, 0.1303236, 0.1138428, 0.1456596,
		0.135432, 0.114966, 0.100278, 0.1303884, 0.1167696, 0.1017576, 0.0870048, 0.0873072, 0.085698, 0.056214, 0.0130572, 0.0275724,
		0.0482652, 0.020682, 0.0133164, 0.0782568, 0.0822312, 0.07155, 0.0712044, 0.0605772, 0.0687096, 0.0687204, 0.0787428, 0.0830088,
		0.0852012, 0.0864432, 0.0920484, 0.085698, 0.0869616, 0.087156, 0.09504, 0.0814104, 0.0918972, 0.0919188, 0.0891216, 0.0947052,
		0.09504, 0.0848448, 0.051408, 0.0820368, 0.0129708, 0.0100656, 0.0061344, 0.047466, 0.0721224, 0.0904716, 0.079542, 0.0154332,
		0.0368064, 0.045576, 0.054, 0.0182736, 0.0179712, 0.0139428, 0.008046, 0.0323352, 0.0155628, 0.0118152, 0.0072684, 0.0070416,
		0.0055512, 0.0030996, 0.0020736, 2(1.08E-05), 0.00054, 0.0010584, -2.16E-05, 0.0031752, 0.0106704, 0.0306504, 0.005022, 0.0426168,
		0.1134, 0.1351188, 0.066258, 0.086562, 0.1340388, 0.1532196, 0.1172016, 0.1268136, 0.139158, 0.1457568, 0.1442556, 0.142614,
		0.143586, 0.1440072, 0.1479168, 0.1447848, 0.138456, 0.0887328, 0.1392012, 0.1258632, 0.1051488, 0.085806, 0.1379484, 0.109566,
		0.1019844, 0.0797904, 0.1045656, 0.094878, 0.0814752, 0.0646488, 0.101844, 0.0893268, 0.077652, 0.0772308, 0.0826092, 0.0796392,
		0.0766368, 0.0702864, 0.0717444, 0.0638064, 0.0589464, 0.0523692, 0.0580716, 0.057888, 0.0622404, 0.06642, 0.0612684, 0.0675216,
		0.0721764, 0.0819612, 0.068688, 0.0839052, 0.1074924, 0.1369872, 0.1094688, 0.1496124, 0.170478, 0.1855872, 0.2101896, 0.214272,
		0.1971864, 0.1863432, 0.216108, 0.1817856, 0.167724, 0.1485756, 0.1620108, 0.1439856, 0.1333152, 0.1198476, 0.124038, 0.1167696,
		0.1086156, 0.1027188, 0.1122768, 0.1064664, 0.0966492, 0.0923832, 0.0929016, 0.1012824, 0.1008072, 0.110052, 0.1221696, 0.1114776,
		0.1168452, 0.1200096, 0.1030752, 0.1081944, 0.1187892, 0.12528, 0.1076868, 0.1193508, 0.131382, 0.1385316, 0.123768, 0.1342872,
		0.171774, 0.2146932, 0.1349136, 0.14418, 0.1804032, 0.21708, 0.1469124, 0.1782, 0.241002, 0.2900448, 0.2545668, 0.246996,
		0.227772, 0.1727892, 0.20736, 0.1773468, 0.1520532, 0.1370304, 0.1412316, 0.1366524, 0.1278396, 0.1242972, 0.152226, 0.1258848,
		0.124416, 0.1183896, 0.1213164, 0.116316, 0.112644, 0.1110888, 0.1139508, 0.110808, 0.1088856, 0.1051812, 0.108, 0.1030968,
		0.1000944, 0.0972324, 0.0993168, 0.099198, 0.0977076, 0.099198, 0.0961416, 0.0972, 0.0981288, 0.1018764, 0.0958392, 0.098334,
		0.1049328, 0.1130868, 0.0959796, 0.102492, 0.1086372, 0.1176444, 0.1149228, 0.1321056, 0.1440072, 0.1679508, 0.1555848, 0.2138616,
		0.279018, 0.2931876, 0.3108024, 0.2996568, 0.2890188, 0.2544264, 0.3050136, 0.2530656, 0.173664, 0.1415772, 0.1963872, 0.1652724,
		0.1403028, 0.1213488, 0.1681668, 0.1559088, 0.1369656, 0.12879, 0.140508, 0.1251288, 0.121176, 0.1211112, 0.1295136, 0.1218888,
		0.1211436, 0.1180008, 0.1196424, 0.1218564, 0.1231092, 0.1248696, 0.117342, 0.122364, 0.1344168, 0.1501092, 0.1199016, 0.1273644,
		0.1460916, 0.1683288, 0.1221696, 0.136998, 0.1654668, 0.2201148, 0.1523772, 0.163242, 0.2310228, 0.3013524, 0.25839, 0.2321568,
		0.1981152, 0.1952748, 0.1926396, 0.1716012, 0.1414908, 0.12636, 0.1589976, 0.1393308, 0.1218132, 0.112266, 0.125658, 0.1208196,
		0.114588, 0.1029996, 0.1164456, 0.1063044, 0.1010556, 0.0973188, 0.1098792, 0.098712, 0.0987876, 0.096336, 0.099198, 0.0961956,
		0.0943164, 0.09234, 0.0963468, 0.0951912, 0.0939492, 0.092772, 0.0941328, 0.0959364, 0.0939384, 0.0946728, 0.0925128, 0.0973296,
		0.101682, 0.1035612, 0.0939384, 0.1007424, 0.11367, 0.1232388, 0.1004292, 0.1191672, 0.1309932, 0.146988, 0.1476684, 0.1657908,
		0.1802736, 0.1835352, 0.217782, 0.1872936, 0.1625832, 0.1442556, 0.1807272, 0.1469016, 0.1255716, 0.1117584, 0.1502604, 0.1312416,
		0.1169748, 0.112212, 0.1354428, 0.115074, 0.1085832, 0.0982044, 0.1040364, 0.0999216, 0.0974052, 0.09747, 0.0998568, 0.0995868,
		0.0992952, 0.0970596, 0.0946944, 0.0974808, 0.1004076, 0.1104948, 0.099522, 0.10476, 0.113724, 0.1265112, 0.107514, 0.1182168,
		0.1465992, 0.1692576, 0.1158624, 0.1330452, 0.1709424, 0.235386, 0.1479384, 0.1552284, 0.2146932, 0.2691036, 0.2403972, 0.2150712,
		0.1948968, 0.189, 0.1846692, 0.1639224, 0.1478196, 0.1389528, 0.1428732, 0.1340388, 0.1221156, 0.1126332, 0.1278072, 0.12717,
		0.1152252, 0.1057644, 0.1206684, 0.1077732, 0.1031184, 0.0972, 0.1190484, 0.1080108, 0.098442, 0.096714, 0.099522, 0.1025028,
		0.1009584, 0.1023084, 0.1050516, 0.1009584, 0.1010016, 0.1018656, 0.1033128, 0.0998136, 0.0999972, 0.1006668, 0.0969408, 0.0994896,
		0.1040364, 0.11583, 0.1007208, 0.1063584, 0.1207008, 0.1420956, 0.1145664, 0.1428408, 0.1495692, 0.1659528, 0.1585764, 0.1677348,
		0.1683828, 0.162756, 0.1843344, 0.1641276, 0.1540188, 0.1390824, 0.1798956, 0.1488024, 0.135756, 0.1183896, 0.1442664, 0.1255608,
		0.111726, 0.101736, 0.1150416, 0.1125468, 0.1019628, 0.0992952, 0.1083564, 0.1022652, 0.1014012, 0.100926, 0.1057536, 0.1067688,
		0.1066284, 0.0821448, 0.0839916, 0.0986688, 0.1053756, 0.112644, 0.1015308, 0.1092528, 0.112752, 0.1208088, 0.1164996, 0.1352592,
		0.1494288, 0.1777248, 0.1274292, 0.1482624, 0.1693656, 0.1868184, 0.1503144, 0.1552608, 0.16875, 0.19575, 0.1671732, 0.1787184,
		0.1742148, 0.1660176, 0.1751868, 0.162594, 0.1450872, 0.1403784, 0.158436, 0.1559952, 0.1545588, 0.1380456, 0.1558656, 0.1495368,
		0.1354212, 0.126144, 0.13986, 0.135702, 0.1142964, 0.1052892, 0.1086912, 0.0990576, 0.0948348, 0.090936, 0.0996948, 0.0937548,
		0.0918648, 0.0906876, 0.090234, 0.0888408, 0.0879552, 0.0875988, 0.0889056, 0.088938, 0.0891324, 0.0894672, 0.0898128, 0.0916812,
		0.0917676, 0.1003428, 0.096498, 0.1212732, 0.137592, 0.1551204, 0.1330884, 0.1578096, 0.1804356, 0.194238, 0.1716336, 0.176418,
		0.178632, 0.1515024, 0.17847, 0.1448172, 0.118152, 0.1036908, 0.1553364, 0.1227744, 0.1044684, 0.08478, 0.1356804, 0.1012824,
		0.091314, 0.0770148, 0.1039608, 0.088236, 0.0862488, 0.0846072, 0.0949428, 0.0879228, 0.08154, 0.0731592, 0.0853092, 0.0915732,
		0.0908172, 0.0816912, 0.0713664, 0.092772, 0.0985068, 0.1113912, 0.0898992, 0.0984528, 0.1055052, 0.118368, 0.091638, 0.112266,
		0.1420632, 0.175986, 0.1311228, 0.1598724, 0.1924128, 0.2146284, 0.175554, 0.1929204, 0.2121228, 0.2276748, 0.2036988, 0.2043468,
		0.2052216, 0.1920672, 0.1988172, 0.1789668, 0.156114, 0.1493856, 0.1576368, 0.1538136, 0.144288, 0.1259064, 0.143856, 0.1364148,
		0.1187136, 0.1115748, 0.118206, 0.1091016, 0.1087776, 0.1002564, 0.1209816, 0.1074816, 0.0951264, 0.0921024, 0.1004616, 0.0966816,
		0.094392, 0.0941436, 0.095202, 0.0957204, 0.0963468, 0.0954288, 0.0942948, 0.0921348, 0.0929988, 0.0906228, 0.0917028, 0.0910008,
		0.0898884, 0.0911952, 0.089532, 0.092772, 0.0926424, 0.095472, 0.0948996, 0.0960876, 0.098496, 0.1004616, 0.1044468, 0.1026648,
		2(0.1054296), 0.1122768, 0.1115424, 0.1094796, 0.1011096, 0.1236708, 0.1123308, 0.1000512, 0.0823284, 0.1158516, 0.1001376, 0.0823068,
		0.0836784, 0.0931284, 0.0804924, 0.0573588, 0.0527148, 0.0621324, 0.0572508, 0.0494208, 0.045306, 0.0402624, 0.037422, 0.0341496,
		0.0380808, 0.0306072, 0.0364284, 0.0407808, 0.0587304, 0.0588924, 0.0848988, 0.1020708, 0.0965412, 0.0752544, 0.0930096, 0.1109592,
		0.128898, 0.0982368, 0.114912, 0.1438668, 0.1677996, 0.1429812, 0.1402272, 0.1559304, 0.1629396, 0.1479276, 0.1554228, 0.1460376,
		0.1311768, 0.1612008, 0.1406592, 0.1174068, 0.1103976, 0.1386504, 0.125172, 0.126306, 0.1071576, 0.1377108, 0.1225908, 0.1096956,
		0.1006128, 0.1135728, 0.1033452, 0.1006344, 0.094068, 0.1177092, 0.1142856, 0.0965304, 0.0889488, 0.1131084, 0.1061532, 0.0946944,
		0.0944028, 0.1068444, 0.097092, 0.094068, 0.0957528, 0.1000728, 0.0961092, 0.0962388, 0.0904284, 0.08667, 0.0928476, 0.1034208,
		0.1039284, 0.0943056, 0.0897696, 0.1039824, 0.1038744, 0.0946512, 0.0964872, 0.0998136, 0.0979668, 0.108486, 0.093258, 0.0947592,
		0.0932688, 0.1124064, 0.0958392, 0.0936576, 0.0830196, 0.1132596, 0.096552, 0.0786672, 0.0875448, 0.1037772, 0.090342, 0.0670788,
		0.0670032, 0.0719388, 0.068418, 0.0680076, 0.0682776, 0.060102, 0.0511704, 0.0289764, 0.0211896, 0.0478872, 0.0465048, 0.044658,
		0.052218, 0.0666036, 0.0691848, 0.0793584, 0.0885384, 0.0872748, 0.0895428, 0.1049004, 0.1134324, 0.0901044, 0.103464, 0.1142532,
		0.1247616, 0.1050516, 0.1236276, 0.1505196, 0.1755432, 0.1378944, 0.1412424, 0.1545696, 0.1874556, 0.1624752, 0.157032, 0.1658772,
		0.1534248, 0.1587276, 0.1593648, 0.152874, 0.14472, 0.1428516, 0.143856, 0.1181088, 0.11205, 0.1350324, 0.1256256, 0.1124388,
		0.1051812, 0.1123092, 0.103626, 0.10098, 0.0935928, 0.1153116, 0.1029024, 0.1017792, 0.1015956, 0.100656, 0.0987768, 0.1027512,
		0.1026648, 0.1029024, 0.102762, 0.1008288, 0.102492, 0.1025784, 0.1025244, 0.1031292, 0.1091016, 0.109512, 0.10638, 0.1095876,
		0.1158948, 0.1068768, 0.1123848, 0.1123524, 0.1326024, 0.1200744, 0.1541484, 0.1843776, 0.2134404, 0.2228688, 0.251694, 0.266436,
		0.2562408, 0.2592, 0.2351484, 0.1857384, 0.146556, 0.2076948, 0.159624, 0.1434996, 0.1146852, 0.1568916, 0.147204, 0.1315656,
		0.1199124, 0.14499, 0.1240164, 0.1148688, 0.1090152, 0.1148364, 0.1059372, 0.1018224, 0.0972, 0.1055052, 0.1024812, 0.0998028,
		0.0961632, 0.0921672, 0.0989712, 0.1121472, 0.1188864, 0.1031616, 0.109296, 0.1219212, 0.1388124, 0.1242648, 0.1552068, 0.2089476,
		0.2519532, 0.156168, 0.1972944, 0.2636388, 0.3315816, 0.238626, 0.3011904, 0.4206708, 0.4431888, 0.4450248, 0.4063176, 0.3306636,
		0.2485512, 0.359046, 0.3067848, 0.2208384, 0.1744956, 0.2306232, 0.1998756, 0.1768716, 0.1600344, 0.1737612, 0.1503792, 0.1287036,
		0.1215972, 0.1379268, 0.1338768, 0.1222668, 0.1155276, 0.1241244, 0.1258524, 0.1171692, 0.111834, 0.1161756, 0.1142532, 0.1127844,
		0.1110024, 0.113238, 0.1099764, 0.1088856, 0.1073952, 0.1107648, 0.110484, 0.1097388, 0.1117044, 0.1090152, 0.1113696, 0.1119096,
		0.118746, 0.1129356, 0.1209384, 0.1232712, 0.1403676, 0.1263492, 0.15687, 0.2153088, 0.2551392, 0.2749788, 0.284364, 0.2625264,
		0.2026296, 0.2487888, 0.2413476, 0.1803492, 0.1519884, 0.2302776, 0.1645596, 0.1429272, 0.1314684, 0.1834272, 0.1397952, 0.1232496,
		0.115182, 0.1510596, 0.1358424, 0.130086, 0.1199772, 0.1267812, 0.1253232, 0.120528, 0.112428, 0.119124, 0.117342, 0.1197504,
		0.1185408, 0.1069848, 0.1231848, 0.1352808, 0.15363, 0.1226556, 0.131382, 0.1485648, 0.1860408, 0.1202148, 0.1371492, 0.209142,
		0.3695652, 0.137322, 0.218916, 0.3211272, 0.418716, 0.3239244, 0.3852252, 0.5113584, 0.5596128, 0.5441256, 0.5013684, 0.4402188,
		0.3578796, 0.38421, 0.296622, 0.2267784, 0.171288, 0.267948, 0.2181492, 0.1980936, 0.169344, 0.182898, 0.1560492, 0.138132,
		0.132678, 0.1464804, 0.1368468, 0.12609, 0.122418, 0.13959, 0.1257876, 0.1299996, 0.1289736, 0.1329264, 0.1272024, 0.123336,
		0.1226016, 0.1228608, 0.1231956, 0.1200636, 0.1179684, 0.1186272, 0.1175472, 0.11691, 0.1170072, 0.1170936, 0.119178, 0.122148,
		0.1272564, 0.12312, 0.129438, 0.1349784, 0.1702944, 0.1234332, 0.1439424, 0.2346192, 0.2706696, 0.3183516, 0.3557412, 0.3398328,
		0.3171852, 0.3654288, 0.3168828, 0.2636928, 0.2101248, 0.262224, 0.20493, 0.1511136, 0.1410804, 0.1845504, 0.1481976, 0.1390392,
		0.118962, 0.1658988, 0.1475496, 0.131868, 0.1246428, 0.14553, 0.1418256, 0.1321164, 0.1246212, 0.1346868, 0.132138, 0.1277424,
		0.124686, 0.1229364, 0.1260684, 0.140346, 0.1529496, 0.1240056, 0.1245456, 0.1476684, 0.1839348, 0.124632, 0.1525176, 0.2266812,
		0.4580388, 0.1373328, 0.189594, 0.2775168, 0.332694, 0.193158, 0.2455164, 0.3429432, 0.4111236, 0.3662172, 0.3051972, 0.261846,
		0.1937628, 0.3016656, 0.2654964, 0.1904796, 0.1661796, 0.237222, 0.2102112, 0.1879848, 0.1397952, 0.142236, 0.1312308, 0.12474,
		0.1220616, 0.121824, 0.1200096, 0.1127952, 0.1122012, 0.1223532, 0.1205388, 0.1116504, 0.098388, 0.1149768, 0.1107216, 0.1093176,
		0.1069632, 0.1042632, 0.1033668, 0.1036476, 0.1026972, 0.1051812, 0.1055808, 0.106272, 0.1039932, 0.1056888, 0.109134, 0.1079892,
		0.1104516, 0.1025028, 0.1142748, 0.1210032, 0.1256904, 0.1195452, 0.129924, 0.164754, 0.2074032, 0.1957932, 0.2006208, 0.1833732,
		0.167616, 0.189918, 0.1686636, 0.1436724, 0.1122768, 0.1593, 0.1437372, 0.1148904, 0.1012176, 0.1308744, 0.1044792, 0.0960228,
		0.0820908, 0.1177848, 0.0948996, 0.0991332, 0.090504, 0.1029348, 0.100386, 0.0939816, 0.0918324, 0.0945756, 0.094986, 0.0993492,
		0.0981828, 0.0852552, 0.091422, 0.1006128, 0.1126656, 0.0848232, 0.1004292, 0.1210572, 0.1247508, 0.119232, 0.1225368, 0.138456,
		0.1789236, 0.1467072, 0.1499472, 0.1743876, 0.241164, 0.1505304, 0.1585008, 0.191808, 0.2214108, 0.185814, 0.1797984, 0.1825524,
		0.158814, 0.1859436, 0.1781028, 0.156978, 0.1416528, 0.1540512, 0.1464588, 0.1274832, 0.112158, 0.1398168, 0.1261224, 0.1252584,
		0.1204956, 0.1231848, 0.1151604, 0.1036152, 0.0980748, 0.1082808, 0.1059048, 0.1039824, 0.1032048, 0.10449, 0.103896, 0.1022112,
		0.1018656, 0.1031292, 0.1001592, 0.1024488, 0.1025892, 0.1003968, 0.1039176, 0.1003752, 0.1028916, 0.0966924, 0.1034316, 0.1042632,
		0.1071792, 0.0995868, 0.105894, 0.1159812, 0.1262088, 0.1194264, 0.1308636, 0.1433376, 0.149688, 0.1426572, 0.1565136, 0.1582848,
		0.1594836, 0.1854792, 0.1727892, 0.1520748, 0.1296432, 0.1739016, 0.14364, 0.1296, 0.1102248, 0.142884, 0.136188, 0.1248804,
		0.1131408, 0.127008, 0.114858, 0.1006884, 0.093744, 0.1060776, 0.0988632, 0.097578, 0.0968652, 0.0995328, 0.1023192, 0.1041876,
		0.0988308, 0.0958284, 0.1039176, 0.1105272, 0.1165968, 0.1077192, 0.1143072, 0.1233684, 0.1393416, 0.1195776, 0.1316304, 0.1629396,
		0.1993896, 0.1301292, 0.1513728, 0.1648728, 0.189918, 0.15201, 0.1709964, 0.1865484, 0.2208276, 0.1873476, 0.181332, 0.1651752,
		0.1586196, 0.1630152, 0.1579284, 0.1505628, 0.150876, 0.157788, 0.1479708, 0.1377864, 0.128844, 0.1442664, 0.134622, 0.1270728,
		0.1209276, 0.126576, 0.1166292, 0.107838, 0.0974268, 0.1197936, 0.1267056, 0.1230552, 0.114696, 0.1197396, 0.1159812, 0.10638,
		0.1042956, 0.1144476, 0.108486, 0.1038204, 0.1018332, 0.1032156, 0.1034316, 0.1045872, 0.101574, 0.0979236, 0.0991008, 0.10341,
		0.106164, 0.0963576, 0.1033992, 0.1113696, 0.1227204, 0.1107324, 0.1301076, 0.1457028, 0.146232, 0.146934, 0.1543752, 0.1529064,
		0.1494396, 0.1603476, 0.1499256, 0.1397736, 0.1135188, 0.1416744, 0.13149, 0.1002996, 0.0829764, 0.1317384, 0.1002348, 0.0944352,
		0.0867024, 0.1007964, 0.099522, 0.0963684, 0.087858, 0.0912924, 0.0930636, 0.0855144, 0.0820908, 0.0891864, 0.089694, 0.0805248,
		0.084456, 0.084888, 0.0894024, 0.0907524, 0.0980424, 0.0865836, 0.0971136, 0.1035288, 0.1130112, 0.0948888, 0.1066716, 0.15066,
		0.1887084, 0.1292436, 0.15363, 0.1621836, 0.1887732, 0.1557468, 0.1631448, 0.1761696, 0.180306, 0.1750572, 0.1669248, 0.1648836,
		0.1613952, 0.1563624, 0.1590408, 0.1544724, 0.1268136, 0.1469448, 0.129654, 0.112158, 0.10476, 0.128142, 0.121608, 0.111618,
		0.1018008, 0.1167696, 0.104058, 0.0964548, 0.0927612, 0.1122336, 0.09936, 0.0952236, 0.0955692, 0.1053216, 0.0981828, 0.0976536,
		0.09477, 0.10044, 0.098712, 0.096498, 0.092718, 0.0995112, 0.0979668, 0.0964656, 0.096228, 0.0973728, 0.0990468, 0.1008396,
		0.0981504, 0.0973728, 0.0970596, 0.1023192, 0.1022652, 0.1005156, 0.103734, 0.1104732, 0.1193832, 0.1153332, 0.122904, 0.1212408,
		0.1101276, 0.1281744, 0.1193076, 0.0964548, 0.0830736, 0.1130868, 0.0955044, 0.085698, 0.0709344, 0.0953208, 0.0838404, 0.0793692,
		0.070794, 0.0879012, 0.078786, 0.0689904, 0.0470988, 0.0618732, 0.0436752, 0.03024, 0.0171288, 0.0260064, 0.0242136, 0.02322,
		0.0180576, 0.013176, 0.0258012, 0.052164, 0.075978, 0.04698, 0.0822528, 0.0884088, 0.10287, 0.0692712, 0.0947592, 0.1188432,
		0.1690848, 0.1106352, 0.1391256, 0.1702512, 0.1893132, 0.1561572, 0.1691172, 0.1751544, 0.1816452, 0.1766556, 0.1753164, 0.1664604,
		0.1617084, 0.1629612, 0.1655532, 0.1539108, 0.1479276, 0.1517616, 0.1444068, 0.1187136, 0.1036476, 0.1474416, 0.1357236, 0.1129356,
		0.0896832, 0.1224396, 0.1064232, 0.0963144, 0.077706, 0.1051056, 0.0973836, 0.092232, 0.0822096, 0.0938952, 0.089424, 0.084618,
		0.0883116, 0.0897264, 0.088506, 0.0878364, 0.0832896, 0.0888948, 0.0875988, 0.0853308, 0.0874044, 0.083916, 0.0930636, 0.0949752,
		0.1020924, 0.0928692, 0.1105164, 0.1244592, 0.1559196, 0.14283, 0.1782648, 0.1998648, 0.2317248, 0.243486, 0.2511972, 0.2426544,
		0.2137752, 0.192834, 0.1565892, 0.137538, 0.1088532, 0.1489644, 0.1325592, 0.1116288, 0.0900828, 0.1142748, 0.0934848, 0.0938412,
		0.0869292, 0.0950616, 0.088182, 0.0868968, 0.0872208, 0.087318, 0.0876852, 0.0878472, 0.0856548, 0.093744, 0.09342, 0.093042,
		0.0917784, 0.0875556, 0.0921348, 0.0966384, 0.1108512, 0.0899424, 0.1027188, 0.133326, 0.1460052, 0.1037556, 0.148608, 0.1914192,
		0.2236032, 0.1732104, 0.2121984, 0.2318436, 0.2470392, 0.2428596, 0.255366, 0.2843964, 0.291546, 0.2639412, 0.2565648, 0.2477844,
		0.2312604, 0.2412612, 0.236142, 0.20331, 0.1836324, 0.1962684, 0.181656, 0.1629288, 0.1542888, 0.1585872, 0.1476144, 0.128952,
		0.1160784, 0.13473, 0.1191672, 0.111456, 0.1006776, 0.12285, 0.1151928, 0.1075464, 0.0976536, 0.0920592, 0.0930204, 0.0871776,
		0.0817668, 0.0921024, 0.0883872, 0.0891216, 0.0862488, 0.088992, 0.0877932, 0.086562, 0.0849852, 0.0862704, 0.087318, 0.0920484,
		0.104706, 0.0936144, 0.1134972, 0.1254204, 0.1512972, 0.1332288, 0.1810296, 0.2117556, 0.2418768, 0.2737692, 0.3164724, 0.2650644,
		0.2244024, 0.2700108, 0.2578068, 0.2392308, 0.218214, 0.1753596, 0.1672596, 0.1548612, 0.1476252, 0.1565028, 0.1372896, 0.131274,
		0.1243404, 0.1258848, 0.1254744, 0.1241892, 0.115236, 0.1224396, 0.1127196, 0.1116612, 0.1066392, 0.1105056, 0.109296, 0.0983664,
		0.0974592, 0.0955368, 0.1091124, 0.1121364, 0.122256, 0.1092636, 0.1279908, 0.15417, 0.1587384, 0.143748, 0.1526364, 0.18036,
		0.2025432, 0.1670004, 0.1790208, 0.1997676, 0.2332368, 0.2040768, 0.232848, 0.1959876, 0.2063664, 0.2042388, 0.1917864, 0.1846908,
		0.1764828, 0.165078, 0.1633932, 0.160542, 0.1434456, 0.1600992, 0.157518, 0.1301076, 0.1141776, 0.1475604, 0.1363716, 0.1183896,
		0.1035612, 0.1246212, 0.1036152, 0.094014, 0.089532, 0.1159164, 0.1098144, 0.0987552, 0.097956, 0.1109376, 0.1076004, 0.1040148,
		0.0989712, 0.1090368, 0.1078056, 0.1057428, 0.1032372, 0.1041336, 0.1064124, 0.1069956, 0.103248, 0.0995436, 0.102708, 0.107892,
		0.1085508, 0.0979236, 0.1086264, 0.1120608, 0.1372248, 0.111942, 0.1535436, 0.1920132, 0.1988064, 0.1673568, 0.186408, 0.1796364,
		0.1669788, 0.1765044, 0.1688796, 0.1567512, 0.1216728, 0.15984, 0.1515024, 0.1248912, 0.1141884, 0.1409832, 0.1199664, 0.1095552,
		0.1012932, 0.1122876, 0.1090692, 0.1042308, 0.0940356, 0.1096848, 0.0961956, 0.0987444, 0.1032372, 0.1068336, 0.1040256, 0.0963576,
		0.096336, 0.0907632, 0.1107972, 0.1228716, 0.1304316, 0.1050948, 0.1207656, 0.1410156, 0.1538244, 0.1044144, 0.141912, 0.1624212,
		0.2318976, 0.1475712, 0.1739988, 0.2355048, 0.2919672, 0.2255148, 0.2733372, 0.3362364, 0.3452544, 0.3300048, 0.3045384, 0.2625372,
		0.230418, 0.27243, 0.205632, 0.1600668, 0.1450548, 0.2029212, 0.1599588, 0.1350648, 0.1183896, 0.164484, 0.1480788, 0.1318248,
		0.1241244, 0.1322136, 0.1300428, 0.1255176, 0.1168668, 0.1296864, 0.1223424, 0.114426, 0.1111212, 0.127008, 0.1244808, 0.1134216,
		0.1087668, 0.118476, 0.1118556, 0.10638, 0.1028052, 0.1118988, 0.1046304, 0.0992736, 0.0979668, 0.1012608, 0.1002996, 0.1000512,
		0.1075464, 0.1095552, 0.1122444, 0.131328, 0.1632744, 0.1272132, 0.1370628, 0.1463508, 0.1580148, 0.13905, 0.1622916, 0.1468584,
		0.1457676, 0.161028, 0.1569456, 0.1365552, 0.124524, 0.1577988, 0.1458216, 0.131706, 0.1108512, 0.133974, 0.10044, 0.0868752,
		0.079434, 0.1132056, 0.0836244, 0.081054, 0.0794124, 0.0809244, 0.0789588, 0.078138, 0.0760536, 0.0791532, 0.0768204, 0.0763128,
		0.0755676, 0.0707724, 0.0758808, 0.112266, 0.122094, 0.0777708, 0.1208952, 0.1274184, 0.138456, 0.1184976, 0.1308744, 0.1402272,
		0.186948, 0.126306, 0.1326024, 0.1398384, 0.1735452, 0.1352592, 0.1564704, 0.1555524, 0.1558332, 0.1491804, 0.141588, 0.1394172,
		0.1401516, 0.1747332, 0.1428192, 0.1280988, 0.1160676, 0.1583496, 0.1456272, 0.1235196, 0.1156356, 0.1280124, 0.113508, 0.0945108,
		0.08559, 0.0991764, 0.0916704, 0.0884304, 0.07776, 0.0850176, 0.073278, 0.0686772, 0.0552528, 0.069984, 0.0650052, 0.0526284,
		0.03969, 0.0590652, 0.0570996, 0.0396792, 0.0334368, 0.0671328, 0.0655236, 2(0.03888), 0.0383076, 0.061722, 0.0696816, 0.0711288,
		0.0427356, 0.0758808, 0.0890568, 0.1039608, 0.0886788, 0.1059588, 0.1221372, 0.135864, 0.132894, 0.1455732, 0.1496772, 0.1512108,
		0.1607364, 0.158436, 0.1505412, 0.1473984, 0.1619676, 0.1503684, 0.1466424, 0.1080108, 0.1450008, 0.12609, 0.0939384, 0.0761832,
		0.110592, 0.1024056, 0.1023516, 0.0947484, 0.0979344, 0.0884412, 0.0878364, 0.0830088, 0.082242, 0.079434, 0.0619596, 0.0600264,
		0.0680076, 0.070956, 0.0753408, 0.091746, 0.0772956, 0.0846072, 0.096336, 0.105678, 0.0548964, 0.0929664, 0.1190052, 0.1495476,
		0.086346, 0.1156356, 0.145638, 0.1503144, 0.1183464, 0.1427544, 0.1471824, 0.1583712, 0.1515564, 0.1568592, 0.1472904, 0.1292976,
		0.1525824, 0.1356048, 0.1154736, 0.1060344, 0.1357668, 0.116694, 0.1046736, 0.0777924, 0.1195344, 0.1135296, 0.098928, 0.0887544,
		0.0989604, 0.08343, 0.0868752, 0.0726516, 0.0860652, 0.0848556, 0.0794664, 0.075114, 0.0801036, 0.078084, 0.0764748, 0.0767124,
		0.0779868, 0.0764424, 0.0755676, 0.073332, 0.078678, 0.0782136, 0.0776196, 0.077166, 0.079812, 0.0799848, 0.0796932, 0.0808812,
		0.0794664, 0.0828468, 0.0884088, 0.1014012, 0.0774684, 0.0969084, 0.1066176, 0.1269648, 0.123714, 0.1202472, 0.1132704, 0.1021464,
		0.128196, 0.1154304, 0.1026216, 0.0835812, 0.1143828, 0.092394, 0.0750816, 0.0274428, 0.09396, 0.077112, 0.0706536, 0.0391716,
		0.0666792, 0.0515052, 0.0472716, 0.0141804, 0.028836, 0.0165672, 0.0146556, 0.0132516, 0.0241272, 0.0238896, 0.022248, 0.0251964,
		0.0166212, 0.0327672, 0.0397116, 0.0569916, 0.0545292, 0.0750492, 0.0912816, 0.1024596, 0.0527904, 0.0930528, 0.1263924, 0.1550988,
		0.1022976, 0.1205712, 0.150714, 0.1822068, 0.1580148, 0.182412, 0.1789344, 0.19764, 0.1714176, 0.1644516, 0.1679184, 0.1622592,
		0.160758, 0.1492776, 0.13716, 0.1056132, 0.152658, 0.145854, 0.1118448, 0.074304, 0.129168, 0.1105812, 0.0926208, 0.0800064,
		0.1073844, 0.0956664, 0.089424, 0.079002, 0.0958284, 0.0882036, 0.0888084, 0.0815508, 0.0820692, 0.0782892, 0.076572, 0.0633636,
		0.0796392, 0.0729108, 0.0629424, 0.0562788, 0.0678672, 0.0698868, 0.0671328, 0.0618192, 0.0609444, 0.0583956, 0.0615708, 0.0665388,
		0.0595944, 0.0589788, 0.0672192, 0.07884, 0.0541836, 0.064584, 0.0719496, 0.0844128, 0.0654156, 0.0726408, 0.0721656, 0.0721008,
		0.084834, 0.0759024, 0.0721872, 0.0487512, 0.09234, 0.0622728, 0.0469584, 0.0314496, 0.073386, 0.058698, 0.04212, 0.0287172,
		0.0616572, 0.0267732, 0.005886, 0.0022896, 0.0193968, 0.0154548, 0.0095472, 0.0056916, 0.0107676, 0.0088344, 0.0088236, 0.0088344,
		0.0080676, 0.0096336, 0.0206388, 0.0236628, 0.035424, 0.0756, 0.0868212, 0.1026648, 0.065124, 0.0868212, 0.115182, 0.143316,
		0.0918324, 0.1139184, 0.1390932, 0.1541592, 0.1133028, 0.1299456, 0.1458972, 0.1525284, 0.1179144, 0.1322784, 0.1455192, 0.1457892,
		0.1430892, 0.1389204, 0.1195128, 0.1024488, 0.1435212, 0.1320516, 0.1054836, 0.0654048, 0.1194156, 0.1002024, 0.0783216, 0.0630936,
		0.0958608, 0.0840564, 0.0764532, 0.0325836, 0.1005156, 0.0403056, 0.012096, 0.0036936, 0.082026, 0.0815508, 0.0662688, 0.0343548,
		0.0495936, 0.0403812, 0.0320112, 0.0315144, 0.03429, 0.0338364, 0.0366876, 0.040392, 0.0376704, 0.0433944, 0.0447336, 0.0444852,
		0.0390852, 0.0370548, 0.0649512, 0.0873936, 0.05697, 0.0837432, 0.1044576, 0.1354752, 0.093366, 0.1119852, 0.1259388, 0.1415016,
		0.1248804, 0.1261656, 0.1267704, 0.119124, 0.1335096, 0.131112, 0.1196424, 0.1062504, 0.1332288, 0.1187028, 0.1127196, 0.1079784,
		0.1179684, 0.1134216, 0.1097604, 0.1008612, 0.1154088, 0.1140588, 0.1090476, 0.1041228, 0.1072872, 0.1033452, 0.1027188, 0.10719,
		0.106434, 0.1109592, 0.1192212, 0.1235088, 0.1156896, 0.1262844, 0.1295244, 0.1421496, 0.1133028, 0.131598, 0.1429704, 0.1554768,
		0.1435968, 0.1543212, 0.2095524, 0.2274048, 0.1575612, 0.1944324, 0.2154708, 0.2336256, 0.1809432, 0.188568, 0.1603368, 0.1620648,
		0.164862, 0.1669896, 0.1984176, 0.1623456, 0.2047032, 0.1552716, 0.1401408, 0.1361772, 0.1496556, 0.1393524, 0.1093176, 0.098658,
		0.1272024, 0.1125576, 0.101952, 0.0902556, 0.1107432, 0.1054296, 0.096768, 0.0812916, 0.1090476, 0.09558, 0.0892404, 0.0799416,
		0.0881064, 0.0832572, 0.0826524, 0.0805248, 0.0836352, 0.0801468, 0.079542, 0.079434, 0.0764316, 0.0774144, 0.080406, 0.0813996,
		0.0731916, 0.0787212, 0.083214, 0.087372, 0.0650808, 0.0928584, 0.1010988, 0.136026, 0.09801, 0.1247616, 0.1361232, 0.1343412,
		0.1405944, 0.142398, 0.1122768, 0.0871776, 0.1181088, 0.0966492, 0.09072, 0.0861732, 0.1063584, 0.0952668, 0.0891324, 0.0795204,
		0.1033128, 0.0921672, 0.0869832, 0.0813888, 0.0880956, 0.084672, 0.0844128, 0.0858276, 0.0834408, 0.0839808, 0.0824472, 0.0856764,
		0.0872424, 0.0905472, 0.0984096, 0.1024704, 0.0860868, 0.103248, 0.1166508, 0.1340712, 0.117774, 0.1339524, 0.15201, 0.1746576,
		0.13203, 0.1472472, 0.1594944, 0.1977588, 0.1575612, 0.1641168, 0.1730916, 0.199908, 0.179712, 0.1862784, 0.180738, 0.1817748,
		0.1717848, 0.1708884, 0.1719468, 0.1631664, 0.171558, 0.1611576, 0.1292544, 0.109782, 0.1491372, 0.136188, 0.1078272, 0.095742,
		0.1310472, 0.1063692, 0.09963, 0.096012, 0.1233036, 0.1065744, 0.0981396, 0.0886248, 0.0927288, 0.0898776, 0.0873612, 0.07938,
		0.0942192, 0.0891216, 0.0787428, 0.0772632, 0.0866808, 0.0830304, 0.0793692, 0.0819072, 0.0820368, 0.0817992, 0.081864, 0.0850392,
		0.0642816, 0.0863676, 0.0946512, 0.0993924, 0.0856764, 0.0976968, 0.1161756, 0.1299132, 0.11043, 0.1203552, 0.1304208, 0.1445904,
		0.1260576, 0.1198584, 0.1192428, 0.1122768, 0.1296972, 0.1172556, 0.104922, 0.0809784, 0.1163268, 0.09855, 0.0801468, 0.0667872,
		0.0813024, 0.0686232, 0.0659664, 0.063018, 0.069174, 0.0666144, 0.0673596, 0.0675432, 0.0635148, 0.0727164, 0.0778032, 0.0836676,
		0.0766368, 0.081594, 0.0816912, 0.0948888, 0.0648324, 0.0864, 0.108216, 0.1254852, 0.103842, 0.1154088, 0.1471284, 0.1612548,
		0.1427976, 0.1573128, 0.1746468, 0.2043252, 0.15741, 0.1669356, 0.1708668, 0.1646028, 0.1449144, 0.145908, 0.1523124, 0.1522152,
		0.1528956, 0.1473444, 0.1475172, 0.1265976, 0.1477008, 0.1444824, 0.1259172, 0.1153656, 0.1256796, 0.1207656, 0.1160028, 0.0965412,
		0.125658, 0.1198692, 0.102438, 0.0910548, 0.1099872, 0.0993924, 0.09504, 0.092394, 0.102492, 0.0950292, 0.097794, 0.0824148,
		0.0950724, 0.0929232, 0.0888948, 0.0849636, 0.0902232, 0.0896724, 0.0853848, 0.0835596, 0.078354, 0.0853632, 0.0903096, 0.0872208,
		0.0805896, 0.0905472, 0.0940032, 0.095202, 0.0730296, 0.1057536, 0.110808, 0.1215648, 0.1098576, 0.1166616, 0.1313928, 0.1350648,
		0.124578, 0.1272132, 0.123174, 0.112374, 0.130518, 0.1190808, 0.104004, 0.0731052, 0.114804, 0.108054, 0.0805896, 0.04941,
		0.0837756, 0.07533, 0.081216, 0.0713556, 0.0676728, 0.0814752, 0.0775764, 0.0781272, 0.0549288, 0.0739368, 0.0730512, 0.0920592,
		0.089748, 0.0942408, 0.0959904, 0.093744, 0.086238, 0.1066716, 0.127008, 0.1550772, 0.1005588, 0.1488456, 0.156438, 0.161298,
		0.1572912, 0.1649052, 0.1628856, 0.1782, 0.1522584, 0.1556604, 0.1550772, 0.1575288, 0.1496772, 0.1504872, 0.157626, 0.161082,
		0.1580688, 0.1575612, 0.1523772, 0.1404864, 0.1570968, 0.14688, 0.1480464, 0.111618, 0.1361232, 0.13338, 0.1230336, 0.1055268,
		0.1239516, 0.124578, 0.116856, 0.105192, 0.1208088, 0.1066716, 0.0972108, 0.0902556, 0.1212624, 0.1150092, 0.1151712, 0.1044036,
		0.109296, 0.1090044, 0.0965952, 0.0955044, 0.1070712, 0.0963468, 0.0951804, 0.0936576, 0.0949752, 0.0953532, 0.096012, 0.0999108,
		0.091854, 0.0944892, 0.1065312, 0.1130544, 0.1061316, 0.111834, 0.1204308, 0.1264896, 0.1076544, 0.1265112, 0.1342116, 0.1442448,
		0.1307988, 0.1340928, 0.1352268, 0.1219428, 0.1566756, 0.1342872, 0.1131624, 0.0952776, 0.1242864, 0.0986472, 0.0824904, 0.0767664,
		0.0926316, 0.0878904, 0.0870804, 0.084456, 0.0875016, 0.0858924, 0.0852228, 0.0866808, 0.0836784, 0.0844884, 0.08937, 0.094986,
		0.087318, 0.0926208, 0.0991656, 0.1119312, 0.092286, 0.1161864, 0.1347624, 0.1575936, 0.1109268, 0.1307232, 0.1540512, 0.1647648,
		0.1567944, 0.1728108, 0.2055456, 0.2289816, 0.205146, 0.2270916, 0.2404512, 0.227664, 0.226314, 0.2241648, 0.2201364, 0.2253204,
		0.22869, 0.2140236, 0.1944432, 0.1799388, 0.2074356, 0.1708884, 0.1572588, 0.1361664, 0.155304, 0.1444392, 0.1323, 0.1255716,
		0.1448388, 0.1404864, 0.12933, 0.1090044, 0.128142, 0.1090152, 0.0866592, 0.078894, 0.1235304, 0.115074, 0.0994896, 0.0826524,
		0.0957204, 0.0888732, 0.088992, 0.0766152, 0.0857952, 0.0742068, 0.0732348, 0.0808812, 0.0815616, 0.0818964, 0.079434, 0.0800604,
		0.0746496, 0.076842, 0.083592, 0.0879012, 0.0862488, 0.0843372, 0.0827064, 0.0873612, 0.077544, 0.0891, 0.090126, 0.0947376,
		0.09342, 0.091962, 0.0852768, 0.0521532, 0.0860328, 0.081486, 0.06318, 0.015552, 0.078462, 0.06696, 0.0261144, 0.0183492,
		0.0256176, 0.0195264, 0.017712, 2(0.0162), 0.0162648, 0.0162, 0.0194076, 0.016038, 0.01944, 0.0267624, 0.0285444, 0.02187,
		0.0266436, 0.0395604, 0.0418716, 0.04995, 0.0649836, 0.0793044, 0.091098, 0.0575316, 0.0857736, 0.1096416, 0.1203444, 0.088722,
		0.1202904, 0.1396548, 0.157086, 0.1135404, 0.1208736, 0.1258632, 0.1192428, 0.1134972, 0.1147932, 0.113076, 0.1067796, 0.1115964,
		0.115344, 0.1086264, 0.1092636, 0.1273428, 0.1386828, 0.1378404, 0.113184, 0.1377972, 0.1368792, 0.1271484, 0.110754, 0.124092,
		0.1114128, 0.1024596, 0.094122, 0.1097604, 0.095796, 0.0876636, 0.0862596, 0.0884088, 0.0926208, 0.0945216, 0.089046, 0.0910764,
		0.0892296, 0.0840672, 0.0829872, 0.085698, 0.0850608, 0.0828468, 0.0827064, 0.085428, 0.0844884, 0.083538, 0.0836136, 0.083376,
		0.0839376, 0.0856656, 0.0872964, 0.08586, 0.0861624, 0.0875664, 0.0905364, 0.088722, 0.0930852, 0.0935388, 0.0899532, 0.0894564,
		0.0870264, 0.0874476, 0.0882468, 0.0927504, 0.0923616, 0.0859248, 0.0845748, 0.0967356, 0.0704268, 0.06669, 0.0606204, 0.0713988,
		0.0673272, 0.0632772, 0.0618192, 0.0682452, 0.0698112, 0.0696276, 0.0682452, 0.0660096, 0.066636, 0.072414, 0.0821988, 0.0676296,
		0.083538, 0.0963036, 0.1029348, 0.0945108, 0.1050948, 0.1138104, 0.1201392, 0.1137132, 0.1256688, 0.1323756, 0.1495476, 0.1209492,
		0.1313172, 0.140886, 0.1582308, 0.1238004, 0.137646, 0.14229, 0.143964, 0.14013, 0.1393956, 0.13824, 0.1246968, 0.1426248,
		0.1415664, 0.1227528, 0.1128708, 0.1398708, 0.1344276, 0.126144, 0.1083996, 0.1207008, 0.11448, 0.1134432, 0.1085832, 0.118746,
		0.1136592, 0.1097388, 0.0994572, 0.1113264, 0.100116, 0.0925776, 0.08343, 0.09261, 0.0948348, 0.0913464, 0.083538, 0.0891432,
		0.0865188, 0.0787968, 0.0739476, 0.0876636, 0.0760536, 0.0729324, 0.0669924, 0.073602, 0.0712152, 0.0718848, 0.0821556, 0.0838296,
		0.0841212, 0.087102, 0.0886248, 0.083376, 0.0881064, 0.0992196, 0.1193292, 0.0945432, 0.1206468, 0.12933, 0.1481652, 0.1350324,
		0.1397412, 0.1429164, 0.1358532, 0.1571184, 0.145638, 0.127764, 0.121338, 0.1313496, 0.1222668, 0.1109592, 0.096768, 0.1119744,
		0.1033668, 0.1027512, 0.0988632, 0.1003752, 0.1020276, 0.0995868, 0.098496, 0.1028808, 0.0992844, 0.0973944, 0.0990252, 0.1040796,
		0.1004184, 0.102276, 0.1033452, 0.0906336, 0.0984096, 0.1198908, 0.1334124, 0.1028268, 0.160218, 0.199098, 0.2080728, 0.1398168,
		0.1691712, 0.1938168, 0.2139156, 0.135378, 0.1681344, 0.1595916, 0.1526148, 0.1726488, 0.1946484, 0.1935468, 0.1987308, 0.203688,
		0.1917864, 0.17172, 0.1582308, 0.1916028, 0.15228, 0.121878, 0.0970272, 0.1427436, 0.1282284, 0.1106028, 0.0937332, 0.1410048,
		0.1213488, 0.1037556, 0.0840996, 0.1103436, 0.0972, 0.0902556, 0.0743148, 0.0889596, 0.0842832, 0.0844128, 0.0836244, 0.0805788,
		0.0790992, 0.0785052, 0.0818316, 0.0805356, 0.0783864, 0.0786672, 0.0771228, 0.079002, 0.0781272, 0.0779004, 0.0781164, 0.0749196,
		0.073926, 0.0836568, 0.0913032, 0.0602316, 0.0871128, 0.1139724, 0.135594, 0.1125576, 0.1421172, 0.1539432, 0.1670436, 0.14958,
		0.1515024, 0.1394604, 0.1090476, 0.1359936, 0.1259712, 0.1074384, 0.0846612, 0.1199556, 0.109566, 0.08451, 0.0670032, 0.1001592,
		0.0958392, 0.092664, 0.0826848, 0.0825552, 0.0816696, 0.0843912, 0.0887868, 0.0794232, 0.079434, 0.0806004, 0.0903528, 0.0903636,
		0.0958284, 0.0969516, 0.1024704, 0.0794988, 0.0986796, 0.1091664, 0.128682, 0.1086588, 0.1239732, 0.15066, 0.1933092, 0.1420308,
		0.1605312, 0.2094984, 0.2447928, 0.1531872, 0.1794852, 0.1845504, 0.177066, 0.2231388, 0.215082, 0.2136996, 0.2030076, 0.1766772,
		0.1604556, 0.1786428, 0.1736964, 0.1796904, 0.1492452, 0.1276128, 0.1098576, 0.1309824, 0.1139616, 0.101412, 0.092124, 0.1297512,
		0.102816, 0.0974808, 0.0897696, 0.1089072, 0.095742, 0.0894456, 0.0815184, 0.0980964, 0.097524, 0.0939708, 0.089694, 0.0912384,
		0.0913248, 0.0899532, 0.0888516, 2(0.0899748), 0.08478, 0.0816804, 0.0880308, 0.0846612, 0.083376, 0.0827064, 0.0820044, 0.0873936,
		0.0862164, 0.0911196, 0.0846828, 0.0893052, 0.097038, 0.119232, 0.1078056, 0.1184544, 0.1304208, 0.1384344, 0.1483488, 0.151092,
		0.1471068, 0.1188324, 0.1602936, 0.1349568, 0.1252908, 0.0780732, 0.129546, 0.1237356, 0.1171476, 0.1054188, 0.1198368, 0.1094256,
		0.1070388, 0.0990684, 0.1008288, 0.099144, 0.0998244, 0.098604, 0.0972324, 0.0978912, 0.0965736, 0.097416, 0.0970812, 0.097416,
		0.0997056, 0.1092312, 0.0951264, 0.1077624, 0.1186056, 0.1434132, 0.1044252, 0.1274076, 0.1451088, 0.1876608, 0.1540512, 0.1882008,
		0.195156, 0.2281932, 0.1639224, 0.1714608, 0.1745928, 0.1848528, 0.1558548, 0.1532304, 0.1761696, 0.1894644, 0.1837404, 0.183384,
		0.1598076, 0.1352268, 0.1775844, 0.14418, 0.1228068, 0.112644, 0.140616, 0.1343088, 0.1085292, 0.1188324, 0.1408212, 0.1348056,
		0.1102572, 0.0941868, 0.131706, 0.1064124, 0.0955584, 0.0900612, 0.1119096, 0.107622, 0.1079352, 0.1041228, 0.1077192, 0.1053756,
		0.104652, 0.103032, 0.1076112, 0.10476, 0.106542, 0.1044468, 0.1067256, 0.1061208, 0.1041012, 0.1053756, 0.1070172, 0.1064664,
		0.107298, 0.109296, 0.1000728, 0.1036044, 0.1116504, 0.1392228, 0.1070172, 0.130194, 0.1470204, 0.1631016, 0.1698624, 0.1517616,
		0.1538568, 0.1283256, 0.1530792, 0.1417068, 0.1162944, 0.0992628, 0.1302264, 0.1111752, 0.0978912, 0.0845208, 0.1066608, 0.09882,
		0.0916812, 0.089586, 0.0978912, 0.0950616, 0.0950292, 0.089424, 0.0945324, 0.0872316, 0.0941004, 0.099036, 0.0889164, 0.0971028,
		0.0974052, 0.105516, 0.085698, 0.1038096, 0.1187244, 0.1477008, 0.113508, 0.1380996, 0.1716552, 0.2429568, 0.1604124, 0.1908576,
		0.2171232, 0.2523852, 0.194184, 0.2104056, 0.2085696, 0.2191752, 0.1820988, 0.1725624, 0.1918728, 0.1955988, 0.1840752, 0.1888812,
		0.1796688, 0.156924, 0.164106, 0.1510488, 0.1375596, 0.1274508, 0.132354, 0.1333152, 0.133002, 0.1049976, 0.1361124, 0.1196964,
		0.1102572, 0.1035396, 0.1249128, 0.1084104, 0.101142, 0.0939168, 0.10071, 0.099468, 0.1039932, 0.0992304, 0.1011852, 0.09882,
		0.0989496, 0.0985824, 0.101304, 0.0998136, 0.1009152, 0.1002348, 0.1016388, 0.1015848, 0.1012608, 0.1023732, 0.098982, 0.1018656,
		0.1053864, 0.1056996, 0.0965304, 0.1024272, 0.1111536, 0.1314144, 0.1203876, 0.1381752, 0.1585008, 0.1697004, 0.173394, 0.1717092,
		0.1484244, 0.1526472, 0.1658772, 0.1511568, 0.125226, 0.1006884, 0.139644, 0.129762, 0.1104084, 0.0985824, 0.1151604, 0.1052568,
		0.0991764, 0.0968112, 0.1032156, 0.1020168, 0.1038204, 0.101682, 0.0996948, 0.09936, 0.0992844, 0.1003644, 0.0988524, 0.1015632,
		0.1052028, 0.10773, 0.0900936, 0.1106028, 0.1250748, 0.1655748, 0.1062072, 0.1468692, 0.1672164, 0.2160972, 0.1387908, 0.1395576,
		0.1638036, 0.2633148, 0.207198, 0.2202012, 0.2154276, 0.178308, 0.1668276, 0.152658, 0.154494, 0.1559736, 0.1603476, 0.1515996,
		0.1501416, 0.1428948, 0.1566108, 0.1393416, 0.1333476, 0.1163916, 0.137538, 0.1266948, 0.111942, 0.10098, 0.120744, 0.120636,
		0.1105056, 0.099684, 0.1263492, 0.11016, 0.0981936, 0.0935172, 0.1140048, 0.112536, 0.1111644, 0.1083024, 0.112212, 0.1106136,
		0.1063476, 0.105894, 0.1104408, 0.1072224, 0.1057428, 0.1039932, 0.1061532, 0.1055916, 0.1055484, 0.1054728, 0.1061316, 0.1084644,
		0.1087776, 0.107784, 0.1064556, 0.1114776, 0.1115964, 0.108054, 0.1071252, 0.1048572, 0.1128816, 0.1204848, 0.1118448, 0.1187352,
		0.1251504, 0.1261116, 0.1292868, 0.1255608, 0.1170936, 0.1136376, 0.1325808, 0.1199016, 0.1163808, 0.1092312, 0.1395792, 0.1182816,
		0.1129788, 0.1101492, 0.1240812, 0.1156788, 0.1120176, 0.1111644, 0.11907, 0.1118448, 0.1104192, 0.1107108, 0.1109268, 0.1139616,
		0.1126008, 0.1252044, 0.107514, 0.1099224, 0.1193184, 0.1347624, 0.1084968, 0.1252476, 0.1443312, 0.1561356, 0.1308312, 0.1379268,
		0.1485864, 0.1845396, 0.1403244, 0.1540404, 0.1542888, 0.1567836, 0.1425168, 0.143316, 0.14445, 0.1436616, 0.144072, 0.141318,
		0.1387584, 0.1362744, 0.1469556, 0.1395036, 0.1347084, 0.1225692, 0.13581, 0.1331532, 0.119934, 0.1131732, 0.124956, 0.11853,
		0.1151172, 0.1106568, 0.114912, 0.1100736, 0.1043604, 0.0966276, 0.1090044, 0.1015524, 0.1089396, 0.1063152, 0.11151, 0.1054188,
		0.1026648, 0.1003428, 0.1057212, 0.1046736, 0.1027728, 0.1008504, 0.1020924, 0.100818, 0.1003212, 0.1039284, 0.10098, 0.1024272,
		0.1015308, 0.1048896, 0.1023516, 0.1017576, 0.104112, 0.100764, 0.1001916, 0.0989388, 0.0997164, 0.0991008, 0.1064664, 0.0979344,
		0.1007208, 0.1036152, 0.1094472, 0.1103436, 0.109296, 0.107676, 0.1114452, 0.1110024, 0.107298, 0.1070496, 0.1104192, 0.1083888,
		0.1091988, 0.108864, 0.111186, 0.1110996, 0.109026, 0.1075356, 0.1115316, 0.1109916, 0.1074276, 0.1108296, 0.1111752, 0.1115856,
		0.1128708, 0.113238, 0.1098252, 0.1105272, 0.1181844, 0.1198044, 0.1110888, 0.1173096, 0.1212732, 0.1304964, 0.1221372, 0.1300644,
		0.1383264, 0.1477764, 0.138078, 0.1424736, 0.1446768, 0.1455516, 0.1387368, 0.1410912, 0.1418472, 0.1393092, 0.1422792, 0.1383372,
		0.1384776, 0.1384128, 0.1431756, 0.1351404, 0.1287144, 0.1223964, 0.1291896, 0.1226232, 0.1160244, 0.1127844, 0.1214676, 0.1143612,
		0.1104192, 0.1040256, 0.1086696, 0.1055052, 0.1004832, 0.0940356, 0.1028268, 0.0990576, 0.0998568, 0.0991332, 0.0989496, 0.0997704,
		0.0981396, 0.0992196, 0.1012608, 0.1020492, 0.0999864, 0.099846, 0.1006236, 0.0998568, 0.0998892, 0.0999, 0.0976752, 0.0971352,
		0.0994788, 0.1048572, 0.099414, 0.0987228, 0.1081728, 0.1172232, 0.1100628, 0.1202364, 0.1299348, 0.1483704, 0.1394172, 0.1488996,
		0.1559736, 0.1625076, 0.1828872, 0.1643436, 0.1620216, 0.1445688, 0.1834704, 0.1517076, 0.1360692, 0.1252692, 0.1661148, 0.14607,
		0.141264, 0.124146, 0.139536, 0.1335528, 0.1274292, 0.1242972, 0.1253448, 0.1261656, 0.1228392, 0.1265976, 0.129816, 0.1319868,
		0.129762, 0.1419444, 0.1207224, 0.1423872, 0.1685232, 0.1830492, 0.14013, 0.1615572, 0.1823688, 0.2103408, 0.1579716, 0.1635228,
		0.187812, 0.2084292, 0.1654344, 0.168372, 0.1671192, 2(0.16389), 0.1599696, 0.1540404, 0.1531224, 0.1595376, 0.1471176, 0.144666,
		0.141696, 0.1705644, 0.147906, 0.132246, 0.1252368, 0.1344816, 0.1290384, 0.1159812, 0.1113372, 0.1297728, 0.1224396, 0.1159272,
		0.1092744, 0.1168236, 0.1116936, 0.1039068, 0.095364, 0.10584, 0.0996084, 0.0978048, 0.094662, 0.1057536, 0.0966708, 0.095364,
		0.096066, 0.0946296, 0.0929124, 0.092664, 0.0988308, 0.0960228, 0.0982152, 0.0981828, 0.098226, 0.0961092, 0.0966168, 0.098442,
		0.1005696, 0.0957528, 0.1067364, 0.1155384, 0.1251828, 0.1140696, 0.1316736, 0.1461564, 0.1592028, 0.1439532, 0.1470528, 0.1456056,
		0.1510488, 0.1536948, 0.1505304, 0.1416636, 0.1259928, 0.140724, 0.1333692, 0.1211652, 0.1124496, 0.1243404, 0.1165752, 0.1121256,
		0.1052352, 0.109242, 0.1081296, 0.1032156, 0.10017, 0.098496, 0.0963144, 0.0979452, 0.1066608, 0.0970056, 0.100008, 0.1045872,
		0.1141884, 0.102924, 0.1130544, 0.1231848, 0.139158, 0.1145124, 0.1229472, 0.1404648, 0.1532952, 0.1313712, 0.145206, 0.1549152,
		0.15795, 0.1562652, 0.159678, 0.1568808, 0.1565352, 0.140886, 0.1501416, 0.1512324, 0.148446, 0.1488024, 0.1480464, 0.1430352,
		0.133596, 0.14796, 0.1420092, 0.1319868, 0.1184004, 0.1395792, 0.1350648, 0.1260792, 0.1166616, 0.1382832, 0.1285956, 0.1212408,
		0.1090584, 0.1281744, 0.1141344, 0.10692, 0.0992088, 0.1177092, 0.1109916, 0.10989, 0.1026, 0.1083564, 0.1045008, 0.097524,
		0.1006776, 0.1030428, 0.097902, 0.098874, 0.1033452, 0.097902, 0.0984528, 0.1053432, 0.106488, 0.100116, 0.108162, 0.1080648,
		0.1095336, 0.1055484, 0.1157436, 0.1182384, 0.1372788, 0.1219104, 0.1411236, 0.1611468, 0.1762128, 0.1485324, 0.1753164, 0.1694304,
		0.1470204, 0.175392, 0.1459512, 0.1369656, 0.111348, 0.1424952, 0.1293084, 0.1112616, 0.0993492, 0.115074, 0.1117692, 0.112644,
		0.096228, 0.1072224, 0.0988956, 0.0955368, 0.0873396, 0.0905688, 0.0903852, 0.09099, 0.095472, 0.0908172, 0.0962928, 0.105408,
		0.1124928, 0.1094364, 0.1151604, 0.1236492, 0.1503468, 0.1172772, 0.1306584, 0.1790856, 0.210654, 0.1803924, 0.1976724, 0.2219184,
		0.239814, 0.220806, 0.2173392, 0.2181816, 0.211032, 0.211356, 0.2008368, 0.2037312, 0.2005344, 0.2135592, 0.2072736, 0.2008044,
		0.1865808, 0.2042604, 0.1841184, 0.1718172, 0.1286712, 0.1487052, 0.1343628, 0.1290924, 0.118962, 0.1419984, 0.1313064, 0.1249992,
		0.1186272, 0.1217808, 0.1143288, 0.1056672, 0.1085508, 0.119124, 0.1076544, 0.1050624, 0.1092528, 0.1072224, 0.1081512, 0.106704,
		0.1037556, 0.1075572, 0.1021248, 0.10557, 0.1003104, 0.1040256, 0.1045008, 0.1037556, 0.1018332, 0.0876852, 0.0943812, 0.1062288,
		0.1125684, 0.1010232, 0.1191672, 0.1293624, 0.13959, 0.1305072, 0.1408536, 0.1575288, 0.1641924, 0.1568268, 0.1633608, 0.1467288,
		0.1356264, 0.1479276, 0.134514, 0.1203012, 0.1157112, 0.1209492, 0.10881, 0.1110348, 0.1190268, 0.1304856, 0.1227636, 0.1205604,
		0.0986148, 0.1080108, 0.0908604, 0.0928584, 0.1152576, 0.1099764, 0.1194912, 0.1166184, 0.0999, 0.11718, 0.10773, 0.1111428,
		0.117666, 0.1124064, 0.12771, 0.1396764, 0.1724328, 0.1338876, 0.1666116, 0.2091636, 0.2539944, 0.1806516, 0.2220048, 0.2491992,
		0.2537568, 0.1941192, 0.203634, 0.21897, 0.23949, 0.2084724, 0.2055672, 0.2207412, 0.2188188, 0.2104596, 0.2051244, 0.2040336,
		0.1860084, 0.2367036, 0.217134, 0.1899072, 0.164808, 0.1709424, 0.1576692, 0.1358424, 0.1198908, 0.1462752, 0.135432, 0.1235628,
		0.1200312, 0.1399788, 0.1333476, 0.1232172, 0.1093932, 0.1154196, 0.1152036, 0.1163592, 0.1142208, 0.114156, 0.112266, 0.1135836,
		0.1143072, 0.113994, 0.113886, 0.1127088, 2(0.1108836), 0.1104948, 0.109566, 0.1098252, 0.1050192, 0.1067796, 0.110646, 0.1145664,
		0.1104624, 0.1181412, 0.1276776, 0.1540404, 0.1334232, 0.1450872, 0.1476252, 0.15093, 0.1473984, 0.1452276, 0.1476576, 0.14634,
		0.1726704, 0.1557684, 0.1441152, 0.1354104, 0.1528416, 0.1383912, 0.1372356, 0.1222668, 0.1396656, 0.13257, 0.1219212, 0.1186812,
		0.1258956, 0.1210572, 0.120204, 0.1167804, 0.1164564, 0.1146528, 0.1140804, 0.1190052, 0.1181304, 0.1201392, 0.1263492, 0.1291248,
		0.1191132, 0.1302588, 0.1440936, 0.168156, 0.1248372, 0.1436292, 0.1732644, 0.232848, 0.1747548, 0.189054, 0.2452032, 0.260766,
		0.1927044, 0.1725192, 0.1674216, 0.1585548, 0.168048, 0.1667844, 0.170424, 0.1430568, 0.1620432, 0.160272, 0.1483596, 0.1345896,
		0.1450116, 0.1345788, 0.1283688, 0.1189404, 0.133272, 0.12447, 0.1137564, 0.1048464, 0.1245132, 0.124146, 0.118098, 0.1143504,
		0.1208088, 0.114264, 0.1117908, 0.1004616, 0.1166832, 0.1165212, 0.1243836, 0.11745, 0.1170828, 0.1099116, 0.1053324, 0.0977076,
		0.1078272, 0.107028, 0.1046736, 0.1009368, 0.1046844, 0.1006776, 0.1006236, 0.1000188, 0.1002564, 0.1014228, 0.1043928, 0.1055052,
		0.1010016, 0.108486, 0.1110564, 0.1130976, 0.1082376, 0.116478, 0.1198584, 0.122634, 0.1173744, 0.1185192, 0.11475, 0.1121688,
		0.1127088, 0.1123308, 0.1115208, 0.1097604, 0.1124064, 0.1044684, 0.107946, 0.1059588, 0.1109052, 0.1095984, 0.1093392, 0.1086588,
		0.1077948, 0.1081512, 0.1089396, 0.1069632, 0.1034208, 0.1039284, 0.1085616, 0.108432, 0.109998, 0.1139508, 0.1124496, 0.1131408,
		0.1100088, 0.1130436, 0.1257012, 0.1470852, 0.1239408, 0.1409292, 0.1461672, 0.1534248, 0.1417824, 0.1476036, 0.1714176, 0.1947132,
		0.1688904, 0.1605636, 0.1545696, 0.1467072, 0.162594, 0.1456488, 0.1404864, 0.1501632, 0.1541268, 0.144774, 0.1516104, 0.1410696,
		0.1492992, 0.14013, 0.1319004, 0.1222344, 0.1323324, 0.1233036, 0.1225584, 0.1199556, 0.1316304, 0.1268676, 0.120258, 0.1127844,
		0.1229904, 0.1191996, 0.1125576, 0.109566, 0.1215216, 0.1151064, 0.1127844, 0.1119312, 0.112752, 0.1079136, 0.1091988, 0.106326,
		0.1083456, 0.1080972, 2(0.1086048), 0.11043, 0.1090368, 0.1073088, 0.1086264, 0.1079136, 0.1072656, 0.1089288, 0.1102788, 0.11124,
		0.1095876, 0.1119204, 0.1145772, 0.1065096, 0.1126224, 0.1126008, 0.1124928, 0.1119312, 0.1125252, 0.105894, 0.108972, 0.1127304,
		0.1127844, 0.1136052, 0.109242, 0.1164456, 0.1161108, 0.1153548, 0.1135944, 0.114318, 0.113778, 0.1128276, 0.1138212, 0.1167696,
		0.1182924, 0.1185948, 0.113994, 0.1188324, 0.1136484, 0.1126764, 0.1127304, 0.1156356, 0.1223748, 0.1165968, 0.1185732, 0.1158192,
		0.125388, 0.129114, 0.129222, 0.1231416, 0.1308528, 0.1369008, 0.1451304, 0.1337148, 0.1407672, 0.1444932, 0.16038, 0.141642,
		0.145152, 0.149472, 0.1469988, 0.1398492, 0.1391796, 0.1383912, 0.1342656, 0.1335744, 0.130356, 0.1290924, 0.1275372, 0.1339956,
		0.131004, 0.1225692, 0.1147824, 0.1258092, 0.1183464, 0.1141236, 0.1097496, 0.117126, 0.1133892, 0.10098, 0.0989712, 0.110268,
		0.0956124, 0.0932904, 0.0821664, 0.098604, 0.0999, 0.1018224, 0.0959688, 0.0951912, 0.0915948, 0.0884304, 0.0828252, 0.0859896,
		0.08262, 0.0815832, 0.0806112, 0.0816372, 0.0805896, 0.0819936, 0.0820476, 0.0819288, 0.0826416, 0.0868968, 0.093258, 0.0823176,
		0.0955908, 0.1033236, 0.1161756, 0.1029456, 0.1134108, 0.121608, 0.1297296, 0.1245348, 0.1305396, 0.13365, 0.1330128, 0.1468476,
		0.1373328, 0.1360584, 0.1296756, 0.1483164, 0.1417392, 0.1354968, 0.1306152, 0.1399464, 0.1307556, 0.1324728, 0.1330128, 0.130572,
		0.1310904, 0.1309716, 0.1257984, 0.1287576, 0.1265436, 0.1220184, 0.1216296, 0.131598, 0.1293408, 0.125604, 0.1294164, 0.1215756,
		0.1311768, 0.135756, 0.1382076, 0.1193292, 0.125334, 0.131382, 0.1368252, 0.1242972, 0.1286712, 0.1312092, 0.136404, 0.1267164,
		0.1302372, 0.1288656, 0.1299024, 0.130464, 0.1234656, 0.125118, 0.125388, 0.1237572, 0.1211976, 0.1174176, 0.1159056, 0.1166184,
		0.1159056, 0.1127412, 0.1003428, 0.1113912, 0.1033884, 0.0988416, 0.092394, 0.1033128, 0.0989712, 0.0976752, 0.0914976, 0.0979776,
		0.0904608, 0.0846612, 0.07776, 0.0961956, 0.0902016, 0.094014, 0.0884952, 0.0942948, 0.0902556, 0.0896076, 0.0863568, 0.0886032,
		0.0860868, 0.0857628, 0.0835488, 0.0850716, 0.0846612, 0.0847584, 0.0844884, 0.083862, 0.0862056, 0.0890676, 0.0925992, 0.0836028,
		0.0909684, 0.0944028, 0.09639, 0.0945864, 0.1031508, 0.1096848, 0.1282068, 0.1287144, 0.1308744, 0.125712, 0.119016, 0.1438884,
		0.1369764, 0.128844, 0.11097, 0.1445364, 0.1201176, 0.1076544, 0.0957312, 0.1113048, 0.0972972, 0.0972216, 0.09558, 0.0978048,
		0.0977832, 0.0989604, 0.1014984, 0.0976428, 0.0992088, 0.098658, 0.1088316, 0.103356, 0.1152792, 0.1176336, 0.1199124, 0.1126224,
		0.126846, 0.1337364, 0.1404108, 0.1268244, 0.1355184, 0.1502928, 0.1640844, 0.1457352, 0.1597752, 0.1724976, 0.1925856, 0.1634148,
		0.1718928, 0.1700676, 0.1652076, 0.1658448, 0.1572804, 0.1510596, 0.1551312, 0.1505196, 0.1475064, 0.1447524, 0.1394712, 0.1473768,
		0.1395252, 0.131004, 0.1210356, 0.13095, 0.1262088, 0.1194696, 0.1115532, 0.1242864, 0.1203336, 0.1124064, 0.0986256, 0.105138,
		0.0962496, 0.095958, 0.0912924, 0.0987768, 0.0951588, 0.0936792, 0.0948888, 0.093798, 0.091476, 0.0940896, 0.0940248, 0.0926316,
		0.0894024, 0.0920808, 0.0932148, 0.0888732, 0.0912168, 0.0925668, 0.0943812, 0.088074, 0.0925344, 0.0956448, 0.102006, 0.0979776,
		0.1093932, 0.1213164, 0.1264032, 0.111564, 0.1279584, 0.1382724, 0.1631016, 0.1521828, 0.1610496, 0.160974, 0.1655856, 0.1716444,
		0.1545048, 0.1449468, 0.135972, 0.1532952, 0.1413072, 0.1336932, 0.1302588, 0.1315764, 0.129816, 0.1240812, 0.1218348, 0.124632,
		0.124254, 0.1237356, 0.1213164, 0.1243836, 0.1230552, 0.1215108, 0.1209816, 0.1233036, 0.1254636, 0.1315872, 0.142182, 0.126846,
		0.132624, 0.146286, 0.2017332, 0.1386612, 0.1722384, 0.2024352, 0.201366, 0.1574424, 0.1718496, 0.2149092, 0.227934, 0.162324,
		0.1603692, 0.1578528, 0.1509732, 0.1516428, 0.1487052, 0.1444284, 0.140832, 0.1480464, 0.1487268, 0.1415772, 0.1398924, 0.1521504,
		0.1394388, 0.136188, 0.1204632, 0.1376028, 0.133164, 0.1283688, 0.1188, 0.1292652, 0.1229256, 0.1122228, 0.1032588, 0.10341,
		0.1009584, 0.0974052, 0.0951696, 0.1012176, 0.1000728, 0.096876, 0.095634, 0.0975564, 0.0963036, 0.0956448, 0.0950832, 0.0961308,
		0.0951588, 0.0945, 0.0943272, 0.09423, 0.0952128, 0.09504, 0.0950508, 0.0941868, 0.0947916, 0.095364, 0.0967464, 0.0954828,
		0.1053216, 0.1134108, 0.1226232, 0.1197612, 0.1322136, 0.1471068, 0.1691712, 0.1532736, 0.1542888, 0.1594944, 0.1665684, 0.1653264,
		0.1733724, 0.1687608, 0.1614708, 0.1878876, 0.1630044, 0.1606716, 0.1458972, 0.1761588, 0.1593648, 0.1559952, 0.1448604, 0.1566108,
		0.155412, 0.1485648, 0.14526, 0.1502496, 0.1479816, 0.1515564, 0.1529928, 0.152064, 0.1565352, 0.1632528, 0.1643112, 0.145638,
		0.1632312, 0.18063, 0.2146176, 0.16119, 0.1681668, 0.1792584, 0.204228, 0.1690956, 0.1880928, 0.2051352, 0.2143044, 0.187164,
		0.1911168, 0.1882764, 0.1844748, 0.1836324, 0.177228, 0.1724436, 0.1709856, 0.180036, 0.1693332, 0.1669032, 0.1577772, 0.1577556,
		0.1589976, 0.1464804, 0.129168, 0.1464156, 0.13797, 0.1247076, 0.1168452, 0.128304, 0.1250748, 0.1189944, 0.108108, 0.1143288,
		0.1009692, 0.0972, 0.09288, 0.1123416, 0.1144692, 0.1130004, 0.1059912, 0.1119312, 0.1031724, 0.0973188, 0.09639, 0.1015092,
		0.0963684, 0.0963144, 0.097524, 0.0972, 0.0965412, 0.0987876, 0.100062, 0.09612, 0.098118, 0.103734, 0.1117908, 0.0984312,
		0.1087452, 0.1125144, 0.1258524, 0.1137888, 0.1263708, 0.1409184, 0.1789344, 0.156276, 0.192456, 0.2014632, 0.216, 0.2385504,
		0.2412612, 0.216, 0.171126, 0.2376, 0.1974672, 0.1723032, 0.128574, 0.1861704, 0.1494288, 0.1544076, 0.1379808, 0.1553472,
		0.1440396, 0.1373436, 0.137592, 0.134028, 0.140994, 0.1411236, 0.142452, 0.1388988, 0.1452924, 0.1514592, 0.1674756, 0.1359396,
		0.16605, 0.1919808, 0.1973808, 0.1658232, 0.1829844, 0.2150496, 0.2849148, 0.2051352, 0.248778, 0.2717172, 0.3401352, 0.2652804,
		0.269244, 0.2515968, 0.236196, 0.2400516, 0.2249532, 0.2090772, 0.1964628, 0.1965276, 0.1793448, 0.181116, 0.1802412, 0.1870992,
		0.1650996, 0.1338984, 0.1255068, 0.1465344, 0.1311876, 0.1220184, 0.1113372, 0.1262196, 0.1206252, 0.1086804, 0.1011204, 0.1184652,
		0.1026, 0.0975996, 0.0929448, 0.1340712, 0.1165644, 0.1014984, 0.093258, 0.1068768, 0.1014876, 0.0995976, 0.10098, 0.0975996,
		0.0962928, 0.0942084, 0.09396, 0.0935712, 0.0918756, 0.0923292, 0.0906228, 0.0887652, 0.0943056, 0.0954288, 0.0976428, 0.0925344,
		0.0925776, 0.0924264, 0.0952992, 0.093852, 0.09531, 0.09801, 0.1114344, 0.1084752, 0.1165536, 0.1242756, 0.12609, 0.1319868,
		0.1261656, 0.1081188, 0.099684, 0.1244592, 0.1050624, 0.1062612, 0.1028376, 0.1109484, 0.1093932, 0.1083564, 0.102816, 0.1086912,
		0.1051488, 0.1076976, 0.1085832, 0.1111104, 0.1052028, 0.1071036, 0.1063692, 0.108702, 0.1078812, 0.1077084, 0.1124604, 0.1090908,
		0.1174284, 0.129222, 0.1500552, 0.1288116, 0.1378512, 0.1669788, 0.1417392, 0.1417716, 0.154278, 0.1590948, 0.1603584, 0.1549692,
		0.1591164, 0.1466748, 0.1380564, 0.1502928, 0.1456812, 0.1461996, 0.1368144, 0.1420416, 0.1414692, 0.1455948, 0.128196, 0.1447956,
		0.1414368, 0.12258, 0.10611, 0.1177308, 0.1093176, 0.104922, 0.0996084, 0.1090908, 0.104382, 0.1027296, 0.094176, 0.09504,
		0.090612, 0.0866052, 0.0843804, 0.1026648, 0.0959364, 0.081, 0.0725976, 0.0877176, 0.0794232, 0.0771768, 0.0768852, 0.0808272,
		0.0771336, 0.0741852, 0.0721548, 0.0703944, 0.0680508, 0.0684504, 0.066258, 0.0677592, 0.0663444, 0.0655128, 0.0634068, 0.0690012,
		0.0693576, 0.0702, 0.0897372, 0.0778788, 0.0875556, 0.0927396, 0.0991332, 0.0870264, 0.0937224, 0.1032048, 0.1050948, 0.1054512,
		0.1077948, 0.108108, 0.1026972, 0.1063152, 0.1034964, 0.1032696, 0.0989928, 0.1046196, 0.1026324, 0.1012608, 0.1013148, 0.1001052,
		0.1039716, 0.1037124, 0.1041768, 0.1030536, 0.1032588, 0.1037988, 0.1036908, 0.0999432, 0.1056672, 0.1079028, 0.1137888, 0.1073412,
		0.1113264, 0.123228, 0.1362096, 0.1121796, 0.1180116, 0.1305828, 0.1426032, 0.1365876, 0.1435536, 0.1503252, 0.1648512, 0.1353672,
		0.1396656, 0.1427436, 0.1470852, 0.140778, 0.140616, 0.142938, 0.1430784, 0.1432944, 0.1439316, 0.1450656, 0.1392444, 0.1424196,
		0.1345356, 0.1282392, 0.120474, 0.127386, 0.1213056, 0.107136, 0.0936792, 0.1198908, 0.1137132, 0.0985176, 0.0885492, 0.0951696,
		0.0813456, 0.0781704, 0.0755892, 0.0865296, 0.0807948, 0.0814968, 0.080352, 0.079812, 0.0758268, 0.0764748, 0.0775224, 0.0750168,
		0.0803844, 0.0801468, 0.0823716, 0.0785808, 0.0799308, 0.0842508, 0.0848988, 0.0798444, 0.083862, 0.0820584, 0.0877392, 0.0772416,
		0.0957852, 0.1101708, 0.1253124, 0.1055484, 0.129546, 0.146718, 0.1725084, 0.1499688, 0.1659744, 0.183708, 0.1785348, 0.1658124,
		0.1652616, 0.1625508, 0.153684, 0.1631556, 0.1523772, 0.1378404, 0.1278828, 0.1385856, 0.12987, 0.136026, 0.1415448, 0.1572588,
		0.1582416, 0.1559196, 0.1683936, 0.169668, 0.1736316, 0.1724544, 0.1817208, 0.175068, 0.1814292, 0.2017224, 0.2133864, 0.2027916,
		0.2447064, 0.2362284, 0.2321028, 0.196776, 0.21897, 0.252828, 0.2788668, 0.2204712, 0.2446848, 0.2858112, 0.340632, 0.2531628,
		0.2888892, 0.2923668, 0.298782, 0.2930472, 0.2517804, 0.2397168, 0.220428, 0.2357424, 0.2126952, 0.210384, 0.1889136, 0.2196504,
		0.189054, 0.1816668, 0.1619676, 0.1788696, 0.1577124, 0.1438344, 0.1326564, 0.1512972, 0.145962, 0.1328184, 0.1205172, 0.12825,
		0.1172988, 0.1134324, 0.1083888, 0.1123848, 0.111186, 0.1153872, 0.113238, 0.1151172, 0.1150848, 0.1090368, 0.109188, 0.1112184,
		0.1101924, 0.1110672, 0.1121256, 0.1131084, 0.1077192, 0.1092852, 0.1109592, 0.1130112, 0.115938, 0.1120932, 0.117612, 0.1094688,
		0.113184, 0.1215216, 0.1409184, 0.129222, 0.1683396, 0.1977264, 0.2568024, 0.1998, 0.306774, 0.3456432, 0.3712932, 0.3163968,
		0.2679264, 0.2565216, 0.2483244, 0.2625588, 0.2572884, 0.2191428, 0.1991412, 0.2610144, 0.2277936, 0.214866, 0.1888164, 0.2027052,
		0.2198664, 0.2391012, 0.2314008, 0.2283768, 0.2144016, 0.2366928, 0.2671812, 0.2437992, 0.2557764, 0.246834, 0.2389932, 0.2352348,
		0.2929608, 0.34992, 0.3510216, 0.3056076, 0.3190212, 0.3380616, 0.364176, 0.2536704, 0.323244, 0.356292, 0.3898908, 0.2685204,
		0.2963628, 0.2967084, 0.2757672, 0.296946, 0.301266, 0.2890836, 0.2517372, 0.342198, 0.2384856, 0.183708, 0.1515132, 0.211356,
		0.1722492, 0.1484244, 0.1334988, 0.166536, 0.1370412, 0.1233144, 0.1116396, 0.1262844, 0.1221588, 0.1149984, 0.107352, 0.1246752,
		0.1088748, 0.0987336, 0.0905688, 0.1047384, 0.095472, 0.097092, 0.0959472, 0.0980532, 0.094176, 0.084024, 0.0963252, 2(0.0960552),
		2(0.0965952), 0.0979452, 0.0981828, 0.09963, 0.0993816, 0.0964332, 0.098172, 0.0998892, 0.1026216, 0.0944784, 0.0997704, 0.1112508,
		0.1211004, 0.1045332, 0.122472, 0.13662, 0.1677024, 0.1546776, 0.1923156, 0.2144556, 0.243162, 0.2235816, 0.2319516, 0.2809512,
		0.2521908, 0.2592, 0.2130084, 0.2146932, 0.1900152, 0.2118204, 0.2096496, 0.189, 0.17334, 0.1959012, 0.1836864, 0.1779192,
		0.176742, 0.1770444, 0.1714176, 0.1768608, 0.177012, 0.1776168, 0.1862568, 0.1880604, 0.176742, 0.172746, 0.1831248, 0.2098548,
		0.221778, 0.180738, 0.2132568, 0.2515644, 0.3065256, 0.225072, 0.2904984, 0.328104, 0.3870936, 0.3004776, 0.3082644, 0.3121416,
		0.3099816, 0.280368, 0.227988, 0.2415852, 0.2241108, 0.2368008, 0.2052, 0.1817748, 0.16578, 0.1873152, 0.1607904, 0.1384236,
		0.1197612, 0.1507896, 0.1333908, 0.1110996, 0.098712, 0.1279908, 0.113238, 0.1018116, 0.0975024, 0.1086048, 0.098172, 0.0951048,
		0.0887544, 0.1015956, 0.0985068, 0.0948348, 0.0939708, 0.0962604, 0.0928368, 0.0894348, 0.086454, 0.0908388, 0.0881064, 0.0863136,
		0.0821016, 0.0885816, 0.0870264, 0.084618, 0.0780948, 0.0845208, 0.0848664, 0.0922644, 0.093852, 0.0911412, 0.0807192, 0.093798,
		0.0973296, 0.0961632, 0.1184328, 0.1269972, 0.139968, 0.1245996, 0.141264, 0.1465884, 0.1503684, 0.1533384, 0.1553472, 0.1446228,
		0.1203444, 0.1497096, 0.1488348, 0.1257984, 0.1006992, 0.137484, 0.124956, 0.1164348, 0.1032804, 0.1153008, 0.1165968, 0.1163484,
		0.112374, 0.1096632, 0.1140156, 0.1136808, 0.1189404, 0.1243944, 0.1265544, 0.1292436, 0.1317168, 0.1272888, 0.1428408, 0.1604016,
		0.16713, 0.143262, 0.1556172, 0.1629396, 0.1739448, 0.1658556, 0.1695708, 0.177822, 0.1781784, 0.1657368, 0.1574532, 0.1555848,
		0.1527336, 0.1485432, 0.147582, 0.1482408, 0.1487484, 0.1488456, 0.1500336, 0.1486944, 0.1300104, 0.1442124, 0.135054, 0.1243836,
		0.1205604, 0.1244376, 0.1137348, 0.1122336, 0.1045656, 0.1155492, 0.1117584, 0.0976752, 0.0893376, 0.1048464, 0.088344, 0.0776628,
		0.0560088, 0.0926316, 0.0960552, 0.093042, 0.0954504, 0.0868536, 0.0799308, 0.0742176, 0.0658692, 0.0807948, 0.0745308, 0.0830196,
		0.0726084, 0.0791856, 0.0883224, 0.0899856, 0.0914976, 0.0687852, 0.0691416, 0.088776, 0.0972648, 0.09747, 0.1058724, 0.1144584,
		0.1232604, 0.1081512, 0.1269972, 0.1357452, 0.1554984, 0.1389096, 0.1557036, 0.1685556, 0.1734264, 0.1615788, 0.1600992, 0.1546992,
		0.1393956, 0.1722276, 0.1513836, 0.1440828, 0.1191024, 0.1480896, 0.126684, 0.128574, 0.1137132, 0.1308096, 0.1247292, 0.1218888,
		0.1060668, 0.125388, 0.1191456, 0.1240488, 0.1253556, 0.1260468, 0.1269108, 0.13041, 0.111996, 0.1254204, 0.14121, 0.1686852,
		0.1800036, 0.1280556, 0.1404972, 0.157518, 0.1604664, 0.1448496, 0.1528524, 0.1596456, 0.1654344, 0.1482624, 0.149256, 0.1468584,
		0.14661, 0.1414476, 0.1409508, 0.151416, 0.1453572, 0.1532196, 0.1459188, 0.1440288, 0.1298808, 0.14553, 0.13797, 0.1274724,
		0.1231092, 0.1289952, 0.1270836, 0.1242648, 0.1117476, 0.133812, 0.121122, 0.1164888, 0.1065096, 0.12069, 0.1050516, 0.0930312,
		0.0881712, 0.1094688, 0.108432, 0.1040472, 0.0977292, 0.09882, 0.098874, 0.099846, 0.1047276, 0.1024704, 0.0963252, 0.0974592,
		0.0966492, 0.09612, 0.0984744, 0.0981612, 0.0971568, 0.09396, 0.097686, 0.100602, 0.1041228, 0.1016064, 0.1008828, 0.1050408,
		0.1152252, 0.0877608, 0.1056456, 0.1179144, 0.1214028, 0.1164888, 0.1215, 0.1251828, 0.1284876, 0.1285524, 0.1239084, 0.1234548,
		0.1224072, 0.1280664, 0.1238004, 0.1181304, 0.1138104, 0.1217808, 0.114966, 0.1117692, 0.1068552, 0.1128708, 0.1126116, 0.1112508,
		0.11016, 0.1131624, 0.1110996, 0.109188, 0.1074168, 0.1131948, 0.1040688, 0.104328, 0.106164, 0.1060776, 0.1096956, 0.1153332,
		0.1326024, 0.1128276, 0.1253124, 0.1316952, 0.1458756, 0.1339092, 0.1461348, 0.1510272, 0.1546992, 0.145368, 0.145638, 0.145476,
		0.1452816, 0.1444608, 0.1484568, 0.1483812, 0.13419, 0.1477872, 0.1478736, 0.1426032, 0.1231632, 0.1485, 0.1413504, 0.1293408,
		0.1113048, 0.1346976, 0.12825, 0.124038, 0.1101168, 0.1324188, 0.1281312, 0.12042, 0.1044684, 0.131544, 0.1118124, 0.1010772,
		0.0900612, 0.1144044, 0.1113372, 0.0992412, 0.0932256, 0.104976, 0.1014444, 0.0998892, 0.1015092, 0.0977616, 0.0937656, 0.096822,
		0.0925236, 0.094446, 0.0928476, 0.0939924, 0.0939276, 0.0905256, 0.0906552, 0.091098, 0.096174, 0.0937656, 0.0972864, 0.1012284,
		0.1049004, 0.0973836, 0.0994788, 0.105948, 0.108216, 0.1030212, 0.1068876, 0.1049652, 0.1052244, 0.1056132, 0.1058508, 0.1025352,
		0.0980748, 0.107028, 0.1045008, 0.0952668, 0.096012, 0.0997488, 0.0931392, 0.0947916, 0.0934632, 0.0931176, 0.09477, 0.0959688,
		0.0972108, 0.1003104, 0.088128, 0.0890784, 0.0927504, 0.0936036, 0.0932148, 0.1004508, 0.1060128, 0.0947376, 0.104004, 0.1143828,
		0.1219968, 0.10071, 0.1150848, 0.12771, 0.129114, 0.1229364, 0.1315548, 0.1415664, 0.143748, 0.1355508, 0.1344492, 0.138132,
		0.1413072, 0.1379592, 0.1400004, 0.1367388, 0.140886, 0.1425816, 0.140022, 0.139644, 0.1380564, 0.1443096, 0.14256, 0.1415772,
		0.1275912, 0.138942, 0.1306908, 0.1278504, 0.118692, 0.1286712, 0.1278288, 0.1240164, 0.1142964, 0.1194048, 0.1098684, 0.105516,
		0.0931932, 0.1131192, 0.111672, 0.1066392, 0.1051272, 0.1120716, 0.1089288, 0.1078596, 0.1041984, 0.10773, 0.1051488, 0.1056348,
		0.1036368, 0.096498, 0.099846, 0.1029456, 0.1045548, 0.1035072, 0.1060128, 0.108324, 0.1073304, 0.1008072, 0.1090476, 0.114426,
		0.1336824, 0.1189512, 0.1379808, 0.1640412, 0.1694196, 0.1544292, 0.1560816, 0.1530468, 0.169884, 0.1934388, 0.1766664, 0.16794,
		0.16092, 0.170586, 0.1651644, 0.1589868, 0.1494072, 0.15552, 0.1529064, 0.1508328, 0.14769, 0.1472256, 0.1473228, 0.1503144,
		0.1488888, 0.1502064, 0.1497204, 0.15417, 0.159138, 0.1496124, 0.160758, 0.1629396, 0.1595808, 0.1519236, 0.1681344, 0.1803816,
		0.1939572, 0.1826928, 0.1945836, 0.213894, 0.2224044, 0.2277612, 0.2348784, 0.2441232, 0.2522772, 0.2072304, 0.2120904, 0.2090232,
		0.195696, 0.2249316, 0.231174, 0.2159784, 0.214002, 0.222588, 0.2004588, 0.2000484, 0.187542, 0.197208, 0.1831572, 0.1678752,
		0.1445796, 0.175608, 0.1553472, 0.142236, 0.121878, 0.1458972, 0.1396548, 0.135972, 0.1217052, 0.1288764, 0.12366, 0.1182384,
		0.109242, 0.1239732, 0.1171692, 0.1140804, 0.104274, 0.113022, 0.1108296, 0.1079676, 0.1127844, 0.111834, 0.1069092, 0.1076652,
		0.1032264, 0.1053432, 0.1025352, 0.1027296, 0.1042632, 0.1014552, 0.1019736, 0.1066932, 0.1144908, 0.0983448, 0.1137024, 0.115992,
		0.1233792, 0.1214568, 0.12771, 0.146502, 0.1633716, 0.1562868, 0.1715256, 0.1918404, 0.205254, 0.1781676, 0.1747764, 0.1851228,
		0.168642, 0.1846152, 0.1776492, 0.1644516, 0.1474092, 0.1717524, 0.1635876, 0.16443, 0.161892, 0.162918, 0.1591272, 0.1584576,
		0.1504548, 0.1474848, 0.1517292, 0.1537596, 0.1547964, 0.1536516, 0.1692684, 0.1803708, 0.1685664, 0.14553, 0.1601424, 0.180198,
		0.2060964, 0.1708668, 0.181764, 0.1917, 0.2145312, 0.1893132, 0.1996488, 0.2076516, 0.2198232, 0.2053728, 0.2122308, 0.1957392,
		0.1875312, 0.1779732, 0.1797984, 0.1855656, 0.1879956, 0.1908684, 0.1714932, 0.178578, 0.1654452, 0.1870776, 0.1668924, 0.1512864,
		0.1354428, 0.1522908, 0.1479276, 0.1387476, 0.123822, 0.1431432, 0.1329372, 0.1261764, 0.117882, 0.1219212, 0.1177308, 0.112482,
		0.1028808, 0.121824, 0.1130112, 0.1091124, 0.108432, 0.12069, 0.1110132, 0.1089396, 0.111564, 0.1114884, 0.1094688, 0.1079892,
		0.1064556, 0.109134, 0.1088748, 0.1083564, 0.108378, 0.1092096, 0.1113804, 0.111726, 0.1157112, 0.1058508, 0.1119204, 0.117234,
		0.131652, 0.1193076, 0.1472364, 0.1599696, 0.1925208, 0.1549476, 0.1842048, 0.232416, 0.223884, 0.23328, 0.2563488, 0.264546,
		0.2301048, 0.26676, 0.2391552, 0.1847988, 0.1839024, 0.2092176, 0.1837728, 0.1773684, 0.17577, 0.176904, 0.1724976, 0.1721736,
		0.1749708, 0.169074, 0.1607904, 0.1695168, 0.177984, 0.1774008, 0.1774224, 0.18549, 0.18765, 0.181062, 0.1967544, 0.2258172,
		0.2212596, 0.2022732, 0.2242188, 0.2771064, 0.3039768, 0.2480112, 0.3156732, 0.3419172, 0.369846, 0.2847528, 0.2962332, 0.266382,
		0.235062, 0.2287224, 0.2302128, 0.20979, 0.192996, 0.2155896, 0.184896, 0.1697328, 0.1604556, 0.1821528, 0.1597644, 0.1440072,
		0.132624, 0.1472364, 0.1407132, 0.1264896, 0.1204632, 0.1497204, 0.13473, 0.1243296, 0.1172448, 0.1333368, 0.1220832, 0.1149552,
		0.109944, 0.113994, 0.1122768, 0.1079352, 0.103032, 0.1107756, 0.10611, 0.1015956, 0.09936, 0.1028808, 0.1001808, 0.1003212,
		0.102114, 0.1031076, 0.1015416, 0.1012176, 0.1003752, 0.1026756, 0.1055268, 0.1072764, 0.1108836, 0.1060668, 0.1110348, 0.11448,
		0.1262844, 0.1098684, 0.1268136, 0.14688, 0.1624428, 0.1497852, 0.1721196, 0.1694412, 0.175392, 0.1676268, 0.18333, 0.1866024,
		0.1677132, 0.1873476, 0.1754352, 0.1682964, 0.1534356, 0.1644192, 0.1500552, 0.15309, 0.1523664, 0.1529604, 0.1530144, 0.156168,
		0.1523988, 0.1568808, 0.1511892, 0.1485864, 0.1525608, 0.1536192, 0.1594296, 0.1565352, 0.1616004, 0.152442, 0.1625832, 0.1706292,
		0.1712232, 0.1561896, 0.1631556, 0.1577772, 0.1752084, 0.155088, 0.1660176, 0.1711692, 0.1770768, 0.1578096, 0.1636416, 0.1578744,
		0.1602828, 0.15579, 0.1539972, 0.1590408, 0.1645164, 0.1642572, 0.1533168, 0.1518048, 0.1421928, 0.152928, 0.1492452, 0.1350972,
		0.1242972, 0.14337, 0.134298, 0.124038, 0.1174392, 0.1267812, 0.1260036, 0.1218564, 0.1142424, 0.1190484, 0.1139508, 0.1069308,
		0.0968868, 0.11475, 0.1096956, 0.1066176, 0.1018332, 0.1111212, 0.1077192, 0.1051704, 0.1023408, 0.103356, 0.1036692, 0.1039284,
		0.098442, 0.097632, 0.100494, 0.1018008, 0.1086912, 0.1033884, 0.1040688, 0.1099872, 0.1130976, 0.103248, 0.1090692, 0.1148904,
		0.1282068, 0.1062396, 0.124092, 0.1396764, 0.1755756, 0.1504548, 0.1649484, 0.167346, 0.1690632, 0.170154, 0.183006, 0.1982988,
		0.203634, 0.2046924, 0.1935252, 0.1786104, 0.1750248, 0.1789452, 0.1812132, 0.1796688, 0.1728, 0.1798848, 0.1775304, 0.1750248,
		0.1677348, 0.1724112, 0.1639872, 0.1616328, 0.1602936, 0.1606068, 0.1612116, 0.1604988, 0.1570968, 0.1581984, 0.1587816, 0.1650888,
		0.1660824, 0.1558764, 0.15606, 0.1675404, 0.1681776, 0.154008, 0.165618, 0.1721736, 0.1739124, 0.1664928, 0.1601316, 0.1635876,
		0.1513728, 0.1635444, 0.1547856, 0.1496232, 0.133866, 0.1512864, 0.1411236, 0.1348056, 0.1172016, 0.1303236, 0.1273104, 0.1181844,
		0.1063584, 0.1196748, 0.1134972, 0.107244, 0.0991548, 0.1126764, 0.1081296, 0.1014012, 0.0976212, 0.1094796, 0.0983988, 0.0868968,
		0.0784512, 0.1037232, 0.0908604, 0.0865188, 0.0858816, 0.0963684, 0.0887976, 0.0855252, 0.076842, 0.0897048, 0.0853092, 0.0800388,
		0.0781272, 0.0854604, 0.0858816, 0.0857412, 0.08802, 0.0868536, 0.087858, 0.0931068, 0.0925776, 0.0944784, 0.0919512, 0.0932796,
		0.0957528, 0.08721, 0.0993924, 0.1053, 0.112104, 0.103356, 0.10746, 0.1143612, 0.1189728, 0.117072, 0.1184004, 0.11988,
		0.1194048, 0.120528, 0.118314, 0.1160568, 0.11232, 0.112104, 0.1112616, 0.1098576, 0.1073844, 0.1109268, 0.1111536, 0.108378,
		0.1075788, 0.110214, 0.106974, 0.1053864, 0.1073844, 0.1081512, 0.1087236, 0.1112832, 0.114156, 0.1087344, 0.1131624, 0.1173312,
		0.1283364, 0.1181736, 0.1223316, 0.1251612, 0.1325916, 0.1253988, 0.1330452, 0.1356912, 0.1387152, 0.13203, 0.131544, 0.131868,
		0.131976, 0.13095, 0.1312416, 0.1323432, 0.1277208, 0.1347084, 0.1306368, 0.1300752, 0.128736, 0.1408536, 0.1310796, 0.123876,
		0.118584, 0.1199232, 0.1142748, 0.108432, 0.100116, 0.110376, 0.1052568, 0.1020816, 0.0985716, 0.1053972, 0.1023084, 0.0959364,
		0.0885276, 0.1006344, 0.0940248, 0.0929556, 0.090288, 0.0925452, 0.0909468, 0.0886572, 0.092178, 0.0932148, 0.0915192, 0.0879768,
		0.0878256, 0.0858708, 0.08424, 0.0817344, 0.0834084, 0.0872856, 0.0861516, 0.0826416, 0.0864864, 0.086454, 0.086022, 0.0859788,
		0.0855144, 0.0847368, 0.0887976, 0.0925668, 0.0941004, 0.0922752, 0.094608, 0.096174, 0.100278, 0.0951588, 0.096714, 0.0969408,
		0.1001268, 0.1005912, 0.1034748, 0.0977616, 0.0971136, 0.1054512, 0.1047708, 0.1011852, 0.1051596, 0.10071, 0.1047168, 0.1062504,
		0.1068444, 0.1077624, 0.1068876, 0.1080108, 0.1070172, 0.1069308, 0.1072764, 0.1106136, 0.1180332, 0.1093608, 0.1141992, 0.118314,
		0.1244484, 0.1184976, 0.1214784, 0.1223748, 0.124848, 0.1224612, 0.1233576, 0.1254744, 0.132084, 0.1165428, 0.1157004, 0.110592,
		0.1073088, 0.1214892, 0.1189728, 0.1164672, 0.1123092, 0.1173312, 0.1180008, 0.118692, 0.1209816, 0.123714, 0.1230552, 0.1179684,
		0.1052244, 0.1158948, 0.114534, 0.0995004, 0.0931176, 0.1098252, 0.1023732, 0.0917352, 0.0885168, 0.0952128, 0.089964, 0.0836136,
		0.071442, 0.0928368, 0.0894996, 0.0864432, 0.0855576, 0.090342, 0.0904068, 0.086832, 0.083916, 0.0821232, 0.0848124, 0.0850284,
		0.0754704, 0.0865512, 0.0840132, 0.0871344, 0.0872532, 0.0835704, 0.0858384, 0.0873504, 0.0877932, 0.0818748, 0.0892836, 0.0927504,
		0.1103652, 0.0899424, 0.10584, 0.1184652, 0.1300212, 0.120312, 0.1307664, 0.133542, 0.1343844, 0.1306044, 0.1309068, 0.129114,
		0.1267704, 0.1280988, 0.1281096, 0.1205388, 0.1101384, 0.13041, 0.1171692, 0.1100844, 0.1062504, 0.1155816, 0.1136484, 0.1106028,
		0.1112616, 0.109674, 0.1088316, 0.1114236, 0.1191888, 0.1108188, 0.1176012, 0.1212624, 0.1216296, 0.105246, 0.1258632, 0.1386936,
		0.1338876, 0.1208844, 0.1277748, 0.1301616, 0.1347516, 0.1325268, 0.1420524, 0.1426572, 0.1415556, 0.1479276, 0.1367388, 0.1320192,
		0.1317384, 0.1338876, 0.131274, 0.1306368, 0.1313388, 0.1351296, 0.1353672, 0.1328832, 0.1322352, 0.1358532, 0.1305828, 0.1261656,
		0.1172124, 0.1287792, 0.1242648, 0.123714, 0.108594, 0.1235628, 0.1190268, 0.108918, 0.0981828, 0.1074384, 0.0991548, 0.0944568,
		0.0916704, 0.1008504, 0.0971676, 0.090126, 0.0900828, 0.0958392, 0.0940788, 0.0923616, 0.0904824, 0.0972864, 0.0934632, 0.0915732,
		0.090828, 0.0921456, 0.0917028, 0.092664, 0.0925992, 0.0930204, 0.0941112, 0.0975888, 0.1031184, 0.0906336, 0.1005264, 0.1095768,
		0.130302, 0.11367, 0.1262628, 0.1443852, 0.1705104, 0.1288116, 0.1363284, 0.1445904, 0.1486836, 0.1483272, 0.1463508, 0.1374408,
		0.1289412, 0.1409184, 0.1284336, 0.1253124, 0.1237032, 0.1317924, 0.123066, 0.1227852, 0.1201176, 0.1234548, 0.1225368, 0.1223316,
		0.1208304, 0.1253016, 0.125388, 0.1207008, 0.1200528, 0.1271268, 0.127062, 0.127872, 0.1305504, 0.127602, 0.1450548, 0.1519668,
		0.1538244, 0.1243944, 0.1339308, 0.1392336, 0.1600992, 0.1375056, 0.1499364, 0.1556604, 0.1638576, 0.1525824, 0.1466964, 0.1432944,
		0.1397088, 0.1450764, 0.1410912, 0.1458, 0.1445472, 0.1466208, 0.1542564, 0.1430352, 0.129762, 0.153738, 0.135432, 0.126684,
		0.120852, 0.1369764, 0.1349784, 0.1270944, 0.1128708, 0.1263816, 0.1207548, 0.1164024, 0.1077948, 0.1101384, 0.0972108, 0.0912384,
		0.0845748, 0.0930096, 0.0954936, 0.0944568, 0.0915948, 0.0934308, 0.0923184, 0.092016, 0.0918972, 0.0907092, 0.0911628, 0.0913572,
		0.090234, 0.0918216, 0.0929124, 0.0923508, 0.0924048, 0.0915516, 0.092772, 0.0944892, 0.0994356, 0.0901692, 0.0972108, 0.1026108,
		0.1178172, 0.0966924, 0.1152252, 0.1328724, 0.152928, 0.1402272, 0.1508544, 0.1601208, 0.162486, 0.1512432, 0.14769, 0.1581552,
		0.1454436, 0.1597968, 0.1446444, 0.1276128, 0.1163592, 0.1378944, 0.1274832, 0.119502, 0.1111644, 0.1170612, 0.110322, 0.10827,
		0.1084212, 0.1086372, 0.1057644, 0.1070388, 0.1071576, 0.1108944, 0.1125792, 0.1127196, 0.1176552, 0.1162296, 0.1262196, 0.1323756,
		0.1486944, 0.1231416, 0.1302804, 0.1477656, 0.1550016, 0.1393632, 0.1500768, 0.1517508, 0.1571724, 0.1451088, 0.1472364, 0.1513944,
		0.1540836, 0.1483812, 0.1489968, 0.1508652, 0.1507896, 0.1579176, 0.154818, 0.1483164, 0.1386288, 0.161892, 0.1546236, 0.1443096,
		0.1267812, 0.152766, 0.1431648, 0.1315008, 0.1215972, 0.1335852, 0.129276, 0.127872, 0.1075356, 0.12528, 0.114156, 0.1044252,
		0.0951588, 0.1088208, 0.1054836, 0.1009368, 0.0978264, 0.0994464, 0.0985608, 0.0989496, 0.0981936, 0.0987552, 0.0974052, 0.0955368,
		0.0940788, 0.0964872, 0.0953208, 0.0967464, 0.0969408, 0.0976212, 0.0981828, 0.0983988, 0.099954, 0.0939384, 0.1019196, 0.1080432,
		0.12204, 0.1089288, 0.124794, 0.1358208, 0.1436508, 0.1276776, 0.1378512, 0.1422684, 0.1444284, 0.1538028, 0.1495908, 0.1398708,
		0.1314792, 0.1466208, 0.1404, 0.1339524, 0.1271808, 0.1398924, 0.1330344, 0.1302048, 0.1214136, 0.1252692, 0.1225368, 0.1211868,
		0.12015, 0.1196532, 0.1183896, 0.1145448, 0.113994, 0.1195452, 0.1201176, 0.1212732, 0.1228932, 0.1218672, 0.1257336, 0.1359612,
		0.150336, 0.1260036, 0.1380024, 0.1415772, 0.216918, 0.141102, 0.1468692, 0.1454004, 0.1493316, 0.141264, 0.1430568, 0.1400112,
		0.143154, 0.137646, 0.1348272, 0.1394496, 0.142884, 0.144666, 0.1408752, 0.136458, 0.1325052, 0.1457784, 0.138186, 0.1295568,
		0.1246212, 0.1374948, 0.131166, 0.1222236, 0.1112292, 0.1242972, 0.1160136, 0.117072, 0.1053324, 0.1161324, 0.1053648, 0.0996408,
		0.0945972, 0.1081512, 0.1072224, 0.102708, 0.10071, 0.106164, 0.1022652, 0.1035504, 0.1032588, 0.1055268, 0.1032264, 0.1045008,
		0.1050516, 0.1043064, 0.1036692, 0.1009152, 0.1045224, 0.0977076, 0.1033128, 0.1056132, 0.1046736, 0.1003536, 0.1056996, 0.110754,
		0.1193508, 0.1142532, 0.1391796, 0.1483488, 0.1495476, 0.1338552, 0.14013, 0.1446336, 0.1480896, 0.1463508, 0.1484136, 0.1459944,
		0.1412424, 0.1456488, 0.1381104, 0.1365768, 0.1337256, 0.1410912, 0.139158, 0.1304208, 0.1251936, 0.1345896, 0.1305612, 0.1301724,
		0.1269, 0.1223748, 0.124146, 0.1244052, 0.1261224, 0.1255392, 0.1273536, 0.133812, 0.1377864, 0.1271592, 0.135108, 0.1483164,
		0.1540404, 0.1357992, 0.1409832, 0.1525932, 0.1574964, 0.151902, 0.1632744, 0.18036, 0.1882548, 0.15687, 0.1605636, 0.1527228,
		0.148716, 0.1463508, 0.1437804, 0.1438776, 0.1441692, 0.1459944, 0.1418256, 0.1408212, 0.1344384, 0.1474524, 0.1355832, 0.1297188,
		0.1182816, 0.139914, 0.1260468, 0.1183248, 0.1124928, 0.1234116, 0.1197072, 0.1172124, 0.1064556, 0.1165968, 0.1114668, 0.1019844,
		0.0959688, 0.1183788, 0.1147932, 0.112104, 0.0963252, 0.111618, 0.1089288, 0.1045116, 0.1006236, 0.107946, 0.1016064, 0.1022112,
		0.0987336, 0.1037016, 0.0961524, 0.0982368, 0.094446, 0.0969516, 0.0987876, 0.0990684, 0.1012932, 0.10071, 0.1020816, 0.1067688,
		0.1076544, 0.1019844, 0.1060884, 0.1160028, 0.1180764, 0.118584, 0.1191672, 0.1173636, 0.121338, 0.1190808, 0.1177092, 0.1238328,
		0.1207332, 0.1190484, 0.1193724, 0.1187784, 0.1139832, 0.1190052, 0.1163808, 0.1118772, 0.1075464, 0.1133676, 0.1110672, 0.1094364,
		0.1047924, 0.1106892, 0.1067796, 0.1060668, 0.1044684, 0.1084104, 0.1073628, 0.1078812, 0.1097604, 0.1032912, 0.1068444, 0.1172772,
		0.1240704, 0.1177416, 0.1282176, 0.132138, 0.1347948, 0.1261656, 0.1306152, 0.1347408, 0.1373868, 0.1323864, 0.1335312, 0.1325916,
		0.1318032, 0.1294488, 0.1283256, 0.1325268, 0.1300104, 0.133164, 0.129816, 0.1289304, 0.125658, 0.1363392, 0.1261872, 0.1189728,
		0.1117044, 0.1287576, 0.1181196, 0.1126764, 0.1027296, 0.123228, 0.1174608, 0.1085076, 0.095148, 0.1108728, 0.1067796, 0.0987336,
		0.0922968, 0.1053, 0.0992736, 0.0970488, 0.095958, 0.108108, 0.1046088, 0.0940896, 0.0900612, 0.0980208, 0.0925236, 0.0910764,
		0.090342, 0.0888948, 0.0894672, 0.0884628, 0.0880632, 0.092502, 0.0927504, 0.0933768, 0.0939168, 0.0896508, 0.092502, 0.0959688,
		0.097902, 0.0862164, 0.0911844, 0.0964008, 0.1066932, 0.1033128, 0.0976428, 0.0964656, 0.0967788, 0.0940464, 0.0951696, 0.106326,
		0.1091556, 0.1116504, 0.1160352, 0.1099332, 0.1081728, 0.1114236, 0.111078, 0.1105596, 0.1066932, 0.1093932, 0.109296, 0.1086048,
		0.1066068, 0.1074492, 0.1037124, 0.1011528, 0.1005588, 0.0886464, 0.1037664, 0.1028916, 0.1040256, 0.0969084, 0.0987336, 0.1038528,
		0.1106892, 0.1002996, 0.1089612, 0.1195668, 0.1233684, 0.1213056, 0.1224288, 0.1266624, 0.1330128, 0.127062, 0.128412, 0.1242972,
		0.1244808, 0.1291788, 0.1263384, 0.1247832, 0.1282824, 0.1320516, 0.1272348, 0.1304424, 0.122634, 0.1278288, 0.1220508, 0.1203552,
		0.1135944, 0.124794, 0.1178388, 0.1082916, 0.0987336, 0.114858, 0.1118448, 0.1026216, 0.095472, 0.1072764, 0.1016712, 0.0984852,
		0.0885708, 0.0979236, 0.0961848, 0.0928476, 0.0945864, 0.09423, 0.0926748, 0.0921348, 0.0923616, 0.0922968, 0.0928908, 0.0935388,
		0.0935064, 0.093096, 0.0914544, 0.0933768, 0.0937332, 0.0921672, 0.0939276, 0.0956232, 0.1019628, 0.0829764, 0.0947916, 0.1109916,
		0.1210032, 0.1180764, 0.13122, 0.1458864, 0.1545696, 0.14013, 0.1435644, 0.1451628, 0.152064, 0.152172, 0.1497528, 0.14418,
		0.1369224, 0.1657908, 0.1484784, 0.1276884, 0.1203876, 0.1414908, 0.1277532, 0.12582, 0.1232064, 0.1249452, 0.1285416, 0.1185516,
		0.1181412, 0.1138212, 0.11232, 0.1138104, 0.1188648, 0.1207332, 0.1273644, 0.1325808, 0.1358424, 0.1188108, 0.1277856, 0.1549368,
		0.1988172, 0.131976, 0.2125656, 0.1683072, 0.1829628, 0.1932444, 0.1689228, 0.173178, 0.1780272, 0.1461888, 0.1476468, 0.1579824,
		0.1564596, 0.150336, 0.1511244, 0.1572264, 0.1529388, 0.1567512, 0.1518912, 0.144558, 0.1429056, 0.1483488, 0.1400868, 0.1343088,
		0.126144, 0.1362744, 0.1330452, 0.1291032, 0.1071684, 0.130788, 0.1315224, 0.1290276, 0.112374, 0.1229364, 0.1164564, 0.1067472,
		0.0973296, 0.1063692, 0.1113696, 0.1134, 0.1072548, 0.1071468, 0.1067364, 0.10341, 0.1018548, 0.1024164, 0.1026864, 0.1031508,
		0.1073304, 0.1027296, 0.1050084, 0.1053108, 0.1085724, 0.1070928, 0.1043388, 0.1057428, 0.1089396, 0.1086588, 0.1130868, 0.1354536,
		0.1550124, 0.1317384, 0.1629828, 0.1820124, 0.1947672, 0.1940004, 0.1979424, 0.1877904, 0.1651752, 0.1537812, 0.1488456, 0.1431108,
		0.1401408, 0.1462644, 0.1393308, 0.1347192, 0.1256364, 0.1413612, 0.134514, 0.131058, 0.1218456, 0.1331748, 0.1271052, 0.122202,
		0.120906, 0.1274292, 0.1215, 0.1262736, 0.1297404, 0.1284228, 0.1321488, 0.1386936, 0.1504764, 0.131976, 0.1449684, 0.1613952,
		0.1638576, 0.1407888, 0.1499364, 0.1843236, 0.2065284, 0.1882656, 0.197478, 0.206982, 0.2207196, 0.2071116, 0.1917432, 0.1881144,
		0.181116, 0.1777464, 0.2019384, 0.1728648, 0.1840212, 0.1791828, 0.1757484, 0.1589976, 0.1474308, 0.1637064, 0.1515348, 0.1409508,
		0.1295028, 0.1464912, 0.134352, 0.1260252, 0.1126764, 0.141264, 0.1280016, 0.123228, 0.1157004, 0.1249884, 0.1173204, 0.111402,
		0.1006452, 0.117612, 0.11421, 0.111672, 0.1034316, 0.1073628, 0.1049112, 0.1028052, 0.1040796, 0.1021356, 0.103734, 0.10287,
		0.1031508, 0.1008828, 0.1029348, 0.1032372, 0.1086696, 0.1024164, 0.1059048, 0.1104732, 0.1126656, 0.100656, 0.1090584, 0.1141236,
		0.118854, 0.1128384, 0.1252044, 0.1452168, 0.177984, 0.148824, 0.1540188, 0.161622, 0.165078, 0.15741, 0.153522, 0.1504116,
		0.1471608, 0.1582524, 0.1461456, 0.1420308, 0.13203, 0.1500552, 0.1417716, 0.1361448, 0.1308852, 0.1393956, 0.1358964, 0.1342656,
		0.1341252, 0.1362852, 0.1359612, 0.1358316, 0.1363284, 0.1427976, 0.1374516, 0.1425384, 0.1428408, 0.133974, 0.1380456, 0.1467612,
		0.1669572, 0.1368792, 0.1460808, 0.1534032, 0.168588, 0.141426, 0.1486836, 0.1724112, 0.162108, 0.1635228, 0.1678104, 0.1620216,
		0.1640196, 0.1728108, 0.1932984, 0.1932876, 0.1829196, 0.1966032, 0.1795932, 0.1640736, 0.1486296, 0.163296, 0.1459728, 0.139968,
		0.1355184, 0.1376136, 0.1312956, 0.1247292, 0.120636, 0.1296864, 0.1358748, 0.1265868, 0.119178, 0.122958, 0.1219212, 0.1130112,
		0.1056564, 0.1217052, 0.1168668, 0.1047492, 0.1039176, 0.1188648, 0.1068552, 0.109836, 0.1091448, 0.107568, 0.1114236, 0.1101924,
		0.1056456, 0.1058616, 0.104868, 0.105408, 0.1078488, 0.1074924, 0.1135404, 0.1136484, 0.1146096, 0.1122552, 0.1197396, 0.1258848,
		0.1348488, 0.1292652, 0.1488024, 0.1612332, 0.1741176, 0.1596456, 0.1686312, 0.175662, 0.1813968, 0.1619892, 0.1513728, 0.1463292,
		0.1427652, 0.1576368, 0.1411236, 0.1379268, 0.1302696, 0.1453464, 0.13608, 0.1292436, 0.1245348, 0.1325484, 0.1266624, 0.126306,
		0.1191348, 0.124686, 0.119286, 0.121392, 0.121122, 0.1219428, 0.123984, 0.1293948, 0.13797, 0.12393, 0.1332936, 0.149688,
		0.1514916, 0.1421388, 0.1689984, 0.2102544, 0.2248776, 0.2155356, 0.2250936, 0.219294, 0.2164104, 0.2116368, 0.2038824, 0.1916892,
		0.1944972, 0.2180952, 0.208116, 0.2016252, 0.1947888, 0.2181816, 0.1901556, 0.1931904, 0.1782324, 0.18603, 0.175878, 0.1687716,
		0.1510164, 0.1707804, 0.1550124, 0.1386288, 0.1330236, 0.139482, 0.1357344, 0.1305288, 0.121014, 0.130086, 0.1217268, 0.1081728,
		0.1048788, 0.111672, 0.1064988, 0.1074816, 0.1097928, 0.110808, 0.1076112, 0.1057212, 0.1014336, 0.101034, 0.1067688, 0.103734,
		0.0997488, 0.095148, 0.1014876, 0.1033128, 0.0981828, 0.1021464, 0.1018116, 0.1002024, 0.1044684, 0.1026972, 0.1082376, 0.1219968,
		0.1253556, 0.1209816, 0.1308852, 0.150012, 0.1667736, 0.1638576, 0.159732, 0.1506708, 0.151794, 0.1515024, 0.148716, 0.145152,
		0.1404, 0.1476792, 0.1458648, 0.136998, 0.1256472, 0.139698, 0.1290276, 0.127278, 0.1230876, 0.1271808, 0.1272456, 0.12204,
		2(0.1241568), 0.1212516, 0.1214244, 0.120474, 0.1212624, 0.1214244, 0.12528, 0.1302372, 0.123282, 0.13851, 0.1412748, 0.1574964,
		0.1330992, 0.1466424, 0.1844208, 0.1922616, 0.1706076, 0.218376, 0.1946376, 0.1810836, 0.1483812, 0.152766, 0.1706616, 0.1571508,
		0.149796, 0.1481436, 0.1643328, 0.1562436, 0.1778328, 0.1602936, 0.1453788, 0.1442988, 0.1684368, 0.1463832, 0.1427004, 0.1294596,
		0.1316736, 0.1258632, 0.124362, 0.120096, 0.1303344, 0.1279152, 0.1220832, 0.1173636, 0.1260144, 0.1220076, 0.1100304, 0.0983016,
		0.1113264, 0.108216, 0.101952, 0.1005804, 0.1089504, 0.1038204, 0.0968976, 0.0965628, 0.0968976, 0.1020816, 0.0966708, 0.0952236,
		0.094662, 0.0942192, 0.0970488, 0.0994464, 0.0956772, 0.0961632, 0.0978696, 0.1019844, 0.0957528, 0.0944568, 0.0988848, 0.1089288,
		0.10206, 0.1045548, 0.1068336, 0.1159596, 0.110592, 0.1147608, 0.1161864, 0.1219428, 0.12015, 0.1223532, 0.1282068, 0.1311012,
		0.1269756, 0.1298376, 0.126846, 0.12555, 0.1267812, 0.1280772, 0.1246536, 0.1218672, 0.126306, 0.1233684, 0.1241676, 0.1235628,
		0.1218888, 0.1207224, 0.12474, 0.1276344, 0.123336, 0.1266408, 0.1341144, 0.1377432, 0.13014, 0.1379592, 0.1365768, 0.1382184,
		0.1322352, 0.1370304, 0.1428084, 0.1442124, 0.1361556, 0.14337, 0.1468368, 0.1468476, 0.1431864, 0.1403568, 0.1362852, 0.1344492,
		0.144774, 0.1347624, 0.1386288, 0.1306476, 0.1405512, 0.129762, 0.127656, 0.1270836, 0.1300752, 0.1292544, 0.1253772, 0.1155816,
		0.1311876, 0.1205712, 0.116424, 0.1130004, 0.1248804, 0.1158516, 0.1139076, 0.1060344, 0.1169856, 0.1047924, 0.097362, 0.0916272,
		0.1165752, 0.110268, 0.1060128, 0.0997056, 0.1105596, 0.0999972, 0.0960336, 0.0949644, 0.101412, 0.0980316, 0.0970056, 0.0989604,
		0.0970488, 0.1014336, 0.1011744, 0.0965628, 0.0972972, 0.096228, 0.0992088, 0.0977616, 0.0997596, 0.0986472, 0.099198, 0.0987336,
		0.0958716, 0.1016712, 0.1035396, 0.108054, 0.1034856, 0.1073952, 0.1110024, 0.113238, 0.1105704, 0.1146204, 0.11529, 0.1164672,
		0.119178, 0.1230876, 0.1200312, 0.1190484, 0.1252692, 0.1210464, 0.116802, 0.1129248, 0.1202256, 0.1197072, 0.1168128, 0.11583,
		0.1185408, 0.1161864, 0.1151928, 0.1153008, 0.1176876, 0.1171584, 0.11421, 0.1199232, 0.1154196, 0.1169856, 0.120366, 0.1336284,
		0.1172124, 0.1221372, 0.1232928, 0.1285416, 0.1200852, 0.12231, 0.1279476, 0.1352268, 0.1285524, 0.128952, 0.1280556, 0.13122,
		0.126198, 0.1266408, 0.1265976, 0.1313064, 0.127548, 0.1328724, 0.1278828, 0.1222452, 0.1289304, 0.127386, 0.1221372, 0.1165212,
		0.1317924, 0.1261332, 0.1197072, 0.1162944, 0.1195344, 0.1193832, 0.1090368, 0.1033992, 0.1119636, 0.105084, 0.1006344, 0.0912924,
		0.1035396, 0.09936, 0.0975456, 0.095472, 0.0957744, 0.0957852, 0.0966168, 0.0960012, 0.0974484, 0.0946404, 0.094284, 0.0926964,
		0.0895212, 0.0899748, 0.0911304, 0.0928692, 0.0922104, 0.0932256, 0.0921024, 0.0963144, 0.0897804, 0.098982, 0.1029888, 0.1134432,
		0.0953748, 0.1075356, 0.114642, 0.1264032, 0.1204308, 0.130356, 0.1384992, 0.1400976, 0.1411776, 0.1360152, 0.1407996, 0.1365984,
		0.1344816, 0.1633068, 0.1343844, 0.1316088, 0.1430136, 0.1317384, 0.1352376, 0.1260792, 0.131112, 0.1336176, 0.129708, 0.1306692,
		0.1317276, 0.1334016, 0.137052, 0.1350756, 0.138348, 0.128142, 0.1377216, 0.1487052, 0.1257984, 0.1318896, 0.1652076, 0.1415556,
		0.1518588, 0.1360044, 0.1348812, 0.1397088, 0.136026, 0.1420308, 0.1480572, 0.152172, 0.1405836, 0.140508, 0.1398276, 0.1569888,
		0.1364796, 0.1377108, 0.136566, 0.1451412, 0.1408428, 0.1435968, 0.136188, 0.1349676, 0.1388232, 0.130572, 0.1245456, 0.1185732,
		0.1368252, 0.1271808, 0.1110024, 0.1001268, 0.1222776, 0.116262, 0.102654, 0.0973296, 0.1116936, 0.0994032, 0.0918756, 0.0867348,
		0.0911196, 0.0897264, 0.086832, 0.0882144, 0.0908712, 0.0812592, 0.0859248, 0.0741204, 0.086508, 0.0905472, 0.0818856, 0.0763452,
		0.0863028, 0.0828036, 0.0771552, 0.0789048, 0.0879012, 0.0760644, 0.0816696, 0.0767124, 0.0754488, 0.0866376, 0.0908064, 0.1053108,
		0.0771984, 0.100548, 0.1142532, 0.1272348, 0.10287, 0.1115856, 0.126198, 0.1350864, 0.1278396, 0.1264464, 0.132732, 0.1280124,
		0.1280556, 0.1305504, 0.1257552, 0.1252908, 0.1315548, 0.1258632, 0.1251936, 0.12447, 0.1218888, 0.1232604, 0.1314036, 0.1224072,
		0.1249236, 0.11853, 0.1194804, 0.1240164, 0.1247076, 0.121014, 0.1200744, 0.12312, 0.1172016, 0.1234332, 0.1300644, 0.1328076,
		0.120474, 0.1331964, 0.1374084, 0.1399248, 0.1301184, 0.1410156, 0.1485972, 0.1500012, 0.1521072, 0.1468152, 0.1441044, 0.1339092,
		0.1364472, 0.1353024, 0.1343412, 0.1396116, 0.1454436, 0.1452492, 0.1334664, 0.1246428, 0.1432944, 0.13527, 0.1234656, 0.1106892,
		0.1297404, 0.1206576, 0.1063476, 0.0971568, 0.1182816, 0.1129248, 0.1080972, 0.0904932, 0.1144908, 0.1008828, 0.0915192, 0.0788724,
		0.1104516, 0.1013796, 0.0940356, 0.077328, 0.0963144, 0.0879552, 0.084078, 0.0766044, 0.0860328, 0.0911196, 0.0849096, 0.0848556,
		0.08397, 0.0833004, 0.0844992, 0.075114, 0.0719496, 0.076788, 0.0770472, 0.0850284, 0.0708048, 0.082782, 0.0914544, 0.0966708,
		0.0828576, 0.0847368, 0.0893808, 0.1018872, 0.0811944, 0.0920592, 0.107136, 0.124902, 0.0985932, 0.0993708, 0.1168668, 0.123876,
		0.1177524, 0.1141884, 0.1108404, 0.11394, 0.119826, 0.1207332, 0.1229904, 0.1133136, 0.12771, 0.12582, 0.123606, 0.1178712,
		0.122904, 0.1199232, 0.113508, 0.1130112, 0.1204848, 0.1177632, 0.1118772, 0.1163376, 0.108432, 0.1086156, 0.1146528, 0.1234116,
		0.0955152, 0.1149552, 0.123714, 0.130464, 0.1182276, 0.1309932, 0.1310904, 0.1184976, 0.1305936, 0.1265004, 0.119826, 0.1030536,
		0.1142856, 0.1025892, 0.0928476, 0.0885492, 0.0997272, 0.093096, 0.0896616, 0.0893052, 0.0963684, 0.0939384, 0.0913788, 0.084456,
		0.0977508, 0.095796, 0.0921996, 0.0843588, 0.103086, 0.0951264, 0.0825552, 0.0751896, 0.0796608, 0.0803412, 0.0732888, 0.0608364,
		0.0808812, 0.0749088, 0.0836784, 0.0852336, 0.0722412, 0.0750384, 0.0752976, 0.065178, 0.0755244, 0.0725004, 0.0758052, 0.0644652,
		0.0752436, 0.08019, 0.0832356, 0.0690768, 0.0690228, 0.0724248, 0.0699408, 0.075168, 0.0684072, 0.0788616, 0.0827172, 0.0876096,
		0.0715932, 0.0621864, 0.0753408, 0.080406, 0.0513972, 0.0875664, 0.0928152, 0.1004616, 0.086508, 0.087426, 0.090882, 0.0910656,
		0.0931176, 0.0915732, 0.0873072, 0.084078, 0.0862812, 0.0842292, 0.0865836, 0.0843048, 0.0868752, 0.0870912, 0.0831276, 0.0785376,
		0.0906768, 0.0865188, 0.0817236, 0.0757728, 0.0833652, 0.0827712, 0.084024, 0.09045, 0.0724464, 0.09396, 0.0994896, 0.1163376,
		0.0950724, 0.1043604, 0.1163052, 0.118908, 0.1077732, 0.1081836, 0.1160892, 0.1159812, 0.1095984, 0.1104084, 0.1168452, 0.111456,
		0.1125036, 0.111726, 0.1191888, 0.11286, 0.1141776, 0.1103976, 0.1128708, 0.1244268, 0.1247184, 0.1200636, 0.1158624, 0.1096632,
		0.124254, 0.114912, 0.1124496, 0.1125792, 0.1295784, 0.1169964, 0.1073196, 0.1005048, 0.1202148, 0.1040148, 0.0977724, 0.0950508,
		0.114966, 0.1079568, 0.0987768, 0.0977724, 0.1033128, 0.098658, 0.0979992, 0.0933768, 0.0979992, 0.0933012, 0.091422, 0.0882792,
		0.0918, 0.089748, 0.089046, 0.0892728, 0.0871668, 0.0893592, 0.0907632, 0.0924156, 0.0885708, 0.0887544, 0.0909036, 0.094392,
		0.0872964, 0.0878904, 0.095202, 0.097794, 0.0979776, 0.0996408, 0.1039284, 0.1092744, 0.102654, 0.1053756, 0.1109592, 0.110538,
		0.1123632, 0.1124496, 0.102384, 0.0920484, 0.10368, 0.0985176, 0.093852, 0.0895104, 0.09612, 0.0921024, 0.0904068, 0.0885384,
		0.0897588, 0.08856, 0.0883764, 0.0888948, 0.0864, 0.0871344, 0.0932904, 0.093204, 0.0811404, 0.0934524, 0.1029564, 0.1287144,
		0.0994464, 0.1198584, 0.1297296, 0.1352052, 0.1227096, 0.1297512, 0.1309716, 0.1330884, 0.1317708, 0.1339092, 0.1338984, 0.131112,
		0.1308204, 0.1285524, 0.1288116, 0.1239516, 0.1290276, 0.1270944, 0.1274832, 0.1252692, 0.1337148, 0.1286496, 0.1216188, 0.1151388,
		0.1304856, 0.1270836, 0.1195128, 0.1125252, 0.1301616, 0.1246968, 0.114156, 0.1042092, 0.1212408, 0.1134756, 0.1022652, 0.0953316,
		0.1120932, 0.1076112, 0.1020384, 0.097632, 0.111672, 0.0987336, 0.0958608, 0.0913788, 0.0956988, 0.0926748, 0.0911088, 0.0880308,
		0.0929016, 0.0909684, 0.090126, 0.0878472, 0.0922644, 0.0925236, 0.0919728, 0.0917028, 0.0867672, 0.0894132, 0.0909792, 0.0974808,
		0.0846504, 0.0938736, 0.1001808, 0.1088208, 0.1030212, 0.1068012, 0.1141128, 0.1163916, 0.115344, 0.1150416, 0.1141776, 0.103464,
		0.1188432, 0.1129572, 0.0948672, 0.080892, 0.1111536, 0.0838728, 0.076842, 0.0748116, 0.084564, 0.083808, 0.0818316, 0.0772308,
		0.0845964, 0.0769392, 0.0803844, 0.0810756, 0.0774684, 0.08289, 0.0891216, 0.0980856, 0.07479, 0.0935928, 0.1106784, 0.1210032,
		0.0967572, 0.1107972, 0.1196748, 0.1481328, 0.117666, 0.1263816, 0.136296, 0.132192, 0.134352, 0.1305828, 0.125604, 0.1274292,
		0.1385316, 0.1316304, 0.1233252, 0.1255392, 0.138348, 0.1344276, 0.1245672, 0.1252908, 0.1529712, 0.1356372, 0.11664, 0.1064232,
		0.1187244, 0.1121796, 0.1096416, 0.1037988, 0.1181628, 0.1129896, 0.1043604, 0.10125, 0.1126548, 0.1040364, 0.0987012, 0.092664,
		0.114912, 0.1037124, 0.0945756, 0.0862812, 0.0985176, 0.0923832, 0.0934416, 0.092286, 0.0948996, 0.0903852, 0.090612, 0.090882,
		0.0902664, 0.088614, 0.0905904, 0.0905796, 0.0890892, 0.090018, 0.0906012, 0.0933552, 0.090828, 0.0918432, 0.0934848, 0.100116,
		0.0890028, 0.0931932, 0.0980208, 0.1053864, 0.0986364, 0.1008504, 0.1058184, 0.1129356, 0.1022976, 0.1074276, 0.109458, 0.1082916,
		0.10287, 0.0970704, 0.0918108, 0.0806868, 0.109296, 0.0973836, 0.0904932, 0.0875016, 0.0860436, 0.0846936, 0.084618, 0.0810756,
		0.0895644, 0.0850392, 0.085914, 0.0854172, 0.082728, 0.0839376, 0.0882792, 0.0923724, 0.0869184, 0.0888948, 0.0951912, 0.1067472,
		0.095256, 0.1051488, 0.122904, 0.11934, 0.1127412, 0.1219536, 0.1253772, 0.12663, 0.1227096, 0.1254636, 0.1246752, 0.124254,
		0.133056, 0.1267272, 0.1234764, 0.1164024, 0.1261008, 0.1196748, 0.1164996, 0.1142208, 0.1171152, 0.11556, 0.1119528, 0.1090152,
		0.1091664, 0.1080108, 0.1069632, 0.1036584, 0.1080108, 0.106596, 0.1060776, 0.103896, 0.1055592, 0.1013364, 0.097686, 0.0906336,
		0.1109808, 0.1022652, 0.0918108, 0.0853956, 0.1004076, 0.0906228, 0.0934524, 0.0928692, 0.0970812, 0.0921024, 0.0879984, 0.0894132,
		0.0911304, 0.08856, 0.087534, 0.0878364, 0.088344, 0.0881928, 0.0915732, 0.095148, 0.0914436, 0.09612, 0.09936, 0.1053,
		0.0946512, 0.1027836, 0.105084, 0.1136376, 0.1197288, 0.114318, 0.1151496, 0.1185516, 0.1287144, 0.1229364, 0.1215, 0.1188,
		0.129654, 0.1212408, 0.1180332, 0.107352, 0.1164564, 0.112266, 0.1027944, 0.0917028, 0.102978, 0.0913464, 0.0985284, 0.09504,
		0.0954612, 0.0940032, 0.0954612, 0.0956556, 0.094338, 0.0955476, 0.0948564, 0.0985284, 0.0976104, 0.1018116, 0.1118556, 0.1309932,
		0.1047708, 0.1141884, 0.13446, 0.1458756, 0.1330668, 0.1479924, 0.1526796, 0.1511892, 0.1472364, 0.1396548, 0.1359936, 0.1395576,
		0.1473012, 0.1417284, 0.1366524, 0.1383372, 0.151578, 0.141696, 0.148662, 0.1277316, 0.1466964, 0.1297836, 0.120096, 0.1032912,
		0.1374624, 0.1176552, 0.1185516, 0.1006344, 0.1325484, 0.1098792, 0.1048572, 0.0992304, 0.1022328, 0.095904, 0.0925452, 0.0851688,
		0.096876, 0.0899964, 0.0856872, 0.081378, 0.0873828, 0.084078, 0.0837216, 0.084402, 0.08775, 0.087318, 0.0838296, 0.0829548,
		0.0834516, 0.0823176, 0.0788724, 0.0771336, 0.08613, 0.0840456, 0.0823284, 0.0776952, 0.0859032, 0.0895968, 0.0842292, 0.0879012,
		0.0802332, 0.090126, 0.0966276, 0.108918, 0.1006992, 0.1030968, 0.104328, 0.1025676, 0.1006344, 0.10692, 0.102978, 0.0993384,
		0.112968, 0.1078596, 0.101034, 0.085914, 0.1044684, 0.0932472, 0.0876312, 0.0853956, 0.087912, 0.0866484, 0.08532, 0.0830412,
		0.0852876, 0.0831492, 0.0821988, 0.078354, 0.0786564, 0.0807408, 0.081162, 0.09261, 0.0774252, 0.0949104, 0.1031616, 0.1157004,
		0.0998892, 0.1065312, 0.1226556, 0.1292976, 0.1139076, 0.1190268, 0.1188432, 0.1343304, 0.1219428, 0.1259928, 0.1201284, 0.123282,
		0.1260684, 0.1226772, 0.1173096, 0.1175688, 0.1202148, 0.11961, 0.1176552, 0.1184652, 0.118422, 0.116856, 0.1125252, 0.1044144,
		0.1141884, 0.104598, 0.1036584, 0.0968544, 0.1196208, 0.1036044, 0.0975888, 0.0919512, 0.1024488, 0.095526, 0.0887652, 0.0841104,
		0.1024596, 0.0975348, 0.0930852, 0.089316, 0.0973188, 0.0901584, 0.0896724, 0.0891324, 0.0902232, 0.0875448, 0.0857412, 0.08316,
		0.0864, 0.0822852, 0.0810324, 0.081108, 0.0803628, 0.0810108, 0.0806868, 0.081648, 0.081054, 0.0816696, 0.084348, 0.0871992,
		0.0840456, 0.0889488, 0.0895536, 0.0914436, 0.0915624, 0.0926208, 0.0950832, 0.0996948, 0.1024812, 0.1062612, 0.1048572, 0.1046628,
		0.1125144, 0.108378, 0.1021464, 0.091962, 0.1061964, 0.0970056, 0.0942192, 0.0893592, 0.0949644, 0.0906444, 0.0886248, 0.0864,
		0.089964, 2(0.08856), 0.0916812, 0.089748, 0.0908712, 0.0918, 0.0955152, 0.091638, 0.0991764, 0.1033992, 0.1314468, 0.1032804,
		0.1145556, 0.1264896, 0.1613628, 0.127602, 0.1378296, 0.1505196, 0.1558764, 0.1457028, 0.137214, 0.1372572, 0.1400544, 0.16605,
		0.138996, 0.1304316, 0.1215972, 0.1351728, 0.1253124, 0.127494, 0.1095336, 0.1385964, 0.1216188, 0.1092852, 0.1002996, 0.1314468,
		0.12042, 0.1075572, 0.1005156, 0.1284228, 0.1216836, 0.1081944, 0.0970812, 0.108432, 0.09774, 0.0920808, 0.0857952
	];
END_VAR
